(* IEC 61131-3 sources: STAR-PLC-Agent/results/raw/batch_fresh_20261114/PUB009/functional/attempt_0001, 1 file *)

(* ---- test_program.st ---- *)
PROGRAM PLC_PRG
VAR
 BenchStep : UDINT := 0;
 BenchCalls : UDINT := 0;
 BenchDone : BOOL := FALSE;
 BenchUut0 : FB_Task;
 BenchUut1 : FB_Task;
 BenchUut2 : FB_Task;
 BenchUut3 : FB_Task;
 BenchUut4 : FB_Task;
 BenchUut5 : FB_Task;
 BenchUut6 : FB_Task;
 TraceIn_cyclicExecution : ARRAY[0..454] OF BOOL;
 TraceIn_trigger : ARRAY[0..454] OF BOOL;
 TraceIn_value : ARRAY[0..454] OF LREAL;
 TraceIn_windowSize : ARRAY[0..454] OF INT;
 TraceIn_reset : ARRAY[0..454] OF BOOL;
 TraceOut_average : ARRAY[0..454] OF LREAL;
 TraceOut_windowSizeReached : ARRAY[0..454] OF BOOL;
 TraceOut_error : ARRAY[0..454] OF BOOL;
 TraceOut_status : ARRAY[0..454] OF WORD;
END_VAR

IF NOT BenchDone THEN
 CASE BenchStep OF
 0:
   BenchUut0.cyclicExecution := TRUE;
   BenchUut0.trigger := FALSE;
   BenchUut0.value := LREAL#3.0;
   BenchUut0.windowSize := INT#3;
   BenchUut0.reset := FALSE;
   TraceIn_cyclicExecution[0] := BenchUut0.cyclicExecution;
   TraceIn_trigger[0] := BenchUut0.trigger;
   TraceIn_value[0] := BenchUut0.value;
   TraceIn_windowSize[0] := BenchUut0.windowSize;
   TraceIn_reset[0] := BenchUut0.reset;
   BenchUut0();
   TraceOut_average[0] := BenchUut0.average;
   TraceOut_windowSizeReached[0] := BenchUut0.windowSizeReached;
   TraceOut_error[0] := BenchUut0.error;
   TraceOut_status[0] := BenchUut0.status;
   BenchCalls := BenchCalls + 1;
 1:
   BenchUut0.cyclicExecution := TRUE;
   BenchUut0.trigger := FALSE;
   BenchUut0.value := LREAL#6.0;
   BenchUut0.windowSize := INT#3;
   BenchUut0.reset := FALSE;
   TraceIn_cyclicExecution[1] := BenchUut0.cyclicExecution;
   TraceIn_trigger[1] := BenchUut0.trigger;
   TraceIn_value[1] := BenchUut0.value;
   TraceIn_windowSize[1] := BenchUut0.windowSize;
   TraceIn_reset[1] := BenchUut0.reset;
   BenchUut0();
   TraceOut_average[1] := BenchUut0.average;
   TraceOut_windowSizeReached[1] := BenchUut0.windowSizeReached;
   TraceOut_error[1] := BenchUut0.error;
   TraceOut_status[1] := BenchUut0.status;
   BenchCalls := BenchCalls + 1;
 2:
   BenchUut0.cyclicExecution := TRUE;
   BenchUut0.trigger := FALSE;
   BenchUut0.value := LREAL#9.0;
   BenchUut0.windowSize := INT#3;
   BenchUut0.reset := FALSE;
   TraceIn_cyclicExecution[2] := BenchUut0.cyclicExecution;
   TraceIn_trigger[2] := BenchUut0.trigger;
   TraceIn_value[2] := BenchUut0.value;
   TraceIn_windowSize[2] := BenchUut0.windowSize;
   TraceIn_reset[2] := BenchUut0.reset;
   BenchUut0();
   TraceOut_average[2] := BenchUut0.average;
   TraceOut_windowSizeReached[2] := BenchUut0.windowSizeReached;
   TraceOut_error[2] := BenchUut0.error;
   TraceOut_status[2] := BenchUut0.status;
   BenchCalls := BenchCalls + 1;
 3:
   BenchUut0.cyclicExecution := TRUE;
   BenchUut0.trigger := TRUE;
   BenchUut0.value := LREAL#12.0;
   BenchUut0.windowSize := INT#3;
   BenchUut0.reset := FALSE;
   TraceIn_cyclicExecution[3] := BenchUut0.cyclicExecution;
   TraceIn_trigger[3] := BenchUut0.trigger;
   TraceIn_value[3] := BenchUut0.value;
   TraceIn_windowSize[3] := BenchUut0.windowSize;
   TraceIn_reset[3] := BenchUut0.reset;
   BenchUut0();
   TraceOut_average[3] := BenchUut0.average;
   TraceOut_windowSizeReached[3] := BenchUut0.windowSizeReached;
   TraceOut_error[3] := BenchUut0.error;
   TraceOut_status[3] := BenchUut0.status;
   BenchCalls := BenchCalls + 1;
 4:
   BenchUut0.cyclicExecution := TRUE;
   BenchUut0.trigger := FALSE;
   BenchUut0.value := LREAL#99.0;
   BenchUut0.windowSize := INT#3;
   BenchUut0.reset := TRUE;
   TraceIn_cyclicExecution[4] := BenchUut0.cyclicExecution;
   TraceIn_trigger[4] := BenchUut0.trigger;
   TraceIn_value[4] := BenchUut0.value;
   TraceIn_windowSize[4] := BenchUut0.windowSize;
   TraceIn_reset[4] := BenchUut0.reset;
   BenchUut0();
   TraceOut_average[4] := BenchUut0.average;
   TraceOut_windowSizeReached[4] := BenchUut0.windowSizeReached;
   TraceOut_error[4] := BenchUut0.error;
   TraceOut_status[4] := BenchUut0.status;
   BenchCalls := BenchCalls + 1;
 5:
   BenchUut0.cyclicExecution := TRUE;
   BenchUut0.trigger := FALSE;
   BenchUut0.value := LREAL#-6.0;
   BenchUut0.windowSize := INT#3;
   BenchUut0.reset := FALSE;
   TraceIn_cyclicExecution[5] := BenchUut0.cyclicExecution;
   TraceIn_trigger[5] := BenchUut0.trigger;
   TraceIn_value[5] := BenchUut0.value;
   TraceIn_windowSize[5] := BenchUut0.windowSize;
   TraceIn_reset[5] := BenchUut0.reset;
   BenchUut0();
   TraceOut_average[5] := BenchUut0.average;
   TraceOut_windowSizeReached[5] := BenchUut0.windowSizeReached;
   TraceOut_error[5] := BenchUut0.error;
   TraceOut_status[5] := BenchUut0.status;
   BenchCalls := BenchCalls + 1;
 6:
   BenchUut1.cyclicExecution := FALSE;
   BenchUut1.trigger := TRUE;
   BenchUut1.value := LREAL#2.0;
   BenchUut1.windowSize := INT#3;
   BenchUut1.reset := FALSE;
   TraceIn_cyclicExecution[6] := BenchUut1.cyclicExecution;
   TraceIn_trigger[6] := BenchUut1.trigger;
   TraceIn_value[6] := BenchUut1.value;
   TraceIn_windowSize[6] := BenchUut1.windowSize;
   TraceIn_reset[6] := BenchUut1.reset;
   BenchUut1();
   TraceOut_average[6] := BenchUut1.average;
   TraceOut_windowSizeReached[6] := BenchUut1.windowSizeReached;
   TraceOut_error[6] := BenchUut1.error;
   TraceOut_status[6] := BenchUut1.status;
   BenchCalls := BenchCalls + 1;
 7:
   BenchUut1.cyclicExecution := FALSE;
   BenchUut1.trigger := TRUE;
   BenchUut1.value := LREAL#100.0;
   BenchUut1.windowSize := INT#3;
   BenchUut1.reset := FALSE;
   TraceIn_cyclicExecution[7] := BenchUut1.cyclicExecution;
   TraceIn_trigger[7] := BenchUut1.trigger;
   TraceIn_value[7] := BenchUut1.value;
   TraceIn_windowSize[7] := BenchUut1.windowSize;
   TraceIn_reset[7] := BenchUut1.reset;
   BenchUut1();
   TraceOut_average[7] := BenchUut1.average;
   TraceOut_windowSizeReached[7] := BenchUut1.windowSizeReached;
   TraceOut_error[7] := BenchUut1.error;
   TraceOut_status[7] := BenchUut1.status;
   BenchCalls := BenchCalls + 1;
 8:
   BenchUut1.cyclicExecution := FALSE;
   BenchUut1.trigger := FALSE;
   BenchUut1.value := LREAL#100.0;
   BenchUut1.windowSize := INT#3;
   BenchUut1.reset := FALSE;
   TraceIn_cyclicExecution[8] := BenchUut1.cyclicExecution;
   TraceIn_trigger[8] := BenchUut1.trigger;
   TraceIn_value[8] := BenchUut1.value;
   TraceIn_windowSize[8] := BenchUut1.windowSize;
   TraceIn_reset[8] := BenchUut1.reset;
   BenchUut1();
   TraceOut_average[8] := BenchUut1.average;
   TraceOut_windowSizeReached[8] := BenchUut1.windowSizeReached;
   TraceOut_error[8] := BenchUut1.error;
   TraceOut_status[8] := BenchUut1.status;
   BenchCalls := BenchCalls + 1;
 9:
   BenchUut1.cyclicExecution := FALSE;
   BenchUut1.trigger := TRUE;
   BenchUut1.value := LREAL#4.0;
   BenchUut1.windowSize := INT#3;
   BenchUut1.reset := FALSE;
   TraceIn_cyclicExecution[9] := BenchUut1.cyclicExecution;
   TraceIn_trigger[9] := BenchUut1.trigger;
   TraceIn_value[9] := BenchUut1.value;
   TraceIn_windowSize[9] := BenchUut1.windowSize;
   TraceIn_reset[9] := BenchUut1.reset;
   BenchUut1();
   TraceOut_average[9] := BenchUut1.average;
   TraceOut_windowSizeReached[9] := BenchUut1.windowSizeReached;
   TraceOut_error[9] := BenchUut1.error;
   TraceOut_status[9] := BenchUut1.status;
   BenchCalls := BenchCalls + 1;
 10:
   BenchUut1.cyclicExecution := TRUE;
   BenchUut1.trigger := FALSE;
   BenchUut1.value := LREAL#8.0;
   BenchUut1.windowSize := INT#1;
   BenchUut1.reset := FALSE;
   TraceIn_cyclicExecution[10] := BenchUut1.cyclicExecution;
   TraceIn_trigger[10] := BenchUut1.trigger;
   TraceIn_value[10] := BenchUut1.value;
   TraceIn_windowSize[10] := BenchUut1.windowSize;
   TraceIn_reset[10] := BenchUut1.reset;
   BenchUut1();
   TraceOut_average[10] := BenchUut1.average;
   TraceOut_windowSizeReached[10] := BenchUut1.windowSizeReached;
   TraceOut_error[10] := BenchUut1.error;
   TraceOut_status[10] := BenchUut1.status;
   BenchCalls := BenchCalls + 1;
 11:
   BenchUut1.cyclicExecution := FALSE;
   BenchUut1.trigger := FALSE;
   BenchUut1.value := LREAL#0.0;
   BenchUut1.windowSize := INT#0;
   BenchUut1.reset := FALSE;
   TraceIn_cyclicExecution[11] := BenchUut1.cyclicExecution;
   TraceIn_trigger[11] := BenchUut1.trigger;
   TraceIn_value[11] := BenchUut1.value;
   TraceIn_windowSize[11] := BenchUut1.windowSize;
   TraceIn_reset[11] := BenchUut1.reset;
   BenchUut1();
   TraceOut_average[11] := BenchUut1.average;
   TraceOut_windowSizeReached[11] := BenchUut1.windowSizeReached;
   TraceOut_error[11] := BenchUut1.error;
   TraceOut_status[11] := BenchUut1.status;
   BenchCalls := BenchCalls + 1;
 12:
   BenchUut1.cyclicExecution := FALSE;
   BenchUut1.trigger := FALSE;
   BenchUut1.value := LREAL#0.0;
   BenchUut1.windowSize := INT#101;
   BenchUut1.reset := FALSE;
   TraceIn_cyclicExecution[12] := BenchUut1.cyclicExecution;
   TraceIn_trigger[12] := BenchUut1.trigger;
   TraceIn_value[12] := BenchUut1.value;
   TraceIn_windowSize[12] := BenchUut1.windowSize;
   TraceIn_reset[12] := BenchUut1.reset;
   BenchUut1();
   TraceOut_average[12] := BenchUut1.average;
   TraceOut_windowSizeReached[12] := BenchUut1.windowSizeReached;
   TraceOut_error[12] := BenchUut1.error;
   TraceOut_status[12] := BenchUut1.status;
   BenchCalls := BenchCalls + 1;
 13:
   BenchUut1.cyclicExecution := FALSE;
   BenchUut1.trigger := FALSE;
   BenchUut1.value := LREAL#0.0;
   BenchUut1.windowSize := INT#1;
   BenchUut1.reset := TRUE;
   TraceIn_cyclicExecution[13] := BenchUut1.cyclicExecution;
   TraceIn_trigger[13] := BenchUut1.trigger;
   TraceIn_value[13] := BenchUut1.value;
   TraceIn_windowSize[13] := BenchUut1.windowSize;
   TraceIn_reset[13] := BenchUut1.reset;
   BenchUut1();
   TraceOut_average[13] := BenchUut1.average;
   TraceOut_windowSizeReached[13] := BenchUut1.windowSizeReached;
   TraceOut_error[13] := BenchUut1.error;
   TraceOut_status[13] := BenchUut1.status;
   BenchCalls := BenchCalls + 1;
 14:
   BenchUut1.cyclicExecution := FALSE;
   BenchUut1.trigger := TRUE;
   BenchUut1.value := LREAL#5.0;
   BenchUut1.windowSize := INT#1;
   BenchUut1.reset := FALSE;
   TraceIn_cyclicExecution[14] := BenchUut1.cyclicExecution;
   TraceIn_trigger[14] := BenchUut1.trigger;
   TraceIn_value[14] := BenchUut1.value;
   TraceIn_windowSize[14] := BenchUut1.windowSize;
   TraceIn_reset[14] := BenchUut1.reset;
   BenchUut1();
   TraceOut_average[14] := BenchUut1.average;
   TraceOut_windowSizeReached[14] := BenchUut1.windowSizeReached;
   TraceOut_error[14] := BenchUut1.error;
   TraceOut_status[14] := BenchUut1.status;
   BenchCalls := BenchCalls + 1;
 15:
   BenchUut2.cyclicExecution := FALSE;
   BenchUut2.trigger := TRUE;
   BenchUut2.value := LREAL#8.0;
   BenchUut2.windowSize := INT#2;
   BenchUut2.reset := FALSE;
   TraceIn_cyclicExecution[15] := BenchUut2.cyclicExecution;
   TraceIn_trigger[15] := BenchUut2.trigger;
   TraceIn_value[15] := BenchUut2.value;
   TraceIn_windowSize[15] := BenchUut2.windowSize;
   TraceIn_reset[15] := BenchUut2.reset;
   BenchUut2();
   TraceOut_average[15] := BenchUut2.average;
   TraceOut_windowSizeReached[15] := BenchUut2.windowSizeReached;
   TraceOut_error[15] := BenchUut2.error;
   TraceOut_status[15] := BenchUut2.status;
   BenchCalls := BenchCalls + 1;
 16:
   BenchUut2.cyclicExecution := FALSE;
   BenchUut2.trigger := FALSE;
   BenchUut2.value := LREAL#8.0;
   BenchUut2.windowSize := INT#2;
   BenchUut2.reset := FALSE;
   TraceIn_cyclicExecution[16] := BenchUut2.cyclicExecution;
   TraceIn_trigger[16] := BenchUut2.trigger;
   TraceIn_value[16] := BenchUut2.value;
   TraceIn_windowSize[16] := BenchUut2.windowSize;
   TraceIn_reset[16] := BenchUut2.reset;
   BenchUut2();
   TraceOut_average[16] := BenchUut2.average;
   TraceOut_windowSizeReached[16] := BenchUut2.windowSizeReached;
   TraceOut_error[16] := BenchUut2.error;
   TraceOut_status[16] := BenchUut2.status;
   BenchCalls := BenchCalls + 1;
 17:
   BenchUut2.cyclicExecution := FALSE;
   BenchUut2.trigger := TRUE;
   BenchUut2.value := LREAL#99.0;
   BenchUut2.windowSize := INT#0;
   BenchUut2.reset := FALSE;
   TraceIn_cyclicExecution[17] := BenchUut2.cyclicExecution;
   TraceIn_trigger[17] := BenchUut2.trigger;
   TraceIn_value[17] := BenchUut2.value;
   TraceIn_windowSize[17] := BenchUut2.windowSize;
   TraceIn_reset[17] := BenchUut2.reset;
   BenchUut2();
   TraceOut_average[17] := BenchUut2.average;
   TraceOut_windowSizeReached[17] := BenchUut2.windowSizeReached;
   TraceOut_error[17] := BenchUut2.error;
   TraceOut_status[17] := BenchUut2.status;
   BenchCalls := BenchCalls + 1;
 18:
   BenchUut2.cyclicExecution := FALSE;
   BenchUut2.trigger := TRUE;
   BenchUut2.value := LREAL#100.0;
   BenchUut2.windowSize := INT#2;
   BenchUut2.reset := FALSE;
   TraceIn_cyclicExecution[18] := BenchUut2.cyclicExecution;
   TraceIn_trigger[18] := BenchUut2.trigger;
   TraceIn_value[18] := BenchUut2.value;
   TraceIn_windowSize[18] := BenchUut2.windowSize;
   TraceIn_reset[18] := BenchUut2.reset;
   BenchUut2();
   TraceOut_average[18] := BenchUut2.average;
   TraceOut_windowSizeReached[18] := BenchUut2.windowSizeReached;
   TraceOut_error[18] := BenchUut2.error;
   TraceOut_status[18] := BenchUut2.status;
   BenchCalls := BenchCalls + 1;
 19:
   BenchUut2.cyclicExecution := FALSE;
   BenchUut2.trigger := FALSE;
   BenchUut2.value := LREAL#8.0;
   BenchUut2.windowSize := INT#2;
   BenchUut2.reset := FALSE;
   TraceIn_cyclicExecution[19] := BenchUut2.cyclicExecution;
   TraceIn_trigger[19] := BenchUut2.trigger;
   TraceIn_value[19] := BenchUut2.value;
   TraceIn_windowSize[19] := BenchUut2.windowSize;
   TraceIn_reset[19] := BenchUut2.reset;
   BenchUut2();
   TraceOut_average[19] := BenchUut2.average;
   TraceOut_windowSizeReached[19] := BenchUut2.windowSizeReached;
   TraceOut_error[19] := BenchUut2.error;
   TraceOut_status[19] := BenchUut2.status;
   BenchCalls := BenchCalls + 1;
 20:
   BenchUut2.cyclicExecution := FALSE;
   BenchUut2.trigger := TRUE;
   BenchUut2.value := LREAL#4.0;
   BenchUut2.windowSize := INT#2;
   BenchUut2.reset := FALSE;
   TraceIn_cyclicExecution[20] := BenchUut2.cyclicExecution;
   TraceIn_trigger[20] := BenchUut2.trigger;
   TraceIn_value[20] := BenchUut2.value;
   TraceIn_windowSize[20] := BenchUut2.windowSize;
   TraceIn_reset[20] := BenchUut2.reset;
   BenchUut2();
   TraceOut_average[20] := BenchUut2.average;
   TraceOut_windowSizeReached[20] := BenchUut2.windowSizeReached;
   TraceOut_error[20] := BenchUut2.error;
   TraceOut_status[20] := BenchUut2.status;
   BenchCalls := BenchCalls + 1;
 21:
   BenchUut2.cyclicExecution := FALSE;
   BenchUut2.trigger := FALSE;
   BenchUut2.value := LREAL#8.0;
   BenchUut2.windowSize := INT#3;
   BenchUut2.reset := FALSE;
   TraceIn_cyclicExecution[21] := BenchUut2.cyclicExecution;
   TraceIn_trigger[21] := BenchUut2.trigger;
   TraceIn_value[21] := BenchUut2.value;
   TraceIn_windowSize[21] := BenchUut2.windowSize;
   TraceIn_reset[21] := BenchUut2.reset;
   BenchUut2();
   TraceOut_average[21] := BenchUut2.average;
   TraceOut_windowSizeReached[21] := BenchUut2.windowSizeReached;
   TraceOut_error[21] := BenchUut2.error;
   TraceOut_status[21] := BenchUut2.status;
   BenchCalls := BenchCalls + 1;
 22:
   BenchUut3.cyclicExecution := TRUE;
   BenchUut3.trigger := FALSE;
   BenchUut3.value := LREAL#10.0;
   BenchUut3.windowSize := INT#2;
   BenchUut3.reset := FALSE;
   TraceIn_cyclicExecution[22] := BenchUut3.cyclicExecution;
   TraceIn_trigger[22] := BenchUut3.trigger;
   TraceIn_value[22] := BenchUut3.value;
   TraceIn_windowSize[22] := BenchUut3.windowSize;
   TraceIn_reset[22] := BenchUut3.reset;
   BenchUut3();
   TraceOut_average[22] := BenchUut3.average;
   TraceOut_windowSizeReached[22] := BenchUut3.windowSizeReached;
   TraceOut_error[22] := BenchUut3.error;
   TraceOut_status[22] := BenchUut3.status;
   BenchCalls := BenchCalls + 1;
 23:
   BenchUut3.cyclicExecution := TRUE;
   BenchUut3.trigger := FALSE;
   BenchUut3.value := LREAL#20.0;
   BenchUut3.windowSize := INT#2;
   BenchUut3.reset := FALSE;
   TraceIn_cyclicExecution[23] := BenchUut3.cyclicExecution;
   TraceIn_trigger[23] := BenchUut3.trigger;
   TraceIn_value[23] := BenchUut3.value;
   TraceIn_windowSize[23] := BenchUut3.windowSize;
   TraceIn_reset[23] := BenchUut3.reset;
   BenchUut3();
   TraceOut_average[23] := BenchUut3.average;
   TraceOut_windowSizeReached[23] := BenchUut3.windowSizeReached;
   TraceOut_error[23] := BenchUut3.error;
   TraceOut_status[23] := BenchUut3.status;
   BenchCalls := BenchCalls + 1;
 24:
   BenchUut3.cyclicExecution := TRUE;
   BenchUut3.trigger := FALSE;
   BenchUut3.value := LREAL#99.0;
   BenchUut3.windowSize := INT#0;
   BenchUut3.reset := TRUE;
   TraceIn_cyclicExecution[24] := BenchUut3.cyclicExecution;
   TraceIn_trigger[24] := BenchUut3.trigger;
   TraceIn_value[24] := BenchUut3.value;
   TraceIn_windowSize[24] := BenchUut3.windowSize;
   TraceIn_reset[24] := BenchUut3.reset;
   BenchUut3();
   TraceOut_average[24] := BenchUut3.average;
   TraceOut_windowSizeReached[24] := BenchUut3.windowSizeReached;
   TraceOut_error[24] := BenchUut3.error;
   TraceOut_status[24] := BenchUut3.status;
   BenchCalls := BenchCalls + 1;
 25:
   BenchUut3.cyclicExecution := TRUE;
   BenchUut3.trigger := FALSE;
   BenchUut3.value := LREAL#99.0;
   BenchUut3.windowSize := INT#-3;
   BenchUut3.reset := FALSE;
   TraceIn_cyclicExecution[25] := BenchUut3.cyclicExecution;
   TraceIn_trigger[25] := BenchUut3.trigger;
   TraceIn_value[25] := BenchUut3.value;
   TraceIn_windowSize[25] := BenchUut3.windowSize;
   TraceIn_reset[25] := BenchUut3.reset;
   BenchUut3();
   TraceOut_average[25] := BenchUut3.average;
   TraceOut_windowSizeReached[25] := BenchUut3.windowSizeReached;
   TraceOut_error[25] := BenchUut3.error;
   TraceOut_status[25] := BenchUut3.status;
   BenchCalls := BenchCalls + 1;
 26:
   BenchUut3.cyclicExecution := TRUE;
   BenchUut3.trigger := FALSE;
   BenchUut3.value := LREAL#30.0;
   BenchUut3.windowSize := INT#3;
   BenchUut3.reset := FALSE;
   TraceIn_cyclicExecution[26] := BenchUut3.cyclicExecution;
   TraceIn_trigger[26] := BenchUut3.trigger;
   TraceIn_value[26] := BenchUut3.value;
   TraceIn_windowSize[26] := BenchUut3.windowSize;
   TraceIn_reset[26] := BenchUut3.reset;
   BenchUut3();
   TraceOut_average[26] := BenchUut3.average;
   TraceOut_windowSizeReached[26] := BenchUut3.windowSizeReached;
   TraceOut_error[26] := BenchUut3.error;
   TraceOut_status[26] := BenchUut3.status;
   BenchCalls := BenchCalls + 1;
 27:
   BenchUut3.cyclicExecution := FALSE;
   BenchUut3.trigger := TRUE;
   BenchUut3.value := LREAL#60.0;
   BenchUut3.windowSize := INT#3;
   BenchUut3.reset := FALSE;
   TraceIn_cyclicExecution[27] := BenchUut3.cyclicExecution;
   TraceIn_trigger[27] := BenchUut3.trigger;
   TraceIn_value[27] := BenchUut3.value;
   TraceIn_windowSize[27] := BenchUut3.windowSize;
   TraceIn_reset[27] := BenchUut3.reset;
   BenchUut3();
   TraceOut_average[27] := BenchUut3.average;
   TraceOut_windowSizeReached[27] := BenchUut3.windowSizeReached;
   TraceOut_error[27] := BenchUut3.error;
   TraceOut_status[27] := BenchUut3.status;
   BenchCalls := BenchCalls + 1;
 28:
   BenchUut3.cyclicExecution := FALSE;
   BenchUut3.trigger := TRUE;
   BenchUut3.value := LREAL#90.0;
   BenchUut3.windowSize := INT#3;
   BenchUut3.reset := FALSE;
   TraceIn_cyclicExecution[28] := BenchUut3.cyclicExecution;
   TraceIn_trigger[28] := BenchUut3.trigger;
   TraceIn_value[28] := BenchUut3.value;
   TraceIn_windowSize[28] := BenchUut3.windowSize;
   TraceIn_reset[28] := BenchUut3.reset;
   BenchUut3();
   TraceOut_average[28] := BenchUut3.average;
   TraceOut_windowSizeReached[28] := BenchUut3.windowSizeReached;
   TraceOut_error[28] := BenchUut3.error;
   TraceOut_status[28] := BenchUut3.status;
   BenchCalls := BenchCalls + 1;
 29:
   BenchUut3.cyclicExecution := TRUE;
   BenchUut3.trigger := FALSE;
   BenchUut3.value := LREAL#90.0;
   BenchUut3.windowSize := INT#3;
   BenchUut3.reset := FALSE;
   TraceIn_cyclicExecution[29] := BenchUut3.cyclicExecution;
   TraceIn_trigger[29] := BenchUut3.trigger;
   TraceIn_value[29] := BenchUut3.value;
   TraceIn_windowSize[29] := BenchUut3.windowSize;
   TraceIn_reset[29] := BenchUut3.reset;
   BenchUut3();
   TraceOut_average[29] := BenchUut3.average;
   TraceOut_windowSizeReached[29] := BenchUut3.windowSizeReached;
   TraceOut_error[29] := BenchUut3.error;
   TraceOut_status[29] := BenchUut3.status;
   BenchCalls := BenchCalls + 1;
 30:
   BenchUut3.cyclicExecution := TRUE;
   BenchUut3.trigger := FALSE;
   BenchUut3.value := LREAL#1.0;
   BenchUut3.windowSize := INT#100;
   BenchUut3.reset := FALSE;
   TraceIn_cyclicExecution[30] := BenchUut3.cyclicExecution;
   TraceIn_trigger[30] := BenchUut3.trigger;
   TraceIn_value[30] := BenchUut3.value;
   TraceIn_windowSize[30] := BenchUut3.windowSize;
   TraceIn_reset[30] := BenchUut3.reset;
   BenchUut3();
   TraceOut_average[30] := BenchUut3.average;
   TraceOut_windowSizeReached[30] := BenchUut3.windowSizeReached;
   TraceOut_error[30] := BenchUut3.error;
   TraceOut_status[30] := BenchUut3.status;
   BenchCalls := BenchCalls + 1;
 31:
   BenchUut3.cyclicExecution := TRUE;
   BenchUut3.trigger := FALSE;
   BenchUut3.value := LREAL#2.0;
   BenchUut3.windowSize := INT#100;
   BenchUut3.reset := FALSE;
   TraceIn_cyclicExecution[31] := BenchUut3.cyclicExecution;
   TraceIn_trigger[31] := BenchUut3.trigger;
   TraceIn_value[31] := BenchUut3.value;
   TraceIn_windowSize[31] := BenchUut3.windowSize;
   TraceIn_reset[31] := BenchUut3.reset;
   BenchUut3();
   TraceOut_average[31] := BenchUut3.average;
   TraceOut_windowSizeReached[31] := BenchUut3.windowSizeReached;
   TraceOut_error[31] := BenchUut3.error;
   TraceOut_status[31] := BenchUut3.status;
   BenchCalls := BenchCalls + 1;
 32:
   BenchUut3.cyclicExecution := TRUE;
   BenchUut3.trigger := FALSE;
   BenchUut3.value := LREAL#3.0;
   BenchUut3.windowSize := INT#100;
   BenchUut3.reset := FALSE;
   TraceIn_cyclicExecution[32] := BenchUut3.cyclicExecution;
   TraceIn_trigger[32] := BenchUut3.trigger;
   TraceIn_value[32] := BenchUut3.value;
   TraceIn_windowSize[32] := BenchUut3.windowSize;
   TraceIn_reset[32] := BenchUut3.reset;
   BenchUut3();
   TraceOut_average[32] := BenchUut3.average;
   TraceOut_windowSizeReached[32] := BenchUut3.windowSizeReached;
   TraceOut_error[32] := BenchUut3.error;
   TraceOut_status[32] := BenchUut3.status;
   BenchCalls := BenchCalls + 1;
 33:
   BenchUut3.cyclicExecution := TRUE;
   BenchUut3.trigger := FALSE;
   BenchUut3.value := LREAL#4.0;
   BenchUut3.windowSize := INT#100;
   BenchUut3.reset := FALSE;
   TraceIn_cyclicExecution[33] := BenchUut3.cyclicExecution;
   TraceIn_trigger[33] := BenchUut3.trigger;
   TraceIn_value[33] := BenchUut3.value;
   TraceIn_windowSize[33] := BenchUut3.windowSize;
   TraceIn_reset[33] := BenchUut3.reset;
   BenchUut3();
   TraceOut_average[33] := BenchUut3.average;
   TraceOut_windowSizeReached[33] := BenchUut3.windowSizeReached;
   TraceOut_error[33] := BenchUut3.error;
   TraceOut_status[33] := BenchUut3.status;
   BenchCalls := BenchCalls + 1;
 34:
   BenchUut3.cyclicExecution := TRUE;
   BenchUut3.trigger := FALSE;
   BenchUut3.value := LREAL#5.0;
   BenchUut3.windowSize := INT#100;
   BenchUut3.reset := FALSE;
   TraceIn_cyclicExecution[34] := BenchUut3.cyclicExecution;
   TraceIn_trigger[34] := BenchUut3.trigger;
   TraceIn_value[34] := BenchUut3.value;
   TraceIn_windowSize[34] := BenchUut3.windowSize;
   TraceIn_reset[34] := BenchUut3.reset;
   BenchUut3();
   TraceOut_average[34] := BenchUut3.average;
   TraceOut_windowSizeReached[34] := BenchUut3.windowSizeReached;
   TraceOut_error[34] := BenchUut3.error;
   TraceOut_status[34] := BenchUut3.status;
   BenchCalls := BenchCalls + 1;
 35:
   BenchUut3.cyclicExecution := TRUE;
   BenchUut3.trigger := FALSE;
   BenchUut3.value := LREAL#6.0;
   BenchUut3.windowSize := INT#100;
   BenchUut3.reset := FALSE;
   TraceIn_cyclicExecution[35] := BenchUut3.cyclicExecution;
   TraceIn_trigger[35] := BenchUut3.trigger;
   TraceIn_value[35] := BenchUut3.value;
   TraceIn_windowSize[35] := BenchUut3.windowSize;
   TraceIn_reset[35] := BenchUut3.reset;
   BenchUut3();
   TraceOut_average[35] := BenchUut3.average;
   TraceOut_windowSizeReached[35] := BenchUut3.windowSizeReached;
   TraceOut_error[35] := BenchUut3.error;
   TraceOut_status[35] := BenchUut3.status;
   BenchCalls := BenchCalls + 1;
 36:
   BenchUut3.cyclicExecution := TRUE;
   BenchUut3.trigger := FALSE;
   BenchUut3.value := LREAL#7.0;
   BenchUut3.windowSize := INT#100;
   BenchUut3.reset := FALSE;
   TraceIn_cyclicExecution[36] := BenchUut3.cyclicExecution;
   TraceIn_trigger[36] := BenchUut3.trigger;
   TraceIn_value[36] := BenchUut3.value;
   TraceIn_windowSize[36] := BenchUut3.windowSize;
   TraceIn_reset[36] := BenchUut3.reset;
   BenchUut3();
   TraceOut_average[36] := BenchUut3.average;
   TraceOut_windowSizeReached[36] := BenchUut3.windowSizeReached;
   TraceOut_error[36] := BenchUut3.error;
   TraceOut_status[36] := BenchUut3.status;
   BenchCalls := BenchCalls + 1;
 37:
   BenchUut3.cyclicExecution := TRUE;
   BenchUut3.trigger := FALSE;
   BenchUut3.value := LREAL#8.0;
   BenchUut3.windowSize := INT#100;
   BenchUut3.reset := FALSE;
   TraceIn_cyclicExecution[37] := BenchUut3.cyclicExecution;
   TraceIn_trigger[37] := BenchUut3.trigger;
   TraceIn_value[37] := BenchUut3.value;
   TraceIn_windowSize[37] := BenchUut3.windowSize;
   TraceIn_reset[37] := BenchUut3.reset;
   BenchUut3();
   TraceOut_average[37] := BenchUut3.average;
   TraceOut_windowSizeReached[37] := BenchUut3.windowSizeReached;
   TraceOut_error[37] := BenchUut3.error;
   TraceOut_status[37] := BenchUut3.status;
   BenchCalls := BenchCalls + 1;
 38:
   BenchUut3.cyclicExecution := TRUE;
   BenchUut3.trigger := FALSE;
   BenchUut3.value := LREAL#9.0;
   BenchUut3.windowSize := INT#100;
   BenchUut3.reset := FALSE;
   TraceIn_cyclicExecution[38] := BenchUut3.cyclicExecution;
   TraceIn_trigger[38] := BenchUut3.trigger;
   TraceIn_value[38] := BenchUut3.value;
   TraceIn_windowSize[38] := BenchUut3.windowSize;
   TraceIn_reset[38] := BenchUut3.reset;
   BenchUut3();
   TraceOut_average[38] := BenchUut3.average;
   TraceOut_windowSizeReached[38] := BenchUut3.windowSizeReached;
   TraceOut_error[38] := BenchUut3.error;
   TraceOut_status[38] := BenchUut3.status;
   BenchCalls := BenchCalls + 1;
 39:
   BenchUut3.cyclicExecution := TRUE;
   BenchUut3.trigger := FALSE;
   BenchUut3.value := LREAL#10.0;
   BenchUut3.windowSize := INT#100;
   BenchUut3.reset := FALSE;
   TraceIn_cyclicExecution[39] := BenchUut3.cyclicExecution;
   TraceIn_trigger[39] := BenchUut3.trigger;
   TraceIn_value[39] := BenchUut3.value;
   TraceIn_windowSize[39] := BenchUut3.windowSize;
   TraceIn_reset[39] := BenchUut3.reset;
   BenchUut3();
   TraceOut_average[39] := BenchUut3.average;
   TraceOut_windowSizeReached[39] := BenchUut3.windowSizeReached;
   TraceOut_error[39] := BenchUut3.error;
   TraceOut_status[39] := BenchUut3.status;
   BenchCalls := BenchCalls + 1;
 40:
   BenchUut3.cyclicExecution := TRUE;
   BenchUut3.trigger := FALSE;
   BenchUut3.value := LREAL#11.0;
   BenchUut3.windowSize := INT#100;
   BenchUut3.reset := FALSE;
   TraceIn_cyclicExecution[40] := BenchUut3.cyclicExecution;
   TraceIn_trigger[40] := BenchUut3.trigger;
   TraceIn_value[40] := BenchUut3.value;
   TraceIn_windowSize[40] := BenchUut3.windowSize;
   TraceIn_reset[40] := BenchUut3.reset;
   BenchUut3();
   TraceOut_average[40] := BenchUut3.average;
   TraceOut_windowSizeReached[40] := BenchUut3.windowSizeReached;
   TraceOut_error[40] := BenchUut3.error;
   TraceOut_status[40] := BenchUut3.status;
   BenchCalls := BenchCalls + 1;
 41:
   BenchUut3.cyclicExecution := TRUE;
   BenchUut3.trigger := FALSE;
   BenchUut3.value := LREAL#12.0;
   BenchUut3.windowSize := INT#100;
   BenchUut3.reset := FALSE;
   TraceIn_cyclicExecution[41] := BenchUut3.cyclicExecution;
   TraceIn_trigger[41] := BenchUut3.trigger;
   TraceIn_value[41] := BenchUut3.value;
   TraceIn_windowSize[41] := BenchUut3.windowSize;
   TraceIn_reset[41] := BenchUut3.reset;
   BenchUut3();
   TraceOut_average[41] := BenchUut3.average;
   TraceOut_windowSizeReached[41] := BenchUut3.windowSizeReached;
   TraceOut_error[41] := BenchUut3.error;
   TraceOut_status[41] := BenchUut3.status;
   BenchCalls := BenchCalls + 1;
 42:
   BenchUut3.cyclicExecution := TRUE;
   BenchUut3.trigger := FALSE;
   BenchUut3.value := LREAL#13.0;
   BenchUut3.windowSize := INT#100;
   BenchUut3.reset := FALSE;
   TraceIn_cyclicExecution[42] := BenchUut3.cyclicExecution;
   TraceIn_trigger[42] := BenchUut3.trigger;
   TraceIn_value[42] := BenchUut3.value;
   TraceIn_windowSize[42] := BenchUut3.windowSize;
   TraceIn_reset[42] := BenchUut3.reset;
   BenchUut3();
   TraceOut_average[42] := BenchUut3.average;
   TraceOut_windowSizeReached[42] := BenchUut3.windowSizeReached;
   TraceOut_error[42] := BenchUut3.error;
   TraceOut_status[42] := BenchUut3.status;
   BenchCalls := BenchCalls + 1;
 43:
   BenchUut3.cyclicExecution := TRUE;
   BenchUut3.trigger := FALSE;
   BenchUut3.value := LREAL#14.0;
   BenchUut3.windowSize := INT#100;
   BenchUut3.reset := FALSE;
   TraceIn_cyclicExecution[43] := BenchUut3.cyclicExecution;
   TraceIn_trigger[43] := BenchUut3.trigger;
   TraceIn_value[43] := BenchUut3.value;
   TraceIn_windowSize[43] := BenchUut3.windowSize;
   TraceIn_reset[43] := BenchUut3.reset;
   BenchUut3();
   TraceOut_average[43] := BenchUut3.average;
   TraceOut_windowSizeReached[43] := BenchUut3.windowSizeReached;
   TraceOut_error[43] := BenchUut3.error;
   TraceOut_status[43] := BenchUut3.status;
   BenchCalls := BenchCalls + 1;
 44:
   BenchUut3.cyclicExecution := TRUE;
   BenchUut3.trigger := FALSE;
   BenchUut3.value := LREAL#15.0;
   BenchUut3.windowSize := INT#100;
   BenchUut3.reset := FALSE;
   TraceIn_cyclicExecution[44] := BenchUut3.cyclicExecution;
   TraceIn_trigger[44] := BenchUut3.trigger;
   TraceIn_value[44] := BenchUut3.value;
   TraceIn_windowSize[44] := BenchUut3.windowSize;
   TraceIn_reset[44] := BenchUut3.reset;
   BenchUut3();
   TraceOut_average[44] := BenchUut3.average;
   TraceOut_windowSizeReached[44] := BenchUut3.windowSizeReached;
   TraceOut_error[44] := BenchUut3.error;
   TraceOut_status[44] := BenchUut3.status;
   BenchCalls := BenchCalls + 1;
 45:
   BenchUut3.cyclicExecution := TRUE;
   BenchUut3.trigger := FALSE;
   BenchUut3.value := LREAL#16.0;
   BenchUut3.windowSize := INT#100;
   BenchUut3.reset := FALSE;
   TraceIn_cyclicExecution[45] := BenchUut3.cyclicExecution;
   TraceIn_trigger[45] := BenchUut3.trigger;
   TraceIn_value[45] := BenchUut3.value;
   TraceIn_windowSize[45] := BenchUut3.windowSize;
   TraceIn_reset[45] := BenchUut3.reset;
   BenchUut3();
   TraceOut_average[45] := BenchUut3.average;
   TraceOut_windowSizeReached[45] := BenchUut3.windowSizeReached;
   TraceOut_error[45] := BenchUut3.error;
   TraceOut_status[45] := BenchUut3.status;
   BenchCalls := BenchCalls + 1;
 46:
   BenchUut3.cyclicExecution := TRUE;
   BenchUut3.trigger := FALSE;
   BenchUut3.value := LREAL#17.0;
   BenchUut3.windowSize := INT#100;
   BenchUut3.reset := FALSE;
   TraceIn_cyclicExecution[46] := BenchUut3.cyclicExecution;
   TraceIn_trigger[46] := BenchUut3.trigger;
   TraceIn_value[46] := BenchUut3.value;
   TraceIn_windowSize[46] := BenchUut3.windowSize;
   TraceIn_reset[46] := BenchUut3.reset;
   BenchUut3();
   TraceOut_average[46] := BenchUut3.average;
   TraceOut_windowSizeReached[46] := BenchUut3.windowSizeReached;
   TraceOut_error[46] := BenchUut3.error;
   TraceOut_status[46] := BenchUut3.status;
   BenchCalls := BenchCalls + 1;
 47:
   BenchUut3.cyclicExecution := TRUE;
   BenchUut3.trigger := FALSE;
   BenchUut3.value := LREAL#18.0;
   BenchUut3.windowSize := INT#100;
   BenchUut3.reset := FALSE;
   TraceIn_cyclicExecution[47] := BenchUut3.cyclicExecution;
   TraceIn_trigger[47] := BenchUut3.trigger;
   TraceIn_value[47] := BenchUut3.value;
   TraceIn_windowSize[47] := BenchUut3.windowSize;
   TraceIn_reset[47] := BenchUut3.reset;
   BenchUut3();
   TraceOut_average[47] := BenchUut3.average;
   TraceOut_windowSizeReached[47] := BenchUut3.windowSizeReached;
   TraceOut_error[47] := BenchUut3.error;
   TraceOut_status[47] := BenchUut3.status;
   BenchCalls := BenchCalls + 1;
 48:
   BenchUut3.cyclicExecution := TRUE;
   BenchUut3.trigger := FALSE;
   BenchUut3.value := LREAL#19.0;
   BenchUut3.windowSize := INT#100;
   BenchUut3.reset := FALSE;
   TraceIn_cyclicExecution[48] := BenchUut3.cyclicExecution;
   TraceIn_trigger[48] := BenchUut3.trigger;
   TraceIn_value[48] := BenchUut3.value;
   TraceIn_windowSize[48] := BenchUut3.windowSize;
   TraceIn_reset[48] := BenchUut3.reset;
   BenchUut3();
   TraceOut_average[48] := BenchUut3.average;
   TraceOut_windowSizeReached[48] := BenchUut3.windowSizeReached;
   TraceOut_error[48] := BenchUut3.error;
   TraceOut_status[48] := BenchUut3.status;
   BenchCalls := BenchCalls + 1;
 49:
   BenchUut3.cyclicExecution := TRUE;
   BenchUut3.trigger := FALSE;
   BenchUut3.value := LREAL#20.0;
   BenchUut3.windowSize := INT#100;
   BenchUut3.reset := FALSE;
   TraceIn_cyclicExecution[49] := BenchUut3.cyclicExecution;
   TraceIn_trigger[49] := BenchUut3.trigger;
   TraceIn_value[49] := BenchUut3.value;
   TraceIn_windowSize[49] := BenchUut3.windowSize;
   TraceIn_reset[49] := BenchUut3.reset;
   BenchUut3();
   TraceOut_average[49] := BenchUut3.average;
   TraceOut_windowSizeReached[49] := BenchUut3.windowSizeReached;
   TraceOut_error[49] := BenchUut3.error;
   TraceOut_status[49] := BenchUut3.status;
   BenchCalls := BenchCalls + 1;
 50:
   BenchUut3.cyclicExecution := TRUE;
   BenchUut3.trigger := FALSE;
   BenchUut3.value := LREAL#21.0;
   BenchUut3.windowSize := INT#100;
   BenchUut3.reset := FALSE;
   TraceIn_cyclicExecution[50] := BenchUut3.cyclicExecution;
   TraceIn_trigger[50] := BenchUut3.trigger;
   TraceIn_value[50] := BenchUut3.value;
   TraceIn_windowSize[50] := BenchUut3.windowSize;
   TraceIn_reset[50] := BenchUut3.reset;
   BenchUut3();
   TraceOut_average[50] := BenchUut3.average;
   TraceOut_windowSizeReached[50] := BenchUut3.windowSizeReached;
   TraceOut_error[50] := BenchUut3.error;
   TraceOut_status[50] := BenchUut3.status;
   BenchCalls := BenchCalls + 1;
 51:
   BenchUut3.cyclicExecution := TRUE;
   BenchUut3.trigger := FALSE;
   BenchUut3.value := LREAL#22.0;
   BenchUut3.windowSize := INT#100;
   BenchUut3.reset := FALSE;
   TraceIn_cyclicExecution[51] := BenchUut3.cyclicExecution;
   TraceIn_trigger[51] := BenchUut3.trigger;
   TraceIn_value[51] := BenchUut3.value;
   TraceIn_windowSize[51] := BenchUut3.windowSize;
   TraceIn_reset[51] := BenchUut3.reset;
   BenchUut3();
   TraceOut_average[51] := BenchUut3.average;
   TraceOut_windowSizeReached[51] := BenchUut3.windowSizeReached;
   TraceOut_error[51] := BenchUut3.error;
   TraceOut_status[51] := BenchUut3.status;
   BenchCalls := BenchCalls + 1;
 52:
   BenchUut3.cyclicExecution := TRUE;
   BenchUut3.trigger := FALSE;
   BenchUut3.value := LREAL#23.0;
   BenchUut3.windowSize := INT#100;
   BenchUut3.reset := FALSE;
   TraceIn_cyclicExecution[52] := BenchUut3.cyclicExecution;
   TraceIn_trigger[52] := BenchUut3.trigger;
   TraceIn_value[52] := BenchUut3.value;
   TraceIn_windowSize[52] := BenchUut3.windowSize;
   TraceIn_reset[52] := BenchUut3.reset;
   BenchUut3();
   TraceOut_average[52] := BenchUut3.average;
   TraceOut_windowSizeReached[52] := BenchUut3.windowSizeReached;
   TraceOut_error[52] := BenchUut3.error;
   TraceOut_status[52] := BenchUut3.status;
   BenchCalls := BenchCalls + 1;
 53:
   BenchUut3.cyclicExecution := TRUE;
   BenchUut3.trigger := FALSE;
   BenchUut3.value := LREAL#24.0;
   BenchUut3.windowSize := INT#100;
   BenchUut3.reset := FALSE;
   TraceIn_cyclicExecution[53] := BenchUut3.cyclicExecution;
   TraceIn_trigger[53] := BenchUut3.trigger;
   TraceIn_value[53] := BenchUut3.value;
   TraceIn_windowSize[53] := BenchUut3.windowSize;
   TraceIn_reset[53] := BenchUut3.reset;
   BenchUut3();
   TraceOut_average[53] := BenchUut3.average;
   TraceOut_windowSizeReached[53] := BenchUut3.windowSizeReached;
   TraceOut_error[53] := BenchUut3.error;
   TraceOut_status[53] := BenchUut3.status;
   BenchCalls := BenchCalls + 1;
 54:
   BenchUut3.cyclicExecution := TRUE;
   BenchUut3.trigger := FALSE;
   BenchUut3.value := LREAL#25.0;
   BenchUut3.windowSize := INT#100;
   BenchUut3.reset := FALSE;
   TraceIn_cyclicExecution[54] := BenchUut3.cyclicExecution;
   TraceIn_trigger[54] := BenchUut3.trigger;
   TraceIn_value[54] := BenchUut3.value;
   TraceIn_windowSize[54] := BenchUut3.windowSize;
   TraceIn_reset[54] := BenchUut3.reset;
   BenchUut3();
   TraceOut_average[54] := BenchUut3.average;
   TraceOut_windowSizeReached[54] := BenchUut3.windowSizeReached;
   TraceOut_error[54] := BenchUut3.error;
   TraceOut_status[54] := BenchUut3.status;
   BenchCalls := BenchCalls + 1;
 55:
   BenchUut3.cyclicExecution := TRUE;
   BenchUut3.trigger := FALSE;
   BenchUut3.value := LREAL#26.0;
   BenchUut3.windowSize := INT#100;
   BenchUut3.reset := FALSE;
   TraceIn_cyclicExecution[55] := BenchUut3.cyclicExecution;
   TraceIn_trigger[55] := BenchUut3.trigger;
   TraceIn_value[55] := BenchUut3.value;
   TraceIn_windowSize[55] := BenchUut3.windowSize;
   TraceIn_reset[55] := BenchUut3.reset;
   BenchUut3();
   TraceOut_average[55] := BenchUut3.average;
   TraceOut_windowSizeReached[55] := BenchUut3.windowSizeReached;
   TraceOut_error[55] := BenchUut3.error;
   TraceOut_status[55] := BenchUut3.status;
   BenchCalls := BenchCalls + 1;
 56:
   BenchUut3.cyclicExecution := TRUE;
   BenchUut3.trigger := FALSE;
   BenchUut3.value := LREAL#27.0;
   BenchUut3.windowSize := INT#100;
   BenchUut3.reset := FALSE;
   TraceIn_cyclicExecution[56] := BenchUut3.cyclicExecution;
   TraceIn_trigger[56] := BenchUut3.trigger;
   TraceIn_value[56] := BenchUut3.value;
   TraceIn_windowSize[56] := BenchUut3.windowSize;
   TraceIn_reset[56] := BenchUut3.reset;
   BenchUut3();
   TraceOut_average[56] := BenchUut3.average;
   TraceOut_windowSizeReached[56] := BenchUut3.windowSizeReached;
   TraceOut_error[56] := BenchUut3.error;
   TraceOut_status[56] := BenchUut3.status;
   BenchCalls := BenchCalls + 1;
 57:
   BenchUut3.cyclicExecution := TRUE;
   BenchUut3.trigger := FALSE;
   BenchUut3.value := LREAL#28.0;
   BenchUut3.windowSize := INT#100;
   BenchUut3.reset := FALSE;
   TraceIn_cyclicExecution[57] := BenchUut3.cyclicExecution;
   TraceIn_trigger[57] := BenchUut3.trigger;
   TraceIn_value[57] := BenchUut3.value;
   TraceIn_windowSize[57] := BenchUut3.windowSize;
   TraceIn_reset[57] := BenchUut3.reset;
   BenchUut3();
   TraceOut_average[57] := BenchUut3.average;
   TraceOut_windowSizeReached[57] := BenchUut3.windowSizeReached;
   TraceOut_error[57] := BenchUut3.error;
   TraceOut_status[57] := BenchUut3.status;
   BenchCalls := BenchCalls + 1;
 58:
   BenchUut3.cyclicExecution := TRUE;
   BenchUut3.trigger := FALSE;
   BenchUut3.value := LREAL#29.0;
   BenchUut3.windowSize := INT#100;
   BenchUut3.reset := FALSE;
   TraceIn_cyclicExecution[58] := BenchUut3.cyclicExecution;
   TraceIn_trigger[58] := BenchUut3.trigger;
   TraceIn_value[58] := BenchUut3.value;
   TraceIn_windowSize[58] := BenchUut3.windowSize;
   TraceIn_reset[58] := BenchUut3.reset;
   BenchUut3();
   TraceOut_average[58] := BenchUut3.average;
   TraceOut_windowSizeReached[58] := BenchUut3.windowSizeReached;
   TraceOut_error[58] := BenchUut3.error;
   TraceOut_status[58] := BenchUut3.status;
   BenchCalls := BenchCalls + 1;
 59:
   BenchUut3.cyclicExecution := TRUE;
   BenchUut3.trigger := FALSE;
   BenchUut3.value := LREAL#30.0;
   BenchUut3.windowSize := INT#100;
   BenchUut3.reset := FALSE;
   TraceIn_cyclicExecution[59] := BenchUut3.cyclicExecution;
   TraceIn_trigger[59] := BenchUut3.trigger;
   TraceIn_value[59] := BenchUut3.value;
   TraceIn_windowSize[59] := BenchUut3.windowSize;
   TraceIn_reset[59] := BenchUut3.reset;
   BenchUut3();
   TraceOut_average[59] := BenchUut3.average;
   TraceOut_windowSizeReached[59] := BenchUut3.windowSizeReached;
   TraceOut_error[59] := BenchUut3.error;
   TraceOut_status[59] := BenchUut3.status;
   BenchCalls := BenchCalls + 1;
 60:
   BenchUut3.cyclicExecution := TRUE;
   BenchUut3.trigger := FALSE;
   BenchUut3.value := LREAL#31.0;
   BenchUut3.windowSize := INT#100;
   BenchUut3.reset := FALSE;
   TraceIn_cyclicExecution[60] := BenchUut3.cyclicExecution;
   TraceIn_trigger[60] := BenchUut3.trigger;
   TraceIn_value[60] := BenchUut3.value;
   TraceIn_windowSize[60] := BenchUut3.windowSize;
   TraceIn_reset[60] := BenchUut3.reset;
   BenchUut3();
   TraceOut_average[60] := BenchUut3.average;
   TraceOut_windowSizeReached[60] := BenchUut3.windowSizeReached;
   TraceOut_error[60] := BenchUut3.error;
   TraceOut_status[60] := BenchUut3.status;
   BenchCalls := BenchCalls + 1;
 61:
   BenchUut3.cyclicExecution := TRUE;
   BenchUut3.trigger := FALSE;
   BenchUut3.value := LREAL#32.0;
   BenchUut3.windowSize := INT#100;
   BenchUut3.reset := FALSE;
   TraceIn_cyclicExecution[61] := BenchUut3.cyclicExecution;
   TraceIn_trigger[61] := BenchUut3.trigger;
   TraceIn_value[61] := BenchUut3.value;
   TraceIn_windowSize[61] := BenchUut3.windowSize;
   TraceIn_reset[61] := BenchUut3.reset;
   BenchUut3();
   TraceOut_average[61] := BenchUut3.average;
   TraceOut_windowSizeReached[61] := BenchUut3.windowSizeReached;
   TraceOut_error[61] := BenchUut3.error;
   TraceOut_status[61] := BenchUut3.status;
   BenchCalls := BenchCalls + 1;
 62:
   BenchUut3.cyclicExecution := TRUE;
   BenchUut3.trigger := FALSE;
   BenchUut3.value := LREAL#33.0;
   BenchUut3.windowSize := INT#100;
   BenchUut3.reset := FALSE;
   TraceIn_cyclicExecution[62] := BenchUut3.cyclicExecution;
   TraceIn_trigger[62] := BenchUut3.trigger;
   TraceIn_value[62] := BenchUut3.value;
   TraceIn_windowSize[62] := BenchUut3.windowSize;
   TraceIn_reset[62] := BenchUut3.reset;
   BenchUut3();
   TraceOut_average[62] := BenchUut3.average;
   TraceOut_windowSizeReached[62] := BenchUut3.windowSizeReached;
   TraceOut_error[62] := BenchUut3.error;
   TraceOut_status[62] := BenchUut3.status;
   BenchCalls := BenchCalls + 1;
 63:
   BenchUut3.cyclicExecution := TRUE;
   BenchUut3.trigger := FALSE;
   BenchUut3.value := LREAL#34.0;
   BenchUut3.windowSize := INT#100;
   BenchUut3.reset := FALSE;
   TraceIn_cyclicExecution[63] := BenchUut3.cyclicExecution;
   TraceIn_trigger[63] := BenchUut3.trigger;
   TraceIn_value[63] := BenchUut3.value;
   TraceIn_windowSize[63] := BenchUut3.windowSize;
   TraceIn_reset[63] := BenchUut3.reset;
   BenchUut3();
   TraceOut_average[63] := BenchUut3.average;
   TraceOut_windowSizeReached[63] := BenchUut3.windowSizeReached;
   TraceOut_error[63] := BenchUut3.error;
   TraceOut_status[63] := BenchUut3.status;
   BenchCalls := BenchCalls + 1;
 64:
   BenchUut3.cyclicExecution := TRUE;
   BenchUut3.trigger := FALSE;
   BenchUut3.value := LREAL#35.0;
   BenchUut3.windowSize := INT#100;
   BenchUut3.reset := FALSE;
   TraceIn_cyclicExecution[64] := BenchUut3.cyclicExecution;
   TraceIn_trigger[64] := BenchUut3.trigger;
   TraceIn_value[64] := BenchUut3.value;
   TraceIn_windowSize[64] := BenchUut3.windowSize;
   TraceIn_reset[64] := BenchUut3.reset;
   BenchUut3();
   TraceOut_average[64] := BenchUut3.average;
   TraceOut_windowSizeReached[64] := BenchUut3.windowSizeReached;
   TraceOut_error[64] := BenchUut3.error;
   TraceOut_status[64] := BenchUut3.status;
   BenchCalls := BenchCalls + 1;
 65:
   BenchUut3.cyclicExecution := TRUE;
   BenchUut3.trigger := FALSE;
   BenchUut3.value := LREAL#36.0;
   BenchUut3.windowSize := INT#100;
   BenchUut3.reset := FALSE;
   TraceIn_cyclicExecution[65] := BenchUut3.cyclicExecution;
   TraceIn_trigger[65] := BenchUut3.trigger;
   TraceIn_value[65] := BenchUut3.value;
   TraceIn_windowSize[65] := BenchUut3.windowSize;
   TraceIn_reset[65] := BenchUut3.reset;
   BenchUut3();
   TraceOut_average[65] := BenchUut3.average;
   TraceOut_windowSizeReached[65] := BenchUut3.windowSizeReached;
   TraceOut_error[65] := BenchUut3.error;
   TraceOut_status[65] := BenchUut3.status;
   BenchCalls := BenchCalls + 1;
 66:
   BenchUut3.cyclicExecution := TRUE;
   BenchUut3.trigger := FALSE;
   BenchUut3.value := LREAL#37.0;
   BenchUut3.windowSize := INT#100;
   BenchUut3.reset := FALSE;
   TraceIn_cyclicExecution[66] := BenchUut3.cyclicExecution;
   TraceIn_trigger[66] := BenchUut3.trigger;
   TraceIn_value[66] := BenchUut3.value;
   TraceIn_windowSize[66] := BenchUut3.windowSize;
   TraceIn_reset[66] := BenchUut3.reset;
   BenchUut3();
   TraceOut_average[66] := BenchUut3.average;
   TraceOut_windowSizeReached[66] := BenchUut3.windowSizeReached;
   TraceOut_error[66] := BenchUut3.error;
   TraceOut_status[66] := BenchUut3.status;
   BenchCalls := BenchCalls + 1;
 67:
   BenchUut3.cyclicExecution := TRUE;
   BenchUut3.trigger := FALSE;
   BenchUut3.value := LREAL#38.0;
   BenchUut3.windowSize := INT#100;
   BenchUut3.reset := FALSE;
   TraceIn_cyclicExecution[67] := BenchUut3.cyclicExecution;
   TraceIn_trigger[67] := BenchUut3.trigger;
   TraceIn_value[67] := BenchUut3.value;
   TraceIn_windowSize[67] := BenchUut3.windowSize;
   TraceIn_reset[67] := BenchUut3.reset;
   BenchUut3();
   TraceOut_average[67] := BenchUut3.average;
   TraceOut_windowSizeReached[67] := BenchUut3.windowSizeReached;
   TraceOut_error[67] := BenchUut3.error;
   TraceOut_status[67] := BenchUut3.status;
   BenchCalls := BenchCalls + 1;
 68:
   BenchUut3.cyclicExecution := TRUE;
   BenchUut3.trigger := FALSE;
   BenchUut3.value := LREAL#39.0;
   BenchUut3.windowSize := INT#100;
   BenchUut3.reset := FALSE;
   TraceIn_cyclicExecution[68] := BenchUut3.cyclicExecution;
   TraceIn_trigger[68] := BenchUut3.trigger;
   TraceIn_value[68] := BenchUut3.value;
   TraceIn_windowSize[68] := BenchUut3.windowSize;
   TraceIn_reset[68] := BenchUut3.reset;
   BenchUut3();
   TraceOut_average[68] := BenchUut3.average;
   TraceOut_windowSizeReached[68] := BenchUut3.windowSizeReached;
   TraceOut_error[68] := BenchUut3.error;
   TraceOut_status[68] := BenchUut3.status;
   BenchCalls := BenchCalls + 1;
 69:
   BenchUut3.cyclicExecution := TRUE;
   BenchUut3.trigger := FALSE;
   BenchUut3.value := LREAL#40.0;
   BenchUut3.windowSize := INT#100;
   BenchUut3.reset := FALSE;
   TraceIn_cyclicExecution[69] := BenchUut3.cyclicExecution;
   TraceIn_trigger[69] := BenchUut3.trigger;
   TraceIn_value[69] := BenchUut3.value;
   TraceIn_windowSize[69] := BenchUut3.windowSize;
   TraceIn_reset[69] := BenchUut3.reset;
   BenchUut3();
   TraceOut_average[69] := BenchUut3.average;
   TraceOut_windowSizeReached[69] := BenchUut3.windowSizeReached;
   TraceOut_error[69] := BenchUut3.error;
   TraceOut_status[69] := BenchUut3.status;
   BenchCalls := BenchCalls + 1;
 70:
   BenchUut3.cyclicExecution := TRUE;
   BenchUut3.trigger := FALSE;
   BenchUut3.value := LREAL#41.0;
   BenchUut3.windowSize := INT#100;
   BenchUut3.reset := FALSE;
   TraceIn_cyclicExecution[70] := BenchUut3.cyclicExecution;
   TraceIn_trigger[70] := BenchUut3.trigger;
   TraceIn_value[70] := BenchUut3.value;
   TraceIn_windowSize[70] := BenchUut3.windowSize;
   TraceIn_reset[70] := BenchUut3.reset;
   BenchUut3();
   TraceOut_average[70] := BenchUut3.average;
   TraceOut_windowSizeReached[70] := BenchUut3.windowSizeReached;
   TraceOut_error[70] := BenchUut3.error;
   TraceOut_status[70] := BenchUut3.status;
   BenchCalls := BenchCalls + 1;
 71:
   BenchUut3.cyclicExecution := TRUE;
   BenchUut3.trigger := FALSE;
   BenchUut3.value := LREAL#42.0;
   BenchUut3.windowSize := INT#100;
   BenchUut3.reset := FALSE;
   TraceIn_cyclicExecution[71] := BenchUut3.cyclicExecution;
   TraceIn_trigger[71] := BenchUut3.trigger;
   TraceIn_value[71] := BenchUut3.value;
   TraceIn_windowSize[71] := BenchUut3.windowSize;
   TraceIn_reset[71] := BenchUut3.reset;
   BenchUut3();
   TraceOut_average[71] := BenchUut3.average;
   TraceOut_windowSizeReached[71] := BenchUut3.windowSizeReached;
   TraceOut_error[71] := BenchUut3.error;
   TraceOut_status[71] := BenchUut3.status;
   BenchCalls := BenchCalls + 1;
 72:
   BenchUut3.cyclicExecution := TRUE;
   BenchUut3.trigger := FALSE;
   BenchUut3.value := LREAL#43.0;
   BenchUut3.windowSize := INT#100;
   BenchUut3.reset := FALSE;
   TraceIn_cyclicExecution[72] := BenchUut3.cyclicExecution;
   TraceIn_trigger[72] := BenchUut3.trigger;
   TraceIn_value[72] := BenchUut3.value;
   TraceIn_windowSize[72] := BenchUut3.windowSize;
   TraceIn_reset[72] := BenchUut3.reset;
   BenchUut3();
   TraceOut_average[72] := BenchUut3.average;
   TraceOut_windowSizeReached[72] := BenchUut3.windowSizeReached;
   TraceOut_error[72] := BenchUut3.error;
   TraceOut_status[72] := BenchUut3.status;
   BenchCalls := BenchCalls + 1;
 73:
   BenchUut3.cyclicExecution := TRUE;
   BenchUut3.trigger := FALSE;
   BenchUut3.value := LREAL#44.0;
   BenchUut3.windowSize := INT#100;
   BenchUut3.reset := FALSE;
   TraceIn_cyclicExecution[73] := BenchUut3.cyclicExecution;
   TraceIn_trigger[73] := BenchUut3.trigger;
   TraceIn_value[73] := BenchUut3.value;
   TraceIn_windowSize[73] := BenchUut3.windowSize;
   TraceIn_reset[73] := BenchUut3.reset;
   BenchUut3();
   TraceOut_average[73] := BenchUut3.average;
   TraceOut_windowSizeReached[73] := BenchUut3.windowSizeReached;
   TraceOut_error[73] := BenchUut3.error;
   TraceOut_status[73] := BenchUut3.status;
   BenchCalls := BenchCalls + 1;
 74:
   BenchUut3.cyclicExecution := TRUE;
   BenchUut3.trigger := FALSE;
   BenchUut3.value := LREAL#45.0;
   BenchUut3.windowSize := INT#100;
   BenchUut3.reset := FALSE;
   TraceIn_cyclicExecution[74] := BenchUut3.cyclicExecution;
   TraceIn_trigger[74] := BenchUut3.trigger;
   TraceIn_value[74] := BenchUut3.value;
   TraceIn_windowSize[74] := BenchUut3.windowSize;
   TraceIn_reset[74] := BenchUut3.reset;
   BenchUut3();
   TraceOut_average[74] := BenchUut3.average;
   TraceOut_windowSizeReached[74] := BenchUut3.windowSizeReached;
   TraceOut_error[74] := BenchUut3.error;
   TraceOut_status[74] := BenchUut3.status;
   BenchCalls := BenchCalls + 1;
 75:
   BenchUut3.cyclicExecution := TRUE;
   BenchUut3.trigger := FALSE;
   BenchUut3.value := LREAL#46.0;
   BenchUut3.windowSize := INT#100;
   BenchUut3.reset := FALSE;
   TraceIn_cyclicExecution[75] := BenchUut3.cyclicExecution;
   TraceIn_trigger[75] := BenchUut3.trigger;
   TraceIn_value[75] := BenchUut3.value;
   TraceIn_windowSize[75] := BenchUut3.windowSize;
   TraceIn_reset[75] := BenchUut3.reset;
   BenchUut3();
   TraceOut_average[75] := BenchUut3.average;
   TraceOut_windowSizeReached[75] := BenchUut3.windowSizeReached;
   TraceOut_error[75] := BenchUut3.error;
   TraceOut_status[75] := BenchUut3.status;
   BenchCalls := BenchCalls + 1;
 76:
   BenchUut3.cyclicExecution := TRUE;
   BenchUut3.trigger := FALSE;
   BenchUut3.value := LREAL#47.0;
   BenchUut3.windowSize := INT#100;
   BenchUut3.reset := FALSE;
   TraceIn_cyclicExecution[76] := BenchUut3.cyclicExecution;
   TraceIn_trigger[76] := BenchUut3.trigger;
   TraceIn_value[76] := BenchUut3.value;
   TraceIn_windowSize[76] := BenchUut3.windowSize;
   TraceIn_reset[76] := BenchUut3.reset;
   BenchUut3();
   TraceOut_average[76] := BenchUut3.average;
   TraceOut_windowSizeReached[76] := BenchUut3.windowSizeReached;
   TraceOut_error[76] := BenchUut3.error;
   TraceOut_status[76] := BenchUut3.status;
   BenchCalls := BenchCalls + 1;
 77:
   BenchUut3.cyclicExecution := TRUE;
   BenchUut3.trigger := FALSE;
   BenchUut3.value := LREAL#48.0;
   BenchUut3.windowSize := INT#100;
   BenchUut3.reset := FALSE;
   TraceIn_cyclicExecution[77] := BenchUut3.cyclicExecution;
   TraceIn_trigger[77] := BenchUut3.trigger;
   TraceIn_value[77] := BenchUut3.value;
   TraceIn_windowSize[77] := BenchUut3.windowSize;
   TraceIn_reset[77] := BenchUut3.reset;
   BenchUut3();
   TraceOut_average[77] := BenchUut3.average;
   TraceOut_windowSizeReached[77] := BenchUut3.windowSizeReached;
   TraceOut_error[77] := BenchUut3.error;
   TraceOut_status[77] := BenchUut3.status;
   BenchCalls := BenchCalls + 1;
 78:
   BenchUut3.cyclicExecution := TRUE;
   BenchUut3.trigger := FALSE;
   BenchUut3.value := LREAL#49.0;
   BenchUut3.windowSize := INT#100;
   BenchUut3.reset := FALSE;
   TraceIn_cyclicExecution[78] := BenchUut3.cyclicExecution;
   TraceIn_trigger[78] := BenchUut3.trigger;
   TraceIn_value[78] := BenchUut3.value;
   TraceIn_windowSize[78] := BenchUut3.windowSize;
   TraceIn_reset[78] := BenchUut3.reset;
   BenchUut3();
   TraceOut_average[78] := BenchUut3.average;
   TraceOut_windowSizeReached[78] := BenchUut3.windowSizeReached;
   TraceOut_error[78] := BenchUut3.error;
   TraceOut_status[78] := BenchUut3.status;
   BenchCalls := BenchCalls + 1;
 79:
   BenchUut3.cyclicExecution := TRUE;
   BenchUut3.trigger := FALSE;
   BenchUut3.value := LREAL#50.0;
   BenchUut3.windowSize := INT#100;
   BenchUut3.reset := FALSE;
   TraceIn_cyclicExecution[79] := BenchUut3.cyclicExecution;
   TraceIn_trigger[79] := BenchUut3.trigger;
   TraceIn_value[79] := BenchUut3.value;
   TraceIn_windowSize[79] := BenchUut3.windowSize;
   TraceIn_reset[79] := BenchUut3.reset;
   BenchUut3();
   TraceOut_average[79] := BenchUut3.average;
   TraceOut_windowSizeReached[79] := BenchUut3.windowSizeReached;
   TraceOut_error[79] := BenchUut3.error;
   TraceOut_status[79] := BenchUut3.status;
   BenchCalls := BenchCalls + 1;
 80:
   BenchUut3.cyclicExecution := TRUE;
   BenchUut3.trigger := FALSE;
   BenchUut3.value := LREAL#51.0;
   BenchUut3.windowSize := INT#100;
   BenchUut3.reset := FALSE;
   TraceIn_cyclicExecution[80] := BenchUut3.cyclicExecution;
   TraceIn_trigger[80] := BenchUut3.trigger;
   TraceIn_value[80] := BenchUut3.value;
   TraceIn_windowSize[80] := BenchUut3.windowSize;
   TraceIn_reset[80] := BenchUut3.reset;
   BenchUut3();
   TraceOut_average[80] := BenchUut3.average;
   TraceOut_windowSizeReached[80] := BenchUut3.windowSizeReached;
   TraceOut_error[80] := BenchUut3.error;
   TraceOut_status[80] := BenchUut3.status;
   BenchCalls := BenchCalls + 1;
 81:
   BenchUut3.cyclicExecution := TRUE;
   BenchUut3.trigger := FALSE;
   BenchUut3.value := LREAL#52.0;
   BenchUut3.windowSize := INT#100;
   BenchUut3.reset := FALSE;
   TraceIn_cyclicExecution[81] := BenchUut3.cyclicExecution;
   TraceIn_trigger[81] := BenchUut3.trigger;
   TraceIn_value[81] := BenchUut3.value;
   TraceIn_windowSize[81] := BenchUut3.windowSize;
   TraceIn_reset[81] := BenchUut3.reset;
   BenchUut3();
   TraceOut_average[81] := BenchUut3.average;
   TraceOut_windowSizeReached[81] := BenchUut3.windowSizeReached;
   TraceOut_error[81] := BenchUut3.error;
   TraceOut_status[81] := BenchUut3.status;
   BenchCalls := BenchCalls + 1;
 82:
   BenchUut3.cyclicExecution := TRUE;
   BenchUut3.trigger := FALSE;
   BenchUut3.value := LREAL#53.0;
   BenchUut3.windowSize := INT#100;
   BenchUut3.reset := FALSE;
   TraceIn_cyclicExecution[82] := BenchUut3.cyclicExecution;
   TraceIn_trigger[82] := BenchUut3.trigger;
   TraceIn_value[82] := BenchUut3.value;
   TraceIn_windowSize[82] := BenchUut3.windowSize;
   TraceIn_reset[82] := BenchUut3.reset;
   BenchUut3();
   TraceOut_average[82] := BenchUut3.average;
   TraceOut_windowSizeReached[82] := BenchUut3.windowSizeReached;
   TraceOut_error[82] := BenchUut3.error;
   TraceOut_status[82] := BenchUut3.status;
   BenchCalls := BenchCalls + 1;
 83:
   BenchUut3.cyclicExecution := TRUE;
   BenchUut3.trigger := FALSE;
   BenchUut3.value := LREAL#54.0;
   BenchUut3.windowSize := INT#100;
   BenchUut3.reset := FALSE;
   TraceIn_cyclicExecution[83] := BenchUut3.cyclicExecution;
   TraceIn_trigger[83] := BenchUut3.trigger;
   TraceIn_value[83] := BenchUut3.value;
   TraceIn_windowSize[83] := BenchUut3.windowSize;
   TraceIn_reset[83] := BenchUut3.reset;
   BenchUut3();
   TraceOut_average[83] := BenchUut3.average;
   TraceOut_windowSizeReached[83] := BenchUut3.windowSizeReached;
   TraceOut_error[83] := BenchUut3.error;
   TraceOut_status[83] := BenchUut3.status;
   BenchCalls := BenchCalls + 1;
 84:
   BenchUut3.cyclicExecution := TRUE;
   BenchUut3.trigger := FALSE;
   BenchUut3.value := LREAL#55.0;
   BenchUut3.windowSize := INT#100;
   BenchUut3.reset := FALSE;
   TraceIn_cyclicExecution[84] := BenchUut3.cyclicExecution;
   TraceIn_trigger[84] := BenchUut3.trigger;
   TraceIn_value[84] := BenchUut3.value;
   TraceIn_windowSize[84] := BenchUut3.windowSize;
   TraceIn_reset[84] := BenchUut3.reset;
   BenchUut3();
   TraceOut_average[84] := BenchUut3.average;
   TraceOut_windowSizeReached[84] := BenchUut3.windowSizeReached;
   TraceOut_error[84] := BenchUut3.error;
   TraceOut_status[84] := BenchUut3.status;
   BenchCalls := BenchCalls + 1;
 85:
   BenchUut3.cyclicExecution := TRUE;
   BenchUut3.trigger := FALSE;
   BenchUut3.value := LREAL#56.0;
   BenchUut3.windowSize := INT#100;
   BenchUut3.reset := FALSE;
   TraceIn_cyclicExecution[85] := BenchUut3.cyclicExecution;
   TraceIn_trigger[85] := BenchUut3.trigger;
   TraceIn_value[85] := BenchUut3.value;
   TraceIn_windowSize[85] := BenchUut3.windowSize;
   TraceIn_reset[85] := BenchUut3.reset;
   BenchUut3();
   TraceOut_average[85] := BenchUut3.average;
   TraceOut_windowSizeReached[85] := BenchUut3.windowSizeReached;
   TraceOut_error[85] := BenchUut3.error;
   TraceOut_status[85] := BenchUut3.status;
   BenchCalls := BenchCalls + 1;
 86:
   BenchUut3.cyclicExecution := TRUE;
   BenchUut3.trigger := FALSE;
   BenchUut3.value := LREAL#57.0;
   BenchUut3.windowSize := INT#100;
   BenchUut3.reset := FALSE;
   TraceIn_cyclicExecution[86] := BenchUut3.cyclicExecution;
   TraceIn_trigger[86] := BenchUut3.trigger;
   TraceIn_value[86] := BenchUut3.value;
   TraceIn_windowSize[86] := BenchUut3.windowSize;
   TraceIn_reset[86] := BenchUut3.reset;
   BenchUut3();
   TraceOut_average[86] := BenchUut3.average;
   TraceOut_windowSizeReached[86] := BenchUut3.windowSizeReached;
   TraceOut_error[86] := BenchUut3.error;
   TraceOut_status[86] := BenchUut3.status;
   BenchCalls := BenchCalls + 1;
 87:
   BenchUut3.cyclicExecution := TRUE;
   BenchUut3.trigger := FALSE;
   BenchUut3.value := LREAL#58.0;
   BenchUut3.windowSize := INT#100;
   BenchUut3.reset := FALSE;
   TraceIn_cyclicExecution[87] := BenchUut3.cyclicExecution;
   TraceIn_trigger[87] := BenchUut3.trigger;
   TraceIn_value[87] := BenchUut3.value;
   TraceIn_windowSize[87] := BenchUut3.windowSize;
   TraceIn_reset[87] := BenchUut3.reset;
   BenchUut3();
   TraceOut_average[87] := BenchUut3.average;
   TraceOut_windowSizeReached[87] := BenchUut3.windowSizeReached;
   TraceOut_error[87] := BenchUut3.error;
   TraceOut_status[87] := BenchUut3.status;
   BenchCalls := BenchCalls + 1;
 88:
   BenchUut3.cyclicExecution := TRUE;
   BenchUut3.trigger := FALSE;
   BenchUut3.value := LREAL#59.0;
   BenchUut3.windowSize := INT#100;
   BenchUut3.reset := FALSE;
   TraceIn_cyclicExecution[88] := BenchUut3.cyclicExecution;
   TraceIn_trigger[88] := BenchUut3.trigger;
   TraceIn_value[88] := BenchUut3.value;
   TraceIn_windowSize[88] := BenchUut3.windowSize;
   TraceIn_reset[88] := BenchUut3.reset;
   BenchUut3();
   TraceOut_average[88] := BenchUut3.average;
   TraceOut_windowSizeReached[88] := BenchUut3.windowSizeReached;
   TraceOut_error[88] := BenchUut3.error;
   TraceOut_status[88] := BenchUut3.status;
   BenchCalls := BenchCalls + 1;
 89:
   BenchUut3.cyclicExecution := TRUE;
   BenchUut3.trigger := FALSE;
   BenchUut3.value := LREAL#60.0;
   BenchUut3.windowSize := INT#100;
   BenchUut3.reset := FALSE;
   TraceIn_cyclicExecution[89] := BenchUut3.cyclicExecution;
   TraceIn_trigger[89] := BenchUut3.trigger;
   TraceIn_value[89] := BenchUut3.value;
   TraceIn_windowSize[89] := BenchUut3.windowSize;
   TraceIn_reset[89] := BenchUut3.reset;
   BenchUut3();
   TraceOut_average[89] := BenchUut3.average;
   TraceOut_windowSizeReached[89] := BenchUut3.windowSizeReached;
   TraceOut_error[89] := BenchUut3.error;
   TraceOut_status[89] := BenchUut3.status;
   BenchCalls := BenchCalls + 1;
 90:
   BenchUut3.cyclicExecution := TRUE;
   BenchUut3.trigger := FALSE;
   BenchUut3.value := LREAL#61.0;
   BenchUut3.windowSize := INT#100;
   BenchUut3.reset := FALSE;
   TraceIn_cyclicExecution[90] := BenchUut3.cyclicExecution;
   TraceIn_trigger[90] := BenchUut3.trigger;
   TraceIn_value[90] := BenchUut3.value;
   TraceIn_windowSize[90] := BenchUut3.windowSize;
   TraceIn_reset[90] := BenchUut3.reset;
   BenchUut3();
   TraceOut_average[90] := BenchUut3.average;
   TraceOut_windowSizeReached[90] := BenchUut3.windowSizeReached;
   TraceOut_error[90] := BenchUut3.error;
   TraceOut_status[90] := BenchUut3.status;
   BenchCalls := BenchCalls + 1;
 91:
   BenchUut3.cyclicExecution := TRUE;
   BenchUut3.trigger := FALSE;
   BenchUut3.value := LREAL#62.0;
   BenchUut3.windowSize := INT#100;
   BenchUut3.reset := FALSE;
   TraceIn_cyclicExecution[91] := BenchUut3.cyclicExecution;
   TraceIn_trigger[91] := BenchUut3.trigger;
   TraceIn_value[91] := BenchUut3.value;
   TraceIn_windowSize[91] := BenchUut3.windowSize;
   TraceIn_reset[91] := BenchUut3.reset;
   BenchUut3();
   TraceOut_average[91] := BenchUut3.average;
   TraceOut_windowSizeReached[91] := BenchUut3.windowSizeReached;
   TraceOut_error[91] := BenchUut3.error;
   TraceOut_status[91] := BenchUut3.status;
   BenchCalls := BenchCalls + 1;
 92:
   BenchUut3.cyclicExecution := TRUE;
   BenchUut3.trigger := FALSE;
   BenchUut3.value := LREAL#63.0;
   BenchUut3.windowSize := INT#100;
   BenchUut3.reset := FALSE;
   TraceIn_cyclicExecution[92] := BenchUut3.cyclicExecution;
   TraceIn_trigger[92] := BenchUut3.trigger;
   TraceIn_value[92] := BenchUut3.value;
   TraceIn_windowSize[92] := BenchUut3.windowSize;
   TraceIn_reset[92] := BenchUut3.reset;
   BenchUut3();
   TraceOut_average[92] := BenchUut3.average;
   TraceOut_windowSizeReached[92] := BenchUut3.windowSizeReached;
   TraceOut_error[92] := BenchUut3.error;
   TraceOut_status[92] := BenchUut3.status;
   BenchCalls := BenchCalls + 1;
 93:
   BenchUut3.cyclicExecution := TRUE;
   BenchUut3.trigger := FALSE;
   BenchUut3.value := LREAL#64.0;
   BenchUut3.windowSize := INT#100;
   BenchUut3.reset := FALSE;
   TraceIn_cyclicExecution[93] := BenchUut3.cyclicExecution;
   TraceIn_trigger[93] := BenchUut3.trigger;
   TraceIn_value[93] := BenchUut3.value;
   TraceIn_windowSize[93] := BenchUut3.windowSize;
   TraceIn_reset[93] := BenchUut3.reset;
   BenchUut3();
   TraceOut_average[93] := BenchUut3.average;
   TraceOut_windowSizeReached[93] := BenchUut3.windowSizeReached;
   TraceOut_error[93] := BenchUut3.error;
   TraceOut_status[93] := BenchUut3.status;
   BenchCalls := BenchCalls + 1;
 94:
   BenchUut3.cyclicExecution := TRUE;
   BenchUut3.trigger := FALSE;
   BenchUut3.value := LREAL#65.0;
   BenchUut3.windowSize := INT#100;
   BenchUut3.reset := FALSE;
   TraceIn_cyclicExecution[94] := BenchUut3.cyclicExecution;
   TraceIn_trigger[94] := BenchUut3.trigger;
   TraceIn_value[94] := BenchUut3.value;
   TraceIn_windowSize[94] := BenchUut3.windowSize;
   TraceIn_reset[94] := BenchUut3.reset;
   BenchUut3();
   TraceOut_average[94] := BenchUut3.average;
   TraceOut_windowSizeReached[94] := BenchUut3.windowSizeReached;
   TraceOut_error[94] := BenchUut3.error;
   TraceOut_status[94] := BenchUut3.status;
   BenchCalls := BenchCalls + 1;
 95:
   BenchUut3.cyclicExecution := TRUE;
   BenchUut3.trigger := FALSE;
   BenchUut3.value := LREAL#66.0;
   BenchUut3.windowSize := INT#100;
   BenchUut3.reset := FALSE;
   TraceIn_cyclicExecution[95] := BenchUut3.cyclicExecution;
   TraceIn_trigger[95] := BenchUut3.trigger;
   TraceIn_value[95] := BenchUut3.value;
   TraceIn_windowSize[95] := BenchUut3.windowSize;
   TraceIn_reset[95] := BenchUut3.reset;
   BenchUut3();
   TraceOut_average[95] := BenchUut3.average;
   TraceOut_windowSizeReached[95] := BenchUut3.windowSizeReached;
   TraceOut_error[95] := BenchUut3.error;
   TraceOut_status[95] := BenchUut3.status;
   BenchCalls := BenchCalls + 1;
 96:
   BenchUut3.cyclicExecution := TRUE;
   BenchUut3.trigger := FALSE;
   BenchUut3.value := LREAL#67.0;
   BenchUut3.windowSize := INT#100;
   BenchUut3.reset := FALSE;
   TraceIn_cyclicExecution[96] := BenchUut3.cyclicExecution;
   TraceIn_trigger[96] := BenchUut3.trigger;
   TraceIn_value[96] := BenchUut3.value;
   TraceIn_windowSize[96] := BenchUut3.windowSize;
   TraceIn_reset[96] := BenchUut3.reset;
   BenchUut3();
   TraceOut_average[96] := BenchUut3.average;
   TraceOut_windowSizeReached[96] := BenchUut3.windowSizeReached;
   TraceOut_error[96] := BenchUut3.error;
   TraceOut_status[96] := BenchUut3.status;
   BenchCalls := BenchCalls + 1;
 97:
   BenchUut3.cyclicExecution := TRUE;
   BenchUut3.trigger := FALSE;
   BenchUut3.value := LREAL#68.0;
   BenchUut3.windowSize := INT#100;
   BenchUut3.reset := FALSE;
   TraceIn_cyclicExecution[97] := BenchUut3.cyclicExecution;
   TraceIn_trigger[97] := BenchUut3.trigger;
   TraceIn_value[97] := BenchUut3.value;
   TraceIn_windowSize[97] := BenchUut3.windowSize;
   TraceIn_reset[97] := BenchUut3.reset;
   BenchUut3();
   TraceOut_average[97] := BenchUut3.average;
   TraceOut_windowSizeReached[97] := BenchUut3.windowSizeReached;
   TraceOut_error[97] := BenchUut3.error;
   TraceOut_status[97] := BenchUut3.status;
   BenchCalls := BenchCalls + 1;
 98:
   BenchUut3.cyclicExecution := TRUE;
   BenchUut3.trigger := FALSE;
   BenchUut3.value := LREAL#69.0;
   BenchUut3.windowSize := INT#100;
   BenchUut3.reset := FALSE;
   TraceIn_cyclicExecution[98] := BenchUut3.cyclicExecution;
   TraceIn_trigger[98] := BenchUut3.trigger;
   TraceIn_value[98] := BenchUut3.value;
   TraceIn_windowSize[98] := BenchUut3.windowSize;
   TraceIn_reset[98] := BenchUut3.reset;
   BenchUut3();
   TraceOut_average[98] := BenchUut3.average;
   TraceOut_windowSizeReached[98] := BenchUut3.windowSizeReached;
   TraceOut_error[98] := BenchUut3.error;
   TraceOut_status[98] := BenchUut3.status;
   BenchCalls := BenchCalls + 1;
 99:
   BenchUut3.cyclicExecution := TRUE;
   BenchUut3.trigger := FALSE;
   BenchUut3.value := LREAL#70.0;
   BenchUut3.windowSize := INT#100;
   BenchUut3.reset := FALSE;
   TraceIn_cyclicExecution[99] := BenchUut3.cyclicExecution;
   TraceIn_trigger[99] := BenchUut3.trigger;
   TraceIn_value[99] := BenchUut3.value;
   TraceIn_windowSize[99] := BenchUut3.windowSize;
   TraceIn_reset[99] := BenchUut3.reset;
   BenchUut3();
   TraceOut_average[99] := BenchUut3.average;
   TraceOut_windowSizeReached[99] := BenchUut3.windowSizeReached;
   TraceOut_error[99] := BenchUut3.error;
   TraceOut_status[99] := BenchUut3.status;
   BenchCalls := BenchCalls + 1;
 100:
   BenchUut3.cyclicExecution := TRUE;
   BenchUut3.trigger := FALSE;
   BenchUut3.value := LREAL#71.0;
   BenchUut3.windowSize := INT#100;
   BenchUut3.reset := FALSE;
   TraceIn_cyclicExecution[100] := BenchUut3.cyclicExecution;
   TraceIn_trigger[100] := BenchUut3.trigger;
   TraceIn_value[100] := BenchUut3.value;
   TraceIn_windowSize[100] := BenchUut3.windowSize;
   TraceIn_reset[100] := BenchUut3.reset;
   BenchUut3();
   TraceOut_average[100] := BenchUut3.average;
   TraceOut_windowSizeReached[100] := BenchUut3.windowSizeReached;
   TraceOut_error[100] := BenchUut3.error;
   TraceOut_status[100] := BenchUut3.status;
   BenchCalls := BenchCalls + 1;
 101:
   BenchUut3.cyclicExecution := TRUE;
   BenchUut3.trigger := FALSE;
   BenchUut3.value := LREAL#72.0;
   BenchUut3.windowSize := INT#100;
   BenchUut3.reset := FALSE;
   TraceIn_cyclicExecution[101] := BenchUut3.cyclicExecution;
   TraceIn_trigger[101] := BenchUut3.trigger;
   TraceIn_value[101] := BenchUut3.value;
   TraceIn_windowSize[101] := BenchUut3.windowSize;
   TraceIn_reset[101] := BenchUut3.reset;
   BenchUut3();
   TraceOut_average[101] := BenchUut3.average;
   TraceOut_windowSizeReached[101] := BenchUut3.windowSizeReached;
   TraceOut_error[101] := BenchUut3.error;
   TraceOut_status[101] := BenchUut3.status;
   BenchCalls := BenchCalls + 1;
 102:
   BenchUut3.cyclicExecution := TRUE;
   BenchUut3.trigger := FALSE;
   BenchUut3.value := LREAL#73.0;
   BenchUut3.windowSize := INT#100;
   BenchUut3.reset := FALSE;
   TraceIn_cyclicExecution[102] := BenchUut3.cyclicExecution;
   TraceIn_trigger[102] := BenchUut3.trigger;
   TraceIn_value[102] := BenchUut3.value;
   TraceIn_windowSize[102] := BenchUut3.windowSize;
   TraceIn_reset[102] := BenchUut3.reset;
   BenchUut3();
   TraceOut_average[102] := BenchUut3.average;
   TraceOut_windowSizeReached[102] := BenchUut3.windowSizeReached;
   TraceOut_error[102] := BenchUut3.error;
   TraceOut_status[102] := BenchUut3.status;
   BenchCalls := BenchCalls + 1;
 103:
   BenchUut3.cyclicExecution := TRUE;
   BenchUut3.trigger := FALSE;
   BenchUut3.value := LREAL#74.0;
   BenchUut3.windowSize := INT#100;
   BenchUut3.reset := FALSE;
   TraceIn_cyclicExecution[103] := BenchUut3.cyclicExecution;
   TraceIn_trigger[103] := BenchUut3.trigger;
   TraceIn_value[103] := BenchUut3.value;
   TraceIn_windowSize[103] := BenchUut3.windowSize;
   TraceIn_reset[103] := BenchUut3.reset;
   BenchUut3();
   TraceOut_average[103] := BenchUut3.average;
   TraceOut_windowSizeReached[103] := BenchUut3.windowSizeReached;
   TraceOut_error[103] := BenchUut3.error;
   TraceOut_status[103] := BenchUut3.status;
   BenchCalls := BenchCalls + 1;
 104:
   BenchUut3.cyclicExecution := TRUE;
   BenchUut3.trigger := FALSE;
   BenchUut3.value := LREAL#75.0;
   BenchUut3.windowSize := INT#100;
   BenchUut3.reset := FALSE;
   TraceIn_cyclicExecution[104] := BenchUut3.cyclicExecution;
   TraceIn_trigger[104] := BenchUut3.trigger;
   TraceIn_value[104] := BenchUut3.value;
   TraceIn_windowSize[104] := BenchUut3.windowSize;
   TraceIn_reset[104] := BenchUut3.reset;
   BenchUut3();
   TraceOut_average[104] := BenchUut3.average;
   TraceOut_windowSizeReached[104] := BenchUut3.windowSizeReached;
   TraceOut_error[104] := BenchUut3.error;
   TraceOut_status[104] := BenchUut3.status;
   BenchCalls := BenchCalls + 1;
 105:
   BenchUut3.cyclicExecution := TRUE;
   BenchUut3.trigger := FALSE;
   BenchUut3.value := LREAL#76.0;
   BenchUut3.windowSize := INT#100;
   BenchUut3.reset := FALSE;
   TraceIn_cyclicExecution[105] := BenchUut3.cyclicExecution;
   TraceIn_trigger[105] := BenchUut3.trigger;
   TraceIn_value[105] := BenchUut3.value;
   TraceIn_windowSize[105] := BenchUut3.windowSize;
   TraceIn_reset[105] := BenchUut3.reset;
   BenchUut3();
   TraceOut_average[105] := BenchUut3.average;
   TraceOut_windowSizeReached[105] := BenchUut3.windowSizeReached;
   TraceOut_error[105] := BenchUut3.error;
   TraceOut_status[105] := BenchUut3.status;
   BenchCalls := BenchCalls + 1;
 106:
   BenchUut3.cyclicExecution := TRUE;
   BenchUut3.trigger := FALSE;
   BenchUut3.value := LREAL#77.0;
   BenchUut3.windowSize := INT#100;
   BenchUut3.reset := FALSE;
   TraceIn_cyclicExecution[106] := BenchUut3.cyclicExecution;
   TraceIn_trigger[106] := BenchUut3.trigger;
   TraceIn_value[106] := BenchUut3.value;
   TraceIn_windowSize[106] := BenchUut3.windowSize;
   TraceIn_reset[106] := BenchUut3.reset;
   BenchUut3();
   TraceOut_average[106] := BenchUut3.average;
   TraceOut_windowSizeReached[106] := BenchUut3.windowSizeReached;
   TraceOut_error[106] := BenchUut3.error;
   TraceOut_status[106] := BenchUut3.status;
   BenchCalls := BenchCalls + 1;
 107:
   BenchUut3.cyclicExecution := TRUE;
   BenchUut3.trigger := FALSE;
   BenchUut3.value := LREAL#78.0;
   BenchUut3.windowSize := INT#100;
   BenchUut3.reset := FALSE;
   TraceIn_cyclicExecution[107] := BenchUut3.cyclicExecution;
   TraceIn_trigger[107] := BenchUut3.trigger;
   TraceIn_value[107] := BenchUut3.value;
   TraceIn_windowSize[107] := BenchUut3.windowSize;
   TraceIn_reset[107] := BenchUut3.reset;
   BenchUut3();
   TraceOut_average[107] := BenchUut3.average;
   TraceOut_windowSizeReached[107] := BenchUut3.windowSizeReached;
   TraceOut_error[107] := BenchUut3.error;
   TraceOut_status[107] := BenchUut3.status;
   BenchCalls := BenchCalls + 1;
 108:
   BenchUut3.cyclicExecution := TRUE;
   BenchUut3.trigger := FALSE;
   BenchUut3.value := LREAL#79.0;
   BenchUut3.windowSize := INT#100;
   BenchUut3.reset := FALSE;
   TraceIn_cyclicExecution[108] := BenchUut3.cyclicExecution;
   TraceIn_trigger[108] := BenchUut3.trigger;
   TraceIn_value[108] := BenchUut3.value;
   TraceIn_windowSize[108] := BenchUut3.windowSize;
   TraceIn_reset[108] := BenchUut3.reset;
   BenchUut3();
   TraceOut_average[108] := BenchUut3.average;
   TraceOut_windowSizeReached[108] := BenchUut3.windowSizeReached;
   TraceOut_error[108] := BenchUut3.error;
   TraceOut_status[108] := BenchUut3.status;
   BenchCalls := BenchCalls + 1;
 109:
   BenchUut3.cyclicExecution := TRUE;
   BenchUut3.trigger := FALSE;
   BenchUut3.value := LREAL#80.0;
   BenchUut3.windowSize := INT#100;
   BenchUut3.reset := FALSE;
   TraceIn_cyclicExecution[109] := BenchUut3.cyclicExecution;
   TraceIn_trigger[109] := BenchUut3.trigger;
   TraceIn_value[109] := BenchUut3.value;
   TraceIn_windowSize[109] := BenchUut3.windowSize;
   TraceIn_reset[109] := BenchUut3.reset;
   BenchUut3();
   TraceOut_average[109] := BenchUut3.average;
   TraceOut_windowSizeReached[109] := BenchUut3.windowSizeReached;
   TraceOut_error[109] := BenchUut3.error;
   TraceOut_status[109] := BenchUut3.status;
   BenchCalls := BenchCalls + 1;
 110:
   BenchUut3.cyclicExecution := TRUE;
   BenchUut3.trigger := FALSE;
   BenchUut3.value := LREAL#81.0;
   BenchUut3.windowSize := INT#100;
   BenchUut3.reset := FALSE;
   TraceIn_cyclicExecution[110] := BenchUut3.cyclicExecution;
   TraceIn_trigger[110] := BenchUut3.trigger;
   TraceIn_value[110] := BenchUut3.value;
   TraceIn_windowSize[110] := BenchUut3.windowSize;
   TraceIn_reset[110] := BenchUut3.reset;
   BenchUut3();
   TraceOut_average[110] := BenchUut3.average;
   TraceOut_windowSizeReached[110] := BenchUut3.windowSizeReached;
   TraceOut_error[110] := BenchUut3.error;
   TraceOut_status[110] := BenchUut3.status;
   BenchCalls := BenchCalls + 1;
 111:
   BenchUut3.cyclicExecution := TRUE;
   BenchUut3.trigger := FALSE;
   BenchUut3.value := LREAL#82.0;
   BenchUut3.windowSize := INT#100;
   BenchUut3.reset := FALSE;
   TraceIn_cyclicExecution[111] := BenchUut3.cyclicExecution;
   TraceIn_trigger[111] := BenchUut3.trigger;
   TraceIn_value[111] := BenchUut3.value;
   TraceIn_windowSize[111] := BenchUut3.windowSize;
   TraceIn_reset[111] := BenchUut3.reset;
   BenchUut3();
   TraceOut_average[111] := BenchUut3.average;
   TraceOut_windowSizeReached[111] := BenchUut3.windowSizeReached;
   TraceOut_error[111] := BenchUut3.error;
   TraceOut_status[111] := BenchUut3.status;
   BenchCalls := BenchCalls + 1;
 112:
   BenchUut3.cyclicExecution := TRUE;
   BenchUut3.trigger := FALSE;
   BenchUut3.value := LREAL#83.0;
   BenchUut3.windowSize := INT#100;
   BenchUut3.reset := FALSE;
   TraceIn_cyclicExecution[112] := BenchUut3.cyclicExecution;
   TraceIn_trigger[112] := BenchUut3.trigger;
   TraceIn_value[112] := BenchUut3.value;
   TraceIn_windowSize[112] := BenchUut3.windowSize;
   TraceIn_reset[112] := BenchUut3.reset;
   BenchUut3();
   TraceOut_average[112] := BenchUut3.average;
   TraceOut_windowSizeReached[112] := BenchUut3.windowSizeReached;
   TraceOut_error[112] := BenchUut3.error;
   TraceOut_status[112] := BenchUut3.status;
   BenchCalls := BenchCalls + 1;
 113:
   BenchUut3.cyclicExecution := TRUE;
   BenchUut3.trigger := FALSE;
   BenchUut3.value := LREAL#84.0;
   BenchUut3.windowSize := INT#100;
   BenchUut3.reset := FALSE;
   TraceIn_cyclicExecution[113] := BenchUut3.cyclicExecution;
   TraceIn_trigger[113] := BenchUut3.trigger;
   TraceIn_value[113] := BenchUut3.value;
   TraceIn_windowSize[113] := BenchUut3.windowSize;
   TraceIn_reset[113] := BenchUut3.reset;
   BenchUut3();
   TraceOut_average[113] := BenchUut3.average;
   TraceOut_windowSizeReached[113] := BenchUut3.windowSizeReached;
   TraceOut_error[113] := BenchUut3.error;
   TraceOut_status[113] := BenchUut3.status;
   BenchCalls := BenchCalls + 1;
 114:
   BenchUut3.cyclicExecution := TRUE;
   BenchUut3.trigger := FALSE;
   BenchUut3.value := LREAL#85.0;
   BenchUut3.windowSize := INT#100;
   BenchUut3.reset := FALSE;
   TraceIn_cyclicExecution[114] := BenchUut3.cyclicExecution;
   TraceIn_trigger[114] := BenchUut3.trigger;
   TraceIn_value[114] := BenchUut3.value;
   TraceIn_windowSize[114] := BenchUut3.windowSize;
   TraceIn_reset[114] := BenchUut3.reset;
   BenchUut3();
   TraceOut_average[114] := BenchUut3.average;
   TraceOut_windowSizeReached[114] := BenchUut3.windowSizeReached;
   TraceOut_error[114] := BenchUut3.error;
   TraceOut_status[114] := BenchUut3.status;
   BenchCalls := BenchCalls + 1;
 115:
   BenchUut3.cyclicExecution := TRUE;
   BenchUut3.trigger := FALSE;
   BenchUut3.value := LREAL#86.0;
   BenchUut3.windowSize := INT#100;
   BenchUut3.reset := FALSE;
   TraceIn_cyclicExecution[115] := BenchUut3.cyclicExecution;
   TraceIn_trigger[115] := BenchUut3.trigger;
   TraceIn_value[115] := BenchUut3.value;
   TraceIn_windowSize[115] := BenchUut3.windowSize;
   TraceIn_reset[115] := BenchUut3.reset;
   BenchUut3();
   TraceOut_average[115] := BenchUut3.average;
   TraceOut_windowSizeReached[115] := BenchUut3.windowSizeReached;
   TraceOut_error[115] := BenchUut3.error;
   TraceOut_status[115] := BenchUut3.status;
   BenchCalls := BenchCalls + 1;
 116:
   BenchUut3.cyclicExecution := TRUE;
   BenchUut3.trigger := FALSE;
   BenchUut3.value := LREAL#87.0;
   BenchUut3.windowSize := INT#100;
   BenchUut3.reset := FALSE;
   TraceIn_cyclicExecution[116] := BenchUut3.cyclicExecution;
   TraceIn_trigger[116] := BenchUut3.trigger;
   TraceIn_value[116] := BenchUut3.value;
   TraceIn_windowSize[116] := BenchUut3.windowSize;
   TraceIn_reset[116] := BenchUut3.reset;
   BenchUut3();
   TraceOut_average[116] := BenchUut3.average;
   TraceOut_windowSizeReached[116] := BenchUut3.windowSizeReached;
   TraceOut_error[116] := BenchUut3.error;
   TraceOut_status[116] := BenchUut3.status;
   BenchCalls := BenchCalls + 1;
 117:
   BenchUut3.cyclicExecution := TRUE;
   BenchUut3.trigger := FALSE;
   BenchUut3.value := LREAL#88.0;
   BenchUut3.windowSize := INT#100;
   BenchUut3.reset := FALSE;
   TraceIn_cyclicExecution[117] := BenchUut3.cyclicExecution;
   TraceIn_trigger[117] := BenchUut3.trigger;
   TraceIn_value[117] := BenchUut3.value;
   TraceIn_windowSize[117] := BenchUut3.windowSize;
   TraceIn_reset[117] := BenchUut3.reset;
   BenchUut3();
   TraceOut_average[117] := BenchUut3.average;
   TraceOut_windowSizeReached[117] := BenchUut3.windowSizeReached;
   TraceOut_error[117] := BenchUut3.error;
   TraceOut_status[117] := BenchUut3.status;
   BenchCalls := BenchCalls + 1;
 118:
   BenchUut3.cyclicExecution := TRUE;
   BenchUut3.trigger := FALSE;
   BenchUut3.value := LREAL#89.0;
   BenchUut3.windowSize := INT#100;
   BenchUut3.reset := FALSE;
   TraceIn_cyclicExecution[118] := BenchUut3.cyclicExecution;
   TraceIn_trigger[118] := BenchUut3.trigger;
   TraceIn_value[118] := BenchUut3.value;
   TraceIn_windowSize[118] := BenchUut3.windowSize;
   TraceIn_reset[118] := BenchUut3.reset;
   BenchUut3();
   TraceOut_average[118] := BenchUut3.average;
   TraceOut_windowSizeReached[118] := BenchUut3.windowSizeReached;
   TraceOut_error[118] := BenchUut3.error;
   TraceOut_status[118] := BenchUut3.status;
   BenchCalls := BenchCalls + 1;
 119:
   BenchUut3.cyclicExecution := TRUE;
   BenchUut3.trigger := FALSE;
   BenchUut3.value := LREAL#90.0;
   BenchUut3.windowSize := INT#100;
   BenchUut3.reset := FALSE;
   TraceIn_cyclicExecution[119] := BenchUut3.cyclicExecution;
   TraceIn_trigger[119] := BenchUut3.trigger;
   TraceIn_value[119] := BenchUut3.value;
   TraceIn_windowSize[119] := BenchUut3.windowSize;
   TraceIn_reset[119] := BenchUut3.reset;
   BenchUut3();
   TraceOut_average[119] := BenchUut3.average;
   TraceOut_windowSizeReached[119] := BenchUut3.windowSizeReached;
   TraceOut_error[119] := BenchUut3.error;
   TraceOut_status[119] := BenchUut3.status;
   BenchCalls := BenchCalls + 1;
 120:
   BenchUut3.cyclicExecution := TRUE;
   BenchUut3.trigger := FALSE;
   BenchUut3.value := LREAL#91.0;
   BenchUut3.windowSize := INT#100;
   BenchUut3.reset := FALSE;
   TraceIn_cyclicExecution[120] := BenchUut3.cyclicExecution;
   TraceIn_trigger[120] := BenchUut3.trigger;
   TraceIn_value[120] := BenchUut3.value;
   TraceIn_windowSize[120] := BenchUut3.windowSize;
   TraceIn_reset[120] := BenchUut3.reset;
   BenchUut3();
   TraceOut_average[120] := BenchUut3.average;
   TraceOut_windowSizeReached[120] := BenchUut3.windowSizeReached;
   TraceOut_error[120] := BenchUut3.error;
   TraceOut_status[120] := BenchUut3.status;
   BenchCalls := BenchCalls + 1;
 121:
   BenchUut3.cyclicExecution := TRUE;
   BenchUut3.trigger := FALSE;
   BenchUut3.value := LREAL#92.0;
   BenchUut3.windowSize := INT#100;
   BenchUut3.reset := FALSE;
   TraceIn_cyclicExecution[121] := BenchUut3.cyclicExecution;
   TraceIn_trigger[121] := BenchUut3.trigger;
   TraceIn_value[121] := BenchUut3.value;
   TraceIn_windowSize[121] := BenchUut3.windowSize;
   TraceIn_reset[121] := BenchUut3.reset;
   BenchUut3();
   TraceOut_average[121] := BenchUut3.average;
   TraceOut_windowSizeReached[121] := BenchUut3.windowSizeReached;
   TraceOut_error[121] := BenchUut3.error;
   TraceOut_status[121] := BenchUut3.status;
   BenchCalls := BenchCalls + 1;
 122:
   BenchUut3.cyclicExecution := TRUE;
   BenchUut3.trigger := FALSE;
   BenchUut3.value := LREAL#93.0;
   BenchUut3.windowSize := INT#100;
   BenchUut3.reset := FALSE;
   TraceIn_cyclicExecution[122] := BenchUut3.cyclicExecution;
   TraceIn_trigger[122] := BenchUut3.trigger;
   TraceIn_value[122] := BenchUut3.value;
   TraceIn_windowSize[122] := BenchUut3.windowSize;
   TraceIn_reset[122] := BenchUut3.reset;
   BenchUut3();
   TraceOut_average[122] := BenchUut3.average;
   TraceOut_windowSizeReached[122] := BenchUut3.windowSizeReached;
   TraceOut_error[122] := BenchUut3.error;
   TraceOut_status[122] := BenchUut3.status;
   BenchCalls := BenchCalls + 1;
 123:
   BenchUut3.cyclicExecution := TRUE;
   BenchUut3.trigger := FALSE;
   BenchUut3.value := LREAL#94.0;
   BenchUut3.windowSize := INT#100;
   BenchUut3.reset := FALSE;
   TraceIn_cyclicExecution[123] := BenchUut3.cyclicExecution;
   TraceIn_trigger[123] := BenchUut3.trigger;
   TraceIn_value[123] := BenchUut3.value;
   TraceIn_windowSize[123] := BenchUut3.windowSize;
   TraceIn_reset[123] := BenchUut3.reset;
   BenchUut3();
   TraceOut_average[123] := BenchUut3.average;
   TraceOut_windowSizeReached[123] := BenchUut3.windowSizeReached;
   TraceOut_error[123] := BenchUut3.error;
   TraceOut_status[123] := BenchUut3.status;
   BenchCalls := BenchCalls + 1;
 124:
   BenchUut3.cyclicExecution := TRUE;
   BenchUut3.trigger := FALSE;
   BenchUut3.value := LREAL#95.0;
   BenchUut3.windowSize := INT#100;
   BenchUut3.reset := FALSE;
   TraceIn_cyclicExecution[124] := BenchUut3.cyclicExecution;
   TraceIn_trigger[124] := BenchUut3.trigger;
   TraceIn_value[124] := BenchUut3.value;
   TraceIn_windowSize[124] := BenchUut3.windowSize;
   TraceIn_reset[124] := BenchUut3.reset;
   BenchUut3();
   TraceOut_average[124] := BenchUut3.average;
   TraceOut_windowSizeReached[124] := BenchUut3.windowSizeReached;
   TraceOut_error[124] := BenchUut3.error;
   TraceOut_status[124] := BenchUut3.status;
   BenchCalls := BenchCalls + 1;
 125:
   BenchUut3.cyclicExecution := TRUE;
   BenchUut3.trigger := FALSE;
   BenchUut3.value := LREAL#96.0;
   BenchUut3.windowSize := INT#100;
   BenchUut3.reset := FALSE;
   TraceIn_cyclicExecution[125] := BenchUut3.cyclicExecution;
   TraceIn_trigger[125] := BenchUut3.trigger;
   TraceIn_value[125] := BenchUut3.value;
   TraceIn_windowSize[125] := BenchUut3.windowSize;
   TraceIn_reset[125] := BenchUut3.reset;
   BenchUut3();
   TraceOut_average[125] := BenchUut3.average;
   TraceOut_windowSizeReached[125] := BenchUut3.windowSizeReached;
   TraceOut_error[125] := BenchUut3.error;
   TraceOut_status[125] := BenchUut3.status;
   BenchCalls := BenchCalls + 1;
 126:
   BenchUut3.cyclicExecution := TRUE;
   BenchUut3.trigger := FALSE;
   BenchUut3.value := LREAL#97.0;
   BenchUut3.windowSize := INT#100;
   BenchUut3.reset := FALSE;
   TraceIn_cyclicExecution[126] := BenchUut3.cyclicExecution;
   TraceIn_trigger[126] := BenchUut3.trigger;
   TraceIn_value[126] := BenchUut3.value;
   TraceIn_windowSize[126] := BenchUut3.windowSize;
   TraceIn_reset[126] := BenchUut3.reset;
   BenchUut3();
   TraceOut_average[126] := BenchUut3.average;
   TraceOut_windowSizeReached[126] := BenchUut3.windowSizeReached;
   TraceOut_error[126] := BenchUut3.error;
   TraceOut_status[126] := BenchUut3.status;
   BenchCalls := BenchCalls + 1;
 127:
   BenchUut3.cyclicExecution := TRUE;
   BenchUut3.trigger := FALSE;
   BenchUut3.value := LREAL#98.0;
   BenchUut3.windowSize := INT#100;
   BenchUut3.reset := FALSE;
   TraceIn_cyclicExecution[127] := BenchUut3.cyclicExecution;
   TraceIn_trigger[127] := BenchUut3.trigger;
   TraceIn_value[127] := BenchUut3.value;
   TraceIn_windowSize[127] := BenchUut3.windowSize;
   TraceIn_reset[127] := BenchUut3.reset;
   BenchUut3();
   TraceOut_average[127] := BenchUut3.average;
   TraceOut_windowSizeReached[127] := BenchUut3.windowSizeReached;
   TraceOut_error[127] := BenchUut3.error;
   TraceOut_status[127] := BenchUut3.status;
   BenchCalls := BenchCalls + 1;
 128:
   BenchUut3.cyclicExecution := TRUE;
   BenchUut3.trigger := FALSE;
   BenchUut3.value := LREAL#99.0;
   BenchUut3.windowSize := INT#100;
   BenchUut3.reset := FALSE;
   TraceIn_cyclicExecution[128] := BenchUut3.cyclicExecution;
   TraceIn_trigger[128] := BenchUut3.trigger;
   TraceIn_value[128] := BenchUut3.value;
   TraceIn_windowSize[128] := BenchUut3.windowSize;
   TraceIn_reset[128] := BenchUut3.reset;
   BenchUut3();
   TraceOut_average[128] := BenchUut3.average;
   TraceOut_windowSizeReached[128] := BenchUut3.windowSizeReached;
   TraceOut_error[128] := BenchUut3.error;
   TraceOut_status[128] := BenchUut3.status;
   BenchCalls := BenchCalls + 1;
 129:
   BenchUut3.cyclicExecution := TRUE;
   BenchUut3.trigger := FALSE;
   BenchUut3.value := LREAL#100.0;
   BenchUut3.windowSize := INT#100;
   BenchUut3.reset := FALSE;
   TraceIn_cyclicExecution[129] := BenchUut3.cyclicExecution;
   TraceIn_trigger[129] := BenchUut3.trigger;
   TraceIn_value[129] := BenchUut3.value;
   TraceIn_windowSize[129] := BenchUut3.windowSize;
   TraceIn_reset[129] := BenchUut3.reset;
   BenchUut3();
   TraceOut_average[129] := BenchUut3.average;
   TraceOut_windowSizeReached[129] := BenchUut3.windowSizeReached;
   TraceOut_error[129] := BenchUut3.error;
   TraceOut_status[129] := BenchUut3.status;
   BenchCalls := BenchCalls + 1;
 130:
   BenchUut3.cyclicExecution := TRUE;
   BenchUut3.trigger := FALSE;
   BenchUut3.value := LREAL#101.0;
   BenchUut3.windowSize := INT#100;
   BenchUut3.reset := FALSE;
   TraceIn_cyclicExecution[130] := BenchUut3.cyclicExecution;
   TraceIn_trigger[130] := BenchUut3.trigger;
   TraceIn_value[130] := BenchUut3.value;
   TraceIn_windowSize[130] := BenchUut3.windowSize;
   TraceIn_reset[130] := BenchUut3.reset;
   BenchUut3();
   TraceOut_average[130] := BenchUut3.average;
   TraceOut_windowSizeReached[130] := BenchUut3.windowSizeReached;
   TraceOut_error[130] := BenchUut3.error;
   TraceOut_status[130] := BenchUut3.status;
   BenchCalls := BenchCalls + 1;
 131:
   BenchUut4.cyclicExecution := TRUE;
   BenchUut4.trigger := FALSE;
   BenchUut4.value := LREAL#3.0;
   BenchUut4.windowSize := INT#100;
   BenchUut4.reset := FALSE;
   TraceIn_cyclicExecution[131] := BenchUut4.cyclicExecution;
   TraceIn_trigger[131] := BenchUut4.trigger;
   TraceIn_value[131] := BenchUut4.value;
   TraceIn_windowSize[131] := BenchUut4.windowSize;
   TraceIn_reset[131] := BenchUut4.reset;
   BenchUut4();
   TraceOut_average[131] := BenchUut4.average;
   TraceOut_windowSizeReached[131] := BenchUut4.windowSizeReached;
   TraceOut_error[131] := BenchUut4.error;
   TraceOut_status[131] := BenchUut4.status;
   BenchCalls := BenchCalls + 1;
 132:
   BenchUut5.cyclicExecution := TRUE;
   BenchUut5.trigger := TRUE;
   BenchUut5.value := LREAL#0.0;
   BenchUut5.windowSize := INT#100;
   BenchUut5.reset := FALSE;
   TraceIn_cyclicExecution[132] := BenchUut5.cyclicExecution;
   TraceIn_trigger[132] := BenchUut5.trigger;
   TraceIn_value[132] := BenchUut5.value;
   TraceIn_windowSize[132] := BenchUut5.windowSize;
   TraceIn_reset[132] := BenchUut5.reset;
   BenchUut5();
   TraceOut_average[132] := BenchUut5.average;
   TraceOut_windowSizeReached[132] := BenchUut5.windowSizeReached;
   TraceOut_error[132] := BenchUut5.error;
   TraceOut_status[132] := BenchUut5.status;
   BenchCalls := BenchCalls + 1;
 133:
   BenchUut5.cyclicExecution := TRUE;
   BenchUut5.trigger := TRUE;
   BenchUut5.value := LREAL#1.0;
   BenchUut5.windowSize := INT#100;
   BenchUut5.reset := FALSE;
   TraceIn_cyclicExecution[133] := BenchUut5.cyclicExecution;
   TraceIn_trigger[133] := BenchUut5.trigger;
   TraceIn_value[133] := BenchUut5.value;
   TraceIn_windowSize[133] := BenchUut5.windowSize;
   TraceIn_reset[133] := BenchUut5.reset;
   BenchUut5();
   TraceOut_average[133] := BenchUut5.average;
   TraceOut_windowSizeReached[133] := BenchUut5.windowSizeReached;
   TraceOut_error[133] := BenchUut5.error;
   TraceOut_status[133] := BenchUut5.status;
   BenchCalls := BenchCalls + 1;
 134:
   BenchUut5.cyclicExecution := TRUE;
   BenchUut5.trigger := TRUE;
   BenchUut5.value := LREAL#2.0;
   BenchUut5.windowSize := INT#100;
   BenchUut5.reset := FALSE;
   TraceIn_cyclicExecution[134] := BenchUut5.cyclicExecution;
   TraceIn_trigger[134] := BenchUut5.trigger;
   TraceIn_value[134] := BenchUut5.value;
   TraceIn_windowSize[134] := BenchUut5.windowSize;
   TraceIn_reset[134] := BenchUut5.reset;
   BenchUut5();
   TraceOut_average[134] := BenchUut5.average;
   TraceOut_windowSizeReached[134] := BenchUut5.windowSizeReached;
   TraceOut_error[134] := BenchUut5.error;
   TraceOut_status[134] := BenchUut5.status;
   BenchCalls := BenchCalls + 1;
 135:
   BenchUut5.cyclicExecution := TRUE;
   BenchUut5.trigger := TRUE;
   BenchUut5.value := LREAL#3.0;
   BenchUut5.windowSize := INT#100;
   BenchUut5.reset := FALSE;
   TraceIn_cyclicExecution[135] := BenchUut5.cyclicExecution;
   TraceIn_trigger[135] := BenchUut5.trigger;
   TraceIn_value[135] := BenchUut5.value;
   TraceIn_windowSize[135] := BenchUut5.windowSize;
   TraceIn_reset[135] := BenchUut5.reset;
   BenchUut5();
   TraceOut_average[135] := BenchUut5.average;
   TraceOut_windowSizeReached[135] := BenchUut5.windowSizeReached;
   TraceOut_error[135] := BenchUut5.error;
   TraceOut_status[135] := BenchUut5.status;
   BenchCalls := BenchCalls + 1;
 136:
   BenchUut5.cyclicExecution := TRUE;
   BenchUut5.trigger := TRUE;
   BenchUut5.value := LREAL#4.0;
   BenchUut5.windowSize := INT#100;
   BenchUut5.reset := FALSE;
   TraceIn_cyclicExecution[136] := BenchUut5.cyclicExecution;
   TraceIn_trigger[136] := BenchUut5.trigger;
   TraceIn_value[136] := BenchUut5.value;
   TraceIn_windowSize[136] := BenchUut5.windowSize;
   TraceIn_reset[136] := BenchUut5.reset;
   BenchUut5();
   TraceOut_average[136] := BenchUut5.average;
   TraceOut_windowSizeReached[136] := BenchUut5.windowSizeReached;
   TraceOut_error[136] := BenchUut5.error;
   TraceOut_status[136] := BenchUut5.status;
   BenchCalls := BenchCalls + 1;
 137:
   BenchUut5.cyclicExecution := TRUE;
   BenchUut5.trigger := TRUE;
   BenchUut5.value := LREAL#5.0;
   BenchUut5.windowSize := INT#100;
   BenchUut5.reset := FALSE;
   TraceIn_cyclicExecution[137] := BenchUut5.cyclicExecution;
   TraceIn_trigger[137] := BenchUut5.trigger;
   TraceIn_value[137] := BenchUut5.value;
   TraceIn_windowSize[137] := BenchUut5.windowSize;
   TraceIn_reset[137] := BenchUut5.reset;
   BenchUut5();
   TraceOut_average[137] := BenchUut5.average;
   TraceOut_windowSizeReached[137] := BenchUut5.windowSizeReached;
   TraceOut_error[137] := BenchUut5.error;
   TraceOut_status[137] := BenchUut5.status;
   BenchCalls := BenchCalls + 1;
 138:
   BenchUut5.cyclicExecution := TRUE;
   BenchUut5.trigger := TRUE;
   BenchUut5.value := LREAL#6.0;
   BenchUut5.windowSize := INT#100;
   BenchUut5.reset := FALSE;
   TraceIn_cyclicExecution[138] := BenchUut5.cyclicExecution;
   TraceIn_trigger[138] := BenchUut5.trigger;
   TraceIn_value[138] := BenchUut5.value;
   TraceIn_windowSize[138] := BenchUut5.windowSize;
   TraceIn_reset[138] := BenchUut5.reset;
   BenchUut5();
   TraceOut_average[138] := BenchUut5.average;
   TraceOut_windowSizeReached[138] := BenchUut5.windowSizeReached;
   TraceOut_error[138] := BenchUut5.error;
   TraceOut_status[138] := BenchUut5.status;
   BenchCalls := BenchCalls + 1;
 139:
   BenchUut5.cyclicExecution := TRUE;
   BenchUut5.trigger := TRUE;
   BenchUut5.value := LREAL#7.0;
   BenchUut5.windowSize := INT#100;
   BenchUut5.reset := FALSE;
   TraceIn_cyclicExecution[139] := BenchUut5.cyclicExecution;
   TraceIn_trigger[139] := BenchUut5.trigger;
   TraceIn_value[139] := BenchUut5.value;
   TraceIn_windowSize[139] := BenchUut5.windowSize;
   TraceIn_reset[139] := BenchUut5.reset;
   BenchUut5();
   TraceOut_average[139] := BenchUut5.average;
   TraceOut_windowSizeReached[139] := BenchUut5.windowSizeReached;
   TraceOut_error[139] := BenchUut5.error;
   TraceOut_status[139] := BenchUut5.status;
   BenchCalls := BenchCalls + 1;
 140:
   BenchUut5.cyclicExecution := TRUE;
   BenchUut5.trigger := TRUE;
   BenchUut5.value := LREAL#8.0;
   BenchUut5.windowSize := INT#100;
   BenchUut5.reset := FALSE;
   TraceIn_cyclicExecution[140] := BenchUut5.cyclicExecution;
   TraceIn_trigger[140] := BenchUut5.trigger;
   TraceIn_value[140] := BenchUut5.value;
   TraceIn_windowSize[140] := BenchUut5.windowSize;
   TraceIn_reset[140] := BenchUut5.reset;
   BenchUut5();
   TraceOut_average[140] := BenchUut5.average;
   TraceOut_windowSizeReached[140] := BenchUut5.windowSizeReached;
   TraceOut_error[140] := BenchUut5.error;
   TraceOut_status[140] := BenchUut5.status;
   BenchCalls := BenchCalls + 1;
 141:
   BenchUut5.cyclicExecution := TRUE;
   BenchUut5.trigger := TRUE;
   BenchUut5.value := LREAL#9.0;
   BenchUut5.windowSize := INT#100;
   BenchUut5.reset := FALSE;
   TraceIn_cyclicExecution[141] := BenchUut5.cyclicExecution;
   TraceIn_trigger[141] := BenchUut5.trigger;
   TraceIn_value[141] := BenchUut5.value;
   TraceIn_windowSize[141] := BenchUut5.windowSize;
   TraceIn_reset[141] := BenchUut5.reset;
   BenchUut5();
   TraceOut_average[141] := BenchUut5.average;
   TraceOut_windowSizeReached[141] := BenchUut5.windowSizeReached;
   TraceOut_error[141] := BenchUut5.error;
   TraceOut_status[141] := BenchUut5.status;
   BenchCalls := BenchCalls + 1;
 142:
   BenchUut5.cyclicExecution := TRUE;
   BenchUut5.trigger := TRUE;
   BenchUut5.value := LREAL#10.0;
   BenchUut5.windowSize := INT#100;
   BenchUut5.reset := FALSE;
   TraceIn_cyclicExecution[142] := BenchUut5.cyclicExecution;
   TraceIn_trigger[142] := BenchUut5.trigger;
   TraceIn_value[142] := BenchUut5.value;
   TraceIn_windowSize[142] := BenchUut5.windowSize;
   TraceIn_reset[142] := BenchUut5.reset;
   BenchUut5();
   TraceOut_average[142] := BenchUut5.average;
   TraceOut_windowSizeReached[142] := BenchUut5.windowSizeReached;
   TraceOut_error[142] := BenchUut5.error;
   TraceOut_status[142] := BenchUut5.status;
   BenchCalls := BenchCalls + 1;
 143:
   BenchUut5.cyclicExecution := TRUE;
   BenchUut5.trigger := TRUE;
   BenchUut5.value := LREAL#11.0;
   BenchUut5.windowSize := INT#100;
   BenchUut5.reset := FALSE;
   TraceIn_cyclicExecution[143] := BenchUut5.cyclicExecution;
   TraceIn_trigger[143] := BenchUut5.trigger;
   TraceIn_value[143] := BenchUut5.value;
   TraceIn_windowSize[143] := BenchUut5.windowSize;
   TraceIn_reset[143] := BenchUut5.reset;
   BenchUut5();
   TraceOut_average[143] := BenchUut5.average;
   TraceOut_windowSizeReached[143] := BenchUut5.windowSizeReached;
   TraceOut_error[143] := BenchUut5.error;
   TraceOut_status[143] := BenchUut5.status;
   BenchCalls := BenchCalls + 1;
 144:
   BenchUut5.cyclicExecution := TRUE;
   BenchUut5.trigger := TRUE;
   BenchUut5.value := LREAL#12.0;
   BenchUut5.windowSize := INT#100;
   BenchUut5.reset := FALSE;
   TraceIn_cyclicExecution[144] := BenchUut5.cyclicExecution;
   TraceIn_trigger[144] := BenchUut5.trigger;
   TraceIn_value[144] := BenchUut5.value;
   TraceIn_windowSize[144] := BenchUut5.windowSize;
   TraceIn_reset[144] := BenchUut5.reset;
   BenchUut5();
   TraceOut_average[144] := BenchUut5.average;
   TraceOut_windowSizeReached[144] := BenchUut5.windowSizeReached;
   TraceOut_error[144] := BenchUut5.error;
   TraceOut_status[144] := BenchUut5.status;
   BenchCalls := BenchCalls + 1;
 145:
   BenchUut5.cyclicExecution := TRUE;
   BenchUut5.trigger := TRUE;
   BenchUut5.value := LREAL#13.0;
   BenchUut5.windowSize := INT#100;
   BenchUut5.reset := FALSE;
   TraceIn_cyclicExecution[145] := BenchUut5.cyclicExecution;
   TraceIn_trigger[145] := BenchUut5.trigger;
   TraceIn_value[145] := BenchUut5.value;
   TraceIn_windowSize[145] := BenchUut5.windowSize;
   TraceIn_reset[145] := BenchUut5.reset;
   BenchUut5();
   TraceOut_average[145] := BenchUut5.average;
   TraceOut_windowSizeReached[145] := BenchUut5.windowSizeReached;
   TraceOut_error[145] := BenchUut5.error;
   TraceOut_status[145] := BenchUut5.status;
   BenchCalls := BenchCalls + 1;
 146:
   BenchUut5.cyclicExecution := TRUE;
   BenchUut5.trigger := TRUE;
   BenchUut5.value := LREAL#14.0;
   BenchUut5.windowSize := INT#100;
   BenchUut5.reset := FALSE;
   TraceIn_cyclicExecution[146] := BenchUut5.cyclicExecution;
   TraceIn_trigger[146] := BenchUut5.trigger;
   TraceIn_value[146] := BenchUut5.value;
   TraceIn_windowSize[146] := BenchUut5.windowSize;
   TraceIn_reset[146] := BenchUut5.reset;
   BenchUut5();
   TraceOut_average[146] := BenchUut5.average;
   TraceOut_windowSizeReached[146] := BenchUut5.windowSizeReached;
   TraceOut_error[146] := BenchUut5.error;
   TraceOut_status[146] := BenchUut5.status;
   BenchCalls := BenchCalls + 1;
 147:
   BenchUut5.cyclicExecution := TRUE;
   BenchUut5.trigger := TRUE;
   BenchUut5.value := LREAL#15.0;
   BenchUut5.windowSize := INT#100;
   BenchUut5.reset := FALSE;
   TraceIn_cyclicExecution[147] := BenchUut5.cyclicExecution;
   TraceIn_trigger[147] := BenchUut5.trigger;
   TraceIn_value[147] := BenchUut5.value;
   TraceIn_windowSize[147] := BenchUut5.windowSize;
   TraceIn_reset[147] := BenchUut5.reset;
   BenchUut5();
   TraceOut_average[147] := BenchUut5.average;
   TraceOut_windowSizeReached[147] := BenchUut5.windowSizeReached;
   TraceOut_error[147] := BenchUut5.error;
   TraceOut_status[147] := BenchUut5.status;
   BenchCalls := BenchCalls + 1;
 148:
   BenchUut5.cyclicExecution := TRUE;
   BenchUut5.trigger := TRUE;
   BenchUut5.value := LREAL#16.0;
   BenchUut5.windowSize := INT#100;
   BenchUut5.reset := FALSE;
   TraceIn_cyclicExecution[148] := BenchUut5.cyclicExecution;
   TraceIn_trigger[148] := BenchUut5.trigger;
   TraceIn_value[148] := BenchUut5.value;
   TraceIn_windowSize[148] := BenchUut5.windowSize;
   TraceIn_reset[148] := BenchUut5.reset;
   BenchUut5();
   TraceOut_average[148] := BenchUut5.average;
   TraceOut_windowSizeReached[148] := BenchUut5.windowSizeReached;
   TraceOut_error[148] := BenchUut5.error;
   TraceOut_status[148] := BenchUut5.status;
   BenchCalls := BenchCalls + 1;
 149:
   BenchUut5.cyclicExecution := TRUE;
   BenchUut5.trigger := TRUE;
   BenchUut5.value := LREAL#17.0;
   BenchUut5.windowSize := INT#100;
   BenchUut5.reset := FALSE;
   TraceIn_cyclicExecution[149] := BenchUut5.cyclicExecution;
   TraceIn_trigger[149] := BenchUut5.trigger;
   TraceIn_value[149] := BenchUut5.value;
   TraceIn_windowSize[149] := BenchUut5.windowSize;
   TraceIn_reset[149] := BenchUut5.reset;
   BenchUut5();
   TraceOut_average[149] := BenchUut5.average;
   TraceOut_windowSizeReached[149] := BenchUut5.windowSizeReached;
   TraceOut_error[149] := BenchUut5.error;
   TraceOut_status[149] := BenchUut5.status;
   BenchCalls := BenchCalls + 1;
 150:
   BenchUut5.cyclicExecution := TRUE;
   BenchUut5.trigger := TRUE;
   BenchUut5.value := LREAL#18.0;
   BenchUut5.windowSize := INT#100;
   BenchUut5.reset := FALSE;
   TraceIn_cyclicExecution[150] := BenchUut5.cyclicExecution;
   TraceIn_trigger[150] := BenchUut5.trigger;
   TraceIn_value[150] := BenchUut5.value;
   TraceIn_windowSize[150] := BenchUut5.windowSize;
   TraceIn_reset[150] := BenchUut5.reset;
   BenchUut5();
   TraceOut_average[150] := BenchUut5.average;
   TraceOut_windowSizeReached[150] := BenchUut5.windowSizeReached;
   TraceOut_error[150] := BenchUut5.error;
   TraceOut_status[150] := BenchUut5.status;
   BenchCalls := BenchCalls + 1;
 151:
   BenchUut5.cyclicExecution := TRUE;
   BenchUut5.trigger := TRUE;
   BenchUut5.value := LREAL#19.0;
   BenchUut5.windowSize := INT#100;
   BenchUut5.reset := FALSE;
   TraceIn_cyclicExecution[151] := BenchUut5.cyclicExecution;
   TraceIn_trigger[151] := BenchUut5.trigger;
   TraceIn_value[151] := BenchUut5.value;
   TraceIn_windowSize[151] := BenchUut5.windowSize;
   TraceIn_reset[151] := BenchUut5.reset;
   BenchUut5();
   TraceOut_average[151] := BenchUut5.average;
   TraceOut_windowSizeReached[151] := BenchUut5.windowSizeReached;
   TraceOut_error[151] := BenchUut5.error;
   TraceOut_status[151] := BenchUut5.status;
   BenchCalls := BenchCalls + 1;
 152:
   BenchUut5.cyclicExecution := TRUE;
   BenchUut5.trigger := TRUE;
   BenchUut5.value := LREAL#20.0;
   BenchUut5.windowSize := INT#100;
   BenchUut5.reset := FALSE;
   TraceIn_cyclicExecution[152] := BenchUut5.cyclicExecution;
   TraceIn_trigger[152] := BenchUut5.trigger;
   TraceIn_value[152] := BenchUut5.value;
   TraceIn_windowSize[152] := BenchUut5.windowSize;
   TraceIn_reset[152] := BenchUut5.reset;
   BenchUut5();
   TraceOut_average[152] := BenchUut5.average;
   TraceOut_windowSizeReached[152] := BenchUut5.windowSizeReached;
   TraceOut_error[152] := BenchUut5.error;
   TraceOut_status[152] := BenchUut5.status;
   BenchCalls := BenchCalls + 1;
 153:
   BenchUut5.cyclicExecution := TRUE;
   BenchUut5.trigger := TRUE;
   BenchUut5.value := LREAL#21.0;
   BenchUut5.windowSize := INT#100;
   BenchUut5.reset := FALSE;
   TraceIn_cyclicExecution[153] := BenchUut5.cyclicExecution;
   TraceIn_trigger[153] := BenchUut5.trigger;
   TraceIn_value[153] := BenchUut5.value;
   TraceIn_windowSize[153] := BenchUut5.windowSize;
   TraceIn_reset[153] := BenchUut5.reset;
   BenchUut5();
   TraceOut_average[153] := BenchUut5.average;
   TraceOut_windowSizeReached[153] := BenchUut5.windowSizeReached;
   TraceOut_error[153] := BenchUut5.error;
   TraceOut_status[153] := BenchUut5.status;
   BenchCalls := BenchCalls + 1;
 154:
   BenchUut5.cyclicExecution := TRUE;
   BenchUut5.trigger := TRUE;
   BenchUut5.value := LREAL#22.0;
   BenchUut5.windowSize := INT#100;
   BenchUut5.reset := FALSE;
   TraceIn_cyclicExecution[154] := BenchUut5.cyclicExecution;
   TraceIn_trigger[154] := BenchUut5.trigger;
   TraceIn_value[154] := BenchUut5.value;
   TraceIn_windowSize[154] := BenchUut5.windowSize;
   TraceIn_reset[154] := BenchUut5.reset;
   BenchUut5();
   TraceOut_average[154] := BenchUut5.average;
   TraceOut_windowSizeReached[154] := BenchUut5.windowSizeReached;
   TraceOut_error[154] := BenchUut5.error;
   TraceOut_status[154] := BenchUut5.status;
   BenchCalls := BenchCalls + 1;
 155:
   BenchUut5.cyclicExecution := TRUE;
   BenchUut5.trigger := TRUE;
   BenchUut5.value := LREAL#23.0;
   BenchUut5.windowSize := INT#100;
   BenchUut5.reset := FALSE;
   TraceIn_cyclicExecution[155] := BenchUut5.cyclicExecution;
   TraceIn_trigger[155] := BenchUut5.trigger;
   TraceIn_value[155] := BenchUut5.value;
   TraceIn_windowSize[155] := BenchUut5.windowSize;
   TraceIn_reset[155] := BenchUut5.reset;
   BenchUut5();
   TraceOut_average[155] := BenchUut5.average;
   TraceOut_windowSizeReached[155] := BenchUut5.windowSizeReached;
   TraceOut_error[155] := BenchUut5.error;
   TraceOut_status[155] := BenchUut5.status;
   BenchCalls := BenchCalls + 1;
 156:
   BenchUut5.cyclicExecution := TRUE;
   BenchUut5.trigger := TRUE;
   BenchUut5.value := LREAL#24.0;
   BenchUut5.windowSize := INT#100;
   BenchUut5.reset := FALSE;
   TraceIn_cyclicExecution[156] := BenchUut5.cyclicExecution;
   TraceIn_trigger[156] := BenchUut5.trigger;
   TraceIn_value[156] := BenchUut5.value;
   TraceIn_windowSize[156] := BenchUut5.windowSize;
   TraceIn_reset[156] := BenchUut5.reset;
   BenchUut5();
   TraceOut_average[156] := BenchUut5.average;
   TraceOut_windowSizeReached[156] := BenchUut5.windowSizeReached;
   TraceOut_error[156] := BenchUut5.error;
   TraceOut_status[156] := BenchUut5.status;
   BenchCalls := BenchCalls + 1;
 157:
   BenchUut5.cyclicExecution := TRUE;
   BenchUut5.trigger := TRUE;
   BenchUut5.value := LREAL#25.0;
   BenchUut5.windowSize := INT#100;
   BenchUut5.reset := FALSE;
   TraceIn_cyclicExecution[157] := BenchUut5.cyclicExecution;
   TraceIn_trigger[157] := BenchUut5.trigger;
   TraceIn_value[157] := BenchUut5.value;
   TraceIn_windowSize[157] := BenchUut5.windowSize;
   TraceIn_reset[157] := BenchUut5.reset;
   BenchUut5();
   TraceOut_average[157] := BenchUut5.average;
   TraceOut_windowSizeReached[157] := BenchUut5.windowSizeReached;
   TraceOut_error[157] := BenchUut5.error;
   TraceOut_status[157] := BenchUut5.status;
   BenchCalls := BenchCalls + 1;
 158:
   BenchUut5.cyclicExecution := TRUE;
   BenchUut5.trigger := TRUE;
   BenchUut5.value := LREAL#26.0;
   BenchUut5.windowSize := INT#100;
   BenchUut5.reset := FALSE;
   TraceIn_cyclicExecution[158] := BenchUut5.cyclicExecution;
   TraceIn_trigger[158] := BenchUut5.trigger;
   TraceIn_value[158] := BenchUut5.value;
   TraceIn_windowSize[158] := BenchUut5.windowSize;
   TraceIn_reset[158] := BenchUut5.reset;
   BenchUut5();
   TraceOut_average[158] := BenchUut5.average;
   TraceOut_windowSizeReached[158] := BenchUut5.windowSizeReached;
   TraceOut_error[158] := BenchUut5.error;
   TraceOut_status[158] := BenchUut5.status;
   BenchCalls := BenchCalls + 1;
 159:
   BenchUut5.cyclicExecution := TRUE;
   BenchUut5.trigger := TRUE;
   BenchUut5.value := LREAL#27.0;
   BenchUut5.windowSize := INT#100;
   BenchUut5.reset := FALSE;
   TraceIn_cyclicExecution[159] := BenchUut5.cyclicExecution;
   TraceIn_trigger[159] := BenchUut5.trigger;
   TraceIn_value[159] := BenchUut5.value;
   TraceIn_windowSize[159] := BenchUut5.windowSize;
   TraceIn_reset[159] := BenchUut5.reset;
   BenchUut5();
   TraceOut_average[159] := BenchUut5.average;
   TraceOut_windowSizeReached[159] := BenchUut5.windowSizeReached;
   TraceOut_error[159] := BenchUut5.error;
   TraceOut_status[159] := BenchUut5.status;
   BenchCalls := BenchCalls + 1;
 160:
   BenchUut5.cyclicExecution := TRUE;
   BenchUut5.trigger := TRUE;
   BenchUut5.value := LREAL#28.0;
   BenchUut5.windowSize := INT#100;
   BenchUut5.reset := FALSE;
   TraceIn_cyclicExecution[160] := BenchUut5.cyclicExecution;
   TraceIn_trigger[160] := BenchUut5.trigger;
   TraceIn_value[160] := BenchUut5.value;
   TraceIn_windowSize[160] := BenchUut5.windowSize;
   TraceIn_reset[160] := BenchUut5.reset;
   BenchUut5();
   TraceOut_average[160] := BenchUut5.average;
   TraceOut_windowSizeReached[160] := BenchUut5.windowSizeReached;
   TraceOut_error[160] := BenchUut5.error;
   TraceOut_status[160] := BenchUut5.status;
   BenchCalls := BenchCalls + 1;
 161:
   BenchUut5.cyclicExecution := TRUE;
   BenchUut5.trigger := TRUE;
   BenchUut5.value := LREAL#29.0;
   BenchUut5.windowSize := INT#100;
   BenchUut5.reset := FALSE;
   TraceIn_cyclicExecution[161] := BenchUut5.cyclicExecution;
   TraceIn_trigger[161] := BenchUut5.trigger;
   TraceIn_value[161] := BenchUut5.value;
   TraceIn_windowSize[161] := BenchUut5.windowSize;
   TraceIn_reset[161] := BenchUut5.reset;
   BenchUut5();
   TraceOut_average[161] := BenchUut5.average;
   TraceOut_windowSizeReached[161] := BenchUut5.windowSizeReached;
   TraceOut_error[161] := BenchUut5.error;
   TraceOut_status[161] := BenchUut5.status;
   BenchCalls := BenchCalls + 1;
 162:
   BenchUut5.cyclicExecution := TRUE;
   BenchUut5.trigger := TRUE;
   BenchUut5.value := LREAL#30.0;
   BenchUut5.windowSize := INT#100;
   BenchUut5.reset := FALSE;
   TraceIn_cyclicExecution[162] := BenchUut5.cyclicExecution;
   TraceIn_trigger[162] := BenchUut5.trigger;
   TraceIn_value[162] := BenchUut5.value;
   TraceIn_windowSize[162] := BenchUut5.windowSize;
   TraceIn_reset[162] := BenchUut5.reset;
   BenchUut5();
   TraceOut_average[162] := BenchUut5.average;
   TraceOut_windowSizeReached[162] := BenchUut5.windowSizeReached;
   TraceOut_error[162] := BenchUut5.error;
   TraceOut_status[162] := BenchUut5.status;
   BenchCalls := BenchCalls + 1;
 163:
   BenchUut5.cyclicExecution := TRUE;
   BenchUut5.trigger := TRUE;
   BenchUut5.value := LREAL#31.0;
   BenchUut5.windowSize := INT#100;
   BenchUut5.reset := FALSE;
   TraceIn_cyclicExecution[163] := BenchUut5.cyclicExecution;
   TraceIn_trigger[163] := BenchUut5.trigger;
   TraceIn_value[163] := BenchUut5.value;
   TraceIn_windowSize[163] := BenchUut5.windowSize;
   TraceIn_reset[163] := BenchUut5.reset;
   BenchUut5();
   TraceOut_average[163] := BenchUut5.average;
   TraceOut_windowSizeReached[163] := BenchUut5.windowSizeReached;
   TraceOut_error[163] := BenchUut5.error;
   TraceOut_status[163] := BenchUut5.status;
   BenchCalls := BenchCalls + 1;
 164:
   BenchUut5.cyclicExecution := TRUE;
   BenchUut5.trigger := TRUE;
   BenchUut5.value := LREAL#32.0;
   BenchUut5.windowSize := INT#100;
   BenchUut5.reset := FALSE;
   TraceIn_cyclicExecution[164] := BenchUut5.cyclicExecution;
   TraceIn_trigger[164] := BenchUut5.trigger;
   TraceIn_value[164] := BenchUut5.value;
   TraceIn_windowSize[164] := BenchUut5.windowSize;
   TraceIn_reset[164] := BenchUut5.reset;
   BenchUut5();
   TraceOut_average[164] := BenchUut5.average;
   TraceOut_windowSizeReached[164] := BenchUut5.windowSizeReached;
   TraceOut_error[164] := BenchUut5.error;
   TraceOut_status[164] := BenchUut5.status;
   BenchCalls := BenchCalls + 1;
 165:
   BenchUut5.cyclicExecution := TRUE;
   BenchUut5.trigger := TRUE;
   BenchUut5.value := LREAL#33.0;
   BenchUut5.windowSize := INT#100;
   BenchUut5.reset := FALSE;
   TraceIn_cyclicExecution[165] := BenchUut5.cyclicExecution;
   TraceIn_trigger[165] := BenchUut5.trigger;
   TraceIn_value[165] := BenchUut5.value;
   TraceIn_windowSize[165] := BenchUut5.windowSize;
   TraceIn_reset[165] := BenchUut5.reset;
   BenchUut5();
   TraceOut_average[165] := BenchUut5.average;
   TraceOut_windowSizeReached[165] := BenchUut5.windowSizeReached;
   TraceOut_error[165] := BenchUut5.error;
   TraceOut_status[165] := BenchUut5.status;
   BenchCalls := BenchCalls + 1;
 166:
   BenchUut5.cyclicExecution := TRUE;
   BenchUut5.trigger := TRUE;
   BenchUut5.value := LREAL#34.0;
   BenchUut5.windowSize := INT#100;
   BenchUut5.reset := FALSE;
   TraceIn_cyclicExecution[166] := BenchUut5.cyclicExecution;
   TraceIn_trigger[166] := BenchUut5.trigger;
   TraceIn_value[166] := BenchUut5.value;
   TraceIn_windowSize[166] := BenchUut5.windowSize;
   TraceIn_reset[166] := BenchUut5.reset;
   BenchUut5();
   TraceOut_average[166] := BenchUut5.average;
   TraceOut_windowSizeReached[166] := BenchUut5.windowSizeReached;
   TraceOut_error[166] := BenchUut5.error;
   TraceOut_status[166] := BenchUut5.status;
   BenchCalls := BenchCalls + 1;
 167:
   BenchUut5.cyclicExecution := TRUE;
   BenchUut5.trigger := TRUE;
   BenchUut5.value := LREAL#35.0;
   BenchUut5.windowSize := INT#100;
   BenchUut5.reset := FALSE;
   TraceIn_cyclicExecution[167] := BenchUut5.cyclicExecution;
   TraceIn_trigger[167] := BenchUut5.trigger;
   TraceIn_value[167] := BenchUut5.value;
   TraceIn_windowSize[167] := BenchUut5.windowSize;
   TraceIn_reset[167] := BenchUut5.reset;
   BenchUut5();
   TraceOut_average[167] := BenchUut5.average;
   TraceOut_windowSizeReached[167] := BenchUut5.windowSizeReached;
   TraceOut_error[167] := BenchUut5.error;
   TraceOut_status[167] := BenchUut5.status;
   BenchCalls := BenchCalls + 1;
 168:
   BenchUut5.cyclicExecution := TRUE;
   BenchUut5.trigger := TRUE;
   BenchUut5.value := LREAL#36.0;
   BenchUut5.windowSize := INT#100;
   BenchUut5.reset := FALSE;
   TraceIn_cyclicExecution[168] := BenchUut5.cyclicExecution;
   TraceIn_trigger[168] := BenchUut5.trigger;
   TraceIn_value[168] := BenchUut5.value;
   TraceIn_windowSize[168] := BenchUut5.windowSize;
   TraceIn_reset[168] := BenchUut5.reset;
   BenchUut5();
   TraceOut_average[168] := BenchUut5.average;
   TraceOut_windowSizeReached[168] := BenchUut5.windowSizeReached;
   TraceOut_error[168] := BenchUut5.error;
   TraceOut_status[168] := BenchUut5.status;
   BenchCalls := BenchCalls + 1;
 169:
   BenchUut5.cyclicExecution := TRUE;
   BenchUut5.trigger := TRUE;
   BenchUut5.value := LREAL#37.0;
   BenchUut5.windowSize := INT#100;
   BenchUut5.reset := FALSE;
   TraceIn_cyclicExecution[169] := BenchUut5.cyclicExecution;
   TraceIn_trigger[169] := BenchUut5.trigger;
   TraceIn_value[169] := BenchUut5.value;
   TraceIn_windowSize[169] := BenchUut5.windowSize;
   TraceIn_reset[169] := BenchUut5.reset;
   BenchUut5();
   TraceOut_average[169] := BenchUut5.average;
   TraceOut_windowSizeReached[169] := BenchUut5.windowSizeReached;
   TraceOut_error[169] := BenchUut5.error;
   TraceOut_status[169] := BenchUut5.status;
   BenchCalls := BenchCalls + 1;
 170:
   BenchUut5.cyclicExecution := TRUE;
   BenchUut5.trigger := TRUE;
   BenchUut5.value := LREAL#38.0;
   BenchUut5.windowSize := INT#100;
   BenchUut5.reset := FALSE;
   TraceIn_cyclicExecution[170] := BenchUut5.cyclicExecution;
   TraceIn_trigger[170] := BenchUut5.trigger;
   TraceIn_value[170] := BenchUut5.value;
   TraceIn_windowSize[170] := BenchUut5.windowSize;
   TraceIn_reset[170] := BenchUut5.reset;
   BenchUut5();
   TraceOut_average[170] := BenchUut5.average;
   TraceOut_windowSizeReached[170] := BenchUut5.windowSizeReached;
   TraceOut_error[170] := BenchUut5.error;
   TraceOut_status[170] := BenchUut5.status;
   BenchCalls := BenchCalls + 1;
 171:
   BenchUut5.cyclicExecution := TRUE;
   BenchUut5.trigger := TRUE;
   BenchUut5.value := LREAL#39.0;
   BenchUut5.windowSize := INT#100;
   BenchUut5.reset := FALSE;
   TraceIn_cyclicExecution[171] := BenchUut5.cyclicExecution;
   TraceIn_trigger[171] := BenchUut5.trigger;
   TraceIn_value[171] := BenchUut5.value;
   TraceIn_windowSize[171] := BenchUut5.windowSize;
   TraceIn_reset[171] := BenchUut5.reset;
   BenchUut5();
   TraceOut_average[171] := BenchUut5.average;
   TraceOut_windowSizeReached[171] := BenchUut5.windowSizeReached;
   TraceOut_error[171] := BenchUut5.error;
   TraceOut_status[171] := BenchUut5.status;
   BenchCalls := BenchCalls + 1;
 172:
   BenchUut5.cyclicExecution := TRUE;
   BenchUut5.trigger := TRUE;
   BenchUut5.value := LREAL#40.0;
   BenchUut5.windowSize := INT#100;
   BenchUut5.reset := FALSE;
   TraceIn_cyclicExecution[172] := BenchUut5.cyclicExecution;
   TraceIn_trigger[172] := BenchUut5.trigger;
   TraceIn_value[172] := BenchUut5.value;
   TraceIn_windowSize[172] := BenchUut5.windowSize;
   TraceIn_reset[172] := BenchUut5.reset;
   BenchUut5();
   TraceOut_average[172] := BenchUut5.average;
   TraceOut_windowSizeReached[172] := BenchUut5.windowSizeReached;
   TraceOut_error[172] := BenchUut5.error;
   TraceOut_status[172] := BenchUut5.status;
   BenchCalls := BenchCalls + 1;
 173:
   BenchUut5.cyclicExecution := TRUE;
   BenchUut5.trigger := TRUE;
   BenchUut5.value := LREAL#41.0;
   BenchUut5.windowSize := INT#100;
   BenchUut5.reset := FALSE;
   TraceIn_cyclicExecution[173] := BenchUut5.cyclicExecution;
   TraceIn_trigger[173] := BenchUut5.trigger;
   TraceIn_value[173] := BenchUut5.value;
   TraceIn_windowSize[173] := BenchUut5.windowSize;
   TraceIn_reset[173] := BenchUut5.reset;
   BenchUut5();
   TraceOut_average[173] := BenchUut5.average;
   TraceOut_windowSizeReached[173] := BenchUut5.windowSizeReached;
   TraceOut_error[173] := BenchUut5.error;
   TraceOut_status[173] := BenchUut5.status;
   BenchCalls := BenchCalls + 1;
 174:
   BenchUut5.cyclicExecution := TRUE;
   BenchUut5.trigger := TRUE;
   BenchUut5.value := LREAL#42.0;
   BenchUut5.windowSize := INT#100;
   BenchUut5.reset := FALSE;
   TraceIn_cyclicExecution[174] := BenchUut5.cyclicExecution;
   TraceIn_trigger[174] := BenchUut5.trigger;
   TraceIn_value[174] := BenchUut5.value;
   TraceIn_windowSize[174] := BenchUut5.windowSize;
   TraceIn_reset[174] := BenchUut5.reset;
   BenchUut5();
   TraceOut_average[174] := BenchUut5.average;
   TraceOut_windowSizeReached[174] := BenchUut5.windowSizeReached;
   TraceOut_error[174] := BenchUut5.error;
   TraceOut_status[174] := BenchUut5.status;
   BenchCalls := BenchCalls + 1;
 175:
   BenchUut5.cyclicExecution := TRUE;
   BenchUut5.trigger := TRUE;
   BenchUut5.value := LREAL#43.0;
   BenchUut5.windowSize := INT#100;
   BenchUut5.reset := FALSE;
   TraceIn_cyclicExecution[175] := BenchUut5.cyclicExecution;
   TraceIn_trigger[175] := BenchUut5.trigger;
   TraceIn_value[175] := BenchUut5.value;
   TraceIn_windowSize[175] := BenchUut5.windowSize;
   TraceIn_reset[175] := BenchUut5.reset;
   BenchUut5();
   TraceOut_average[175] := BenchUut5.average;
   TraceOut_windowSizeReached[175] := BenchUut5.windowSizeReached;
   TraceOut_error[175] := BenchUut5.error;
   TraceOut_status[175] := BenchUut5.status;
   BenchCalls := BenchCalls + 1;
 176:
   BenchUut5.cyclicExecution := TRUE;
   BenchUut5.trigger := TRUE;
   BenchUut5.value := LREAL#44.0;
   BenchUut5.windowSize := INT#100;
   BenchUut5.reset := FALSE;
   TraceIn_cyclicExecution[176] := BenchUut5.cyclicExecution;
   TraceIn_trigger[176] := BenchUut5.trigger;
   TraceIn_value[176] := BenchUut5.value;
   TraceIn_windowSize[176] := BenchUut5.windowSize;
   TraceIn_reset[176] := BenchUut5.reset;
   BenchUut5();
   TraceOut_average[176] := BenchUut5.average;
   TraceOut_windowSizeReached[176] := BenchUut5.windowSizeReached;
   TraceOut_error[176] := BenchUut5.error;
   TraceOut_status[176] := BenchUut5.status;
   BenchCalls := BenchCalls + 1;
 177:
   BenchUut5.cyclicExecution := TRUE;
   BenchUut5.trigger := TRUE;
   BenchUut5.value := LREAL#45.0;
   BenchUut5.windowSize := INT#100;
   BenchUut5.reset := FALSE;
   TraceIn_cyclicExecution[177] := BenchUut5.cyclicExecution;
   TraceIn_trigger[177] := BenchUut5.trigger;
   TraceIn_value[177] := BenchUut5.value;
   TraceIn_windowSize[177] := BenchUut5.windowSize;
   TraceIn_reset[177] := BenchUut5.reset;
   BenchUut5();
   TraceOut_average[177] := BenchUut5.average;
   TraceOut_windowSizeReached[177] := BenchUut5.windowSizeReached;
   TraceOut_error[177] := BenchUut5.error;
   TraceOut_status[177] := BenchUut5.status;
   BenchCalls := BenchCalls + 1;
 178:
   BenchUut5.cyclicExecution := TRUE;
   BenchUut5.trigger := TRUE;
   BenchUut5.value := LREAL#46.0;
   BenchUut5.windowSize := INT#100;
   BenchUut5.reset := FALSE;
   TraceIn_cyclicExecution[178] := BenchUut5.cyclicExecution;
   TraceIn_trigger[178] := BenchUut5.trigger;
   TraceIn_value[178] := BenchUut5.value;
   TraceIn_windowSize[178] := BenchUut5.windowSize;
   TraceIn_reset[178] := BenchUut5.reset;
   BenchUut5();
   TraceOut_average[178] := BenchUut5.average;
   TraceOut_windowSizeReached[178] := BenchUut5.windowSizeReached;
   TraceOut_error[178] := BenchUut5.error;
   TraceOut_status[178] := BenchUut5.status;
   BenchCalls := BenchCalls + 1;
 179:
   BenchUut5.cyclicExecution := TRUE;
   BenchUut5.trigger := TRUE;
   BenchUut5.value := LREAL#47.0;
   BenchUut5.windowSize := INT#100;
   BenchUut5.reset := FALSE;
   TraceIn_cyclicExecution[179] := BenchUut5.cyclicExecution;
   TraceIn_trigger[179] := BenchUut5.trigger;
   TraceIn_value[179] := BenchUut5.value;
   TraceIn_windowSize[179] := BenchUut5.windowSize;
   TraceIn_reset[179] := BenchUut5.reset;
   BenchUut5();
   TraceOut_average[179] := BenchUut5.average;
   TraceOut_windowSizeReached[179] := BenchUut5.windowSizeReached;
   TraceOut_error[179] := BenchUut5.error;
   TraceOut_status[179] := BenchUut5.status;
   BenchCalls := BenchCalls + 1;
 180:
   BenchUut5.cyclicExecution := TRUE;
   BenchUut5.trigger := TRUE;
   BenchUut5.value := LREAL#48.0;
   BenchUut5.windowSize := INT#100;
   BenchUut5.reset := FALSE;
   TraceIn_cyclicExecution[180] := BenchUut5.cyclicExecution;
   TraceIn_trigger[180] := BenchUut5.trigger;
   TraceIn_value[180] := BenchUut5.value;
   TraceIn_windowSize[180] := BenchUut5.windowSize;
   TraceIn_reset[180] := BenchUut5.reset;
   BenchUut5();
   TraceOut_average[180] := BenchUut5.average;
   TraceOut_windowSizeReached[180] := BenchUut5.windowSizeReached;
   TraceOut_error[180] := BenchUut5.error;
   TraceOut_status[180] := BenchUut5.status;
   BenchCalls := BenchCalls + 1;
 181:
   BenchUut5.cyclicExecution := TRUE;
   BenchUut5.trigger := TRUE;
   BenchUut5.value := LREAL#49.0;
   BenchUut5.windowSize := INT#100;
   BenchUut5.reset := FALSE;
   TraceIn_cyclicExecution[181] := BenchUut5.cyclicExecution;
   TraceIn_trigger[181] := BenchUut5.trigger;
   TraceIn_value[181] := BenchUut5.value;
   TraceIn_windowSize[181] := BenchUut5.windowSize;
   TraceIn_reset[181] := BenchUut5.reset;
   BenchUut5();
   TraceOut_average[181] := BenchUut5.average;
   TraceOut_windowSizeReached[181] := BenchUut5.windowSizeReached;
   TraceOut_error[181] := BenchUut5.error;
   TraceOut_status[181] := BenchUut5.status;
   BenchCalls := BenchCalls + 1;
 182:
   BenchUut5.cyclicExecution := TRUE;
   BenchUut5.trigger := TRUE;
   BenchUut5.value := LREAL#50.0;
   BenchUut5.windowSize := INT#100;
   BenchUut5.reset := FALSE;
   TraceIn_cyclicExecution[182] := BenchUut5.cyclicExecution;
   TraceIn_trigger[182] := BenchUut5.trigger;
   TraceIn_value[182] := BenchUut5.value;
   TraceIn_windowSize[182] := BenchUut5.windowSize;
   TraceIn_reset[182] := BenchUut5.reset;
   BenchUut5();
   TraceOut_average[182] := BenchUut5.average;
   TraceOut_windowSizeReached[182] := BenchUut5.windowSizeReached;
   TraceOut_error[182] := BenchUut5.error;
   TraceOut_status[182] := BenchUut5.status;
   BenchCalls := BenchCalls + 1;
 183:
   BenchUut5.cyclicExecution := TRUE;
   BenchUut5.trigger := TRUE;
   BenchUut5.value := LREAL#51.0;
   BenchUut5.windowSize := INT#100;
   BenchUut5.reset := FALSE;
   TraceIn_cyclicExecution[183] := BenchUut5.cyclicExecution;
   TraceIn_trigger[183] := BenchUut5.trigger;
   TraceIn_value[183] := BenchUut5.value;
   TraceIn_windowSize[183] := BenchUut5.windowSize;
   TraceIn_reset[183] := BenchUut5.reset;
   BenchUut5();
   TraceOut_average[183] := BenchUut5.average;
   TraceOut_windowSizeReached[183] := BenchUut5.windowSizeReached;
   TraceOut_error[183] := BenchUut5.error;
   TraceOut_status[183] := BenchUut5.status;
   BenchCalls := BenchCalls + 1;
 184:
   BenchUut5.cyclicExecution := TRUE;
   BenchUut5.trigger := TRUE;
   BenchUut5.value := LREAL#52.0;
   BenchUut5.windowSize := INT#100;
   BenchUut5.reset := FALSE;
   TraceIn_cyclicExecution[184] := BenchUut5.cyclicExecution;
   TraceIn_trigger[184] := BenchUut5.trigger;
   TraceIn_value[184] := BenchUut5.value;
   TraceIn_windowSize[184] := BenchUut5.windowSize;
   TraceIn_reset[184] := BenchUut5.reset;
   BenchUut5();
   TraceOut_average[184] := BenchUut5.average;
   TraceOut_windowSizeReached[184] := BenchUut5.windowSizeReached;
   TraceOut_error[184] := BenchUut5.error;
   TraceOut_status[184] := BenchUut5.status;
   BenchCalls := BenchCalls + 1;
 185:
   BenchUut5.cyclicExecution := TRUE;
   BenchUut5.trigger := TRUE;
   BenchUut5.value := LREAL#53.0;
   BenchUut5.windowSize := INT#100;
   BenchUut5.reset := FALSE;
   TraceIn_cyclicExecution[185] := BenchUut5.cyclicExecution;
   TraceIn_trigger[185] := BenchUut5.trigger;
   TraceIn_value[185] := BenchUut5.value;
   TraceIn_windowSize[185] := BenchUut5.windowSize;
   TraceIn_reset[185] := BenchUut5.reset;
   BenchUut5();
   TraceOut_average[185] := BenchUut5.average;
   TraceOut_windowSizeReached[185] := BenchUut5.windowSizeReached;
   TraceOut_error[185] := BenchUut5.error;
   TraceOut_status[185] := BenchUut5.status;
   BenchCalls := BenchCalls + 1;
 186:
   BenchUut5.cyclicExecution := TRUE;
   BenchUut5.trigger := TRUE;
   BenchUut5.value := LREAL#54.0;
   BenchUut5.windowSize := INT#100;
   BenchUut5.reset := FALSE;
   TraceIn_cyclicExecution[186] := BenchUut5.cyclicExecution;
   TraceIn_trigger[186] := BenchUut5.trigger;
   TraceIn_value[186] := BenchUut5.value;
   TraceIn_windowSize[186] := BenchUut5.windowSize;
   TraceIn_reset[186] := BenchUut5.reset;
   BenchUut5();
   TraceOut_average[186] := BenchUut5.average;
   TraceOut_windowSizeReached[186] := BenchUut5.windowSizeReached;
   TraceOut_error[186] := BenchUut5.error;
   TraceOut_status[186] := BenchUut5.status;
   BenchCalls := BenchCalls + 1;
 187:
   BenchUut5.cyclicExecution := TRUE;
   BenchUut5.trigger := TRUE;
   BenchUut5.value := LREAL#55.0;
   BenchUut5.windowSize := INT#100;
   BenchUut5.reset := FALSE;
   TraceIn_cyclicExecution[187] := BenchUut5.cyclicExecution;
   TraceIn_trigger[187] := BenchUut5.trigger;
   TraceIn_value[187] := BenchUut5.value;
   TraceIn_windowSize[187] := BenchUut5.windowSize;
   TraceIn_reset[187] := BenchUut5.reset;
   BenchUut5();
   TraceOut_average[187] := BenchUut5.average;
   TraceOut_windowSizeReached[187] := BenchUut5.windowSizeReached;
   TraceOut_error[187] := BenchUut5.error;
   TraceOut_status[187] := BenchUut5.status;
   BenchCalls := BenchCalls + 1;
 188:
   BenchUut5.cyclicExecution := TRUE;
   BenchUut5.trigger := TRUE;
   BenchUut5.value := LREAL#56.0;
   BenchUut5.windowSize := INT#100;
   BenchUut5.reset := FALSE;
   TraceIn_cyclicExecution[188] := BenchUut5.cyclicExecution;
   TraceIn_trigger[188] := BenchUut5.trigger;
   TraceIn_value[188] := BenchUut5.value;
   TraceIn_windowSize[188] := BenchUut5.windowSize;
   TraceIn_reset[188] := BenchUut5.reset;
   BenchUut5();
   TraceOut_average[188] := BenchUut5.average;
   TraceOut_windowSizeReached[188] := BenchUut5.windowSizeReached;
   TraceOut_error[188] := BenchUut5.error;
   TraceOut_status[188] := BenchUut5.status;
   BenchCalls := BenchCalls + 1;
 189:
   BenchUut5.cyclicExecution := TRUE;
   BenchUut5.trigger := TRUE;
   BenchUut5.value := LREAL#57.0;
   BenchUut5.windowSize := INT#100;
   BenchUut5.reset := FALSE;
   TraceIn_cyclicExecution[189] := BenchUut5.cyclicExecution;
   TraceIn_trigger[189] := BenchUut5.trigger;
   TraceIn_value[189] := BenchUut5.value;
   TraceIn_windowSize[189] := BenchUut5.windowSize;
   TraceIn_reset[189] := BenchUut5.reset;
   BenchUut5();
   TraceOut_average[189] := BenchUut5.average;
   TraceOut_windowSizeReached[189] := BenchUut5.windowSizeReached;
   TraceOut_error[189] := BenchUut5.error;
   TraceOut_status[189] := BenchUut5.status;
   BenchCalls := BenchCalls + 1;
 190:
   BenchUut5.cyclicExecution := TRUE;
   BenchUut5.trigger := TRUE;
   BenchUut5.value := LREAL#58.0;
   BenchUut5.windowSize := INT#100;
   BenchUut5.reset := FALSE;
   TraceIn_cyclicExecution[190] := BenchUut5.cyclicExecution;
   TraceIn_trigger[190] := BenchUut5.trigger;
   TraceIn_value[190] := BenchUut5.value;
   TraceIn_windowSize[190] := BenchUut5.windowSize;
   TraceIn_reset[190] := BenchUut5.reset;
   BenchUut5();
   TraceOut_average[190] := BenchUut5.average;
   TraceOut_windowSizeReached[190] := BenchUut5.windowSizeReached;
   TraceOut_error[190] := BenchUut5.error;
   TraceOut_status[190] := BenchUut5.status;
   BenchCalls := BenchCalls + 1;
 191:
   BenchUut5.cyclicExecution := TRUE;
   BenchUut5.trigger := TRUE;
   BenchUut5.value := LREAL#59.0;
   BenchUut5.windowSize := INT#100;
   BenchUut5.reset := FALSE;
   TraceIn_cyclicExecution[191] := BenchUut5.cyclicExecution;
   TraceIn_trigger[191] := BenchUut5.trigger;
   TraceIn_value[191] := BenchUut5.value;
   TraceIn_windowSize[191] := BenchUut5.windowSize;
   TraceIn_reset[191] := BenchUut5.reset;
   BenchUut5();
   TraceOut_average[191] := BenchUut5.average;
   TraceOut_windowSizeReached[191] := BenchUut5.windowSizeReached;
   TraceOut_error[191] := BenchUut5.error;
   TraceOut_status[191] := BenchUut5.status;
   BenchCalls := BenchCalls + 1;
 192:
   BenchUut5.cyclicExecution := TRUE;
   BenchUut5.trigger := TRUE;
   BenchUut5.value := LREAL#60.0;
   BenchUut5.windowSize := INT#100;
   BenchUut5.reset := FALSE;
   TraceIn_cyclicExecution[192] := BenchUut5.cyclicExecution;
   TraceIn_trigger[192] := BenchUut5.trigger;
   TraceIn_value[192] := BenchUut5.value;
   TraceIn_windowSize[192] := BenchUut5.windowSize;
   TraceIn_reset[192] := BenchUut5.reset;
   BenchUut5();
   TraceOut_average[192] := BenchUut5.average;
   TraceOut_windowSizeReached[192] := BenchUut5.windowSizeReached;
   TraceOut_error[192] := BenchUut5.error;
   TraceOut_status[192] := BenchUut5.status;
   BenchCalls := BenchCalls + 1;
 193:
   BenchUut5.cyclicExecution := TRUE;
   BenchUut5.trigger := TRUE;
   BenchUut5.value := LREAL#61.0;
   BenchUut5.windowSize := INT#100;
   BenchUut5.reset := FALSE;
   TraceIn_cyclicExecution[193] := BenchUut5.cyclicExecution;
   TraceIn_trigger[193] := BenchUut5.trigger;
   TraceIn_value[193] := BenchUut5.value;
   TraceIn_windowSize[193] := BenchUut5.windowSize;
   TraceIn_reset[193] := BenchUut5.reset;
   BenchUut5();
   TraceOut_average[193] := BenchUut5.average;
   TraceOut_windowSizeReached[193] := BenchUut5.windowSizeReached;
   TraceOut_error[193] := BenchUut5.error;
   TraceOut_status[193] := BenchUut5.status;
   BenchCalls := BenchCalls + 1;
 194:
   BenchUut5.cyclicExecution := TRUE;
   BenchUut5.trigger := TRUE;
   BenchUut5.value := LREAL#62.0;
   BenchUut5.windowSize := INT#100;
   BenchUut5.reset := FALSE;
   TraceIn_cyclicExecution[194] := BenchUut5.cyclicExecution;
   TraceIn_trigger[194] := BenchUut5.trigger;
   TraceIn_value[194] := BenchUut5.value;
   TraceIn_windowSize[194] := BenchUut5.windowSize;
   TraceIn_reset[194] := BenchUut5.reset;
   BenchUut5();
   TraceOut_average[194] := BenchUut5.average;
   TraceOut_windowSizeReached[194] := BenchUut5.windowSizeReached;
   TraceOut_error[194] := BenchUut5.error;
   TraceOut_status[194] := BenchUut5.status;
   BenchCalls := BenchCalls + 1;
 195:
   BenchUut5.cyclicExecution := TRUE;
   BenchUut5.trigger := TRUE;
   BenchUut5.value := LREAL#63.0;
   BenchUut5.windowSize := INT#100;
   BenchUut5.reset := FALSE;
   TraceIn_cyclicExecution[195] := BenchUut5.cyclicExecution;
   TraceIn_trigger[195] := BenchUut5.trigger;
   TraceIn_value[195] := BenchUut5.value;
   TraceIn_windowSize[195] := BenchUut5.windowSize;
   TraceIn_reset[195] := BenchUut5.reset;
   BenchUut5();
   TraceOut_average[195] := BenchUut5.average;
   TraceOut_windowSizeReached[195] := BenchUut5.windowSizeReached;
   TraceOut_error[195] := BenchUut5.error;
   TraceOut_status[195] := BenchUut5.status;
   BenchCalls := BenchCalls + 1;
 196:
   BenchUut5.cyclicExecution := TRUE;
   BenchUut5.trigger := TRUE;
   BenchUut5.value := LREAL#64.0;
   BenchUut5.windowSize := INT#100;
   BenchUut5.reset := FALSE;
   TraceIn_cyclicExecution[196] := BenchUut5.cyclicExecution;
   TraceIn_trigger[196] := BenchUut5.trigger;
   TraceIn_value[196] := BenchUut5.value;
   TraceIn_windowSize[196] := BenchUut5.windowSize;
   TraceIn_reset[196] := BenchUut5.reset;
   BenchUut5();
   TraceOut_average[196] := BenchUut5.average;
   TraceOut_windowSizeReached[196] := BenchUut5.windowSizeReached;
   TraceOut_error[196] := BenchUut5.error;
   TraceOut_status[196] := BenchUut5.status;
   BenchCalls := BenchCalls + 1;
 197:
   BenchUut5.cyclicExecution := TRUE;
   BenchUut5.trigger := TRUE;
   BenchUut5.value := LREAL#65.0;
   BenchUut5.windowSize := INT#100;
   BenchUut5.reset := FALSE;
   TraceIn_cyclicExecution[197] := BenchUut5.cyclicExecution;
   TraceIn_trigger[197] := BenchUut5.trigger;
   TraceIn_value[197] := BenchUut5.value;
   TraceIn_windowSize[197] := BenchUut5.windowSize;
   TraceIn_reset[197] := BenchUut5.reset;
   BenchUut5();
   TraceOut_average[197] := BenchUut5.average;
   TraceOut_windowSizeReached[197] := BenchUut5.windowSizeReached;
   TraceOut_error[197] := BenchUut5.error;
   TraceOut_status[197] := BenchUut5.status;
   BenchCalls := BenchCalls + 1;
 198:
   BenchUut5.cyclicExecution := TRUE;
   BenchUut5.trigger := TRUE;
   BenchUut5.value := LREAL#66.0;
   BenchUut5.windowSize := INT#100;
   BenchUut5.reset := FALSE;
   TraceIn_cyclicExecution[198] := BenchUut5.cyclicExecution;
   TraceIn_trigger[198] := BenchUut5.trigger;
   TraceIn_value[198] := BenchUut5.value;
   TraceIn_windowSize[198] := BenchUut5.windowSize;
   TraceIn_reset[198] := BenchUut5.reset;
   BenchUut5();
   TraceOut_average[198] := BenchUut5.average;
   TraceOut_windowSizeReached[198] := BenchUut5.windowSizeReached;
   TraceOut_error[198] := BenchUut5.error;
   TraceOut_status[198] := BenchUut5.status;
   BenchCalls := BenchCalls + 1;
 199:
   BenchUut5.cyclicExecution := TRUE;
   BenchUut5.trigger := TRUE;
   BenchUut5.value := LREAL#67.0;
   BenchUut5.windowSize := INT#100;
   BenchUut5.reset := FALSE;
   TraceIn_cyclicExecution[199] := BenchUut5.cyclicExecution;
   TraceIn_trigger[199] := BenchUut5.trigger;
   TraceIn_value[199] := BenchUut5.value;
   TraceIn_windowSize[199] := BenchUut5.windowSize;
   TraceIn_reset[199] := BenchUut5.reset;
   BenchUut5();
   TraceOut_average[199] := BenchUut5.average;
   TraceOut_windowSizeReached[199] := BenchUut5.windowSizeReached;
   TraceOut_error[199] := BenchUut5.error;
   TraceOut_status[199] := BenchUut5.status;
   BenchCalls := BenchCalls + 1;
 200:
   BenchUut5.cyclicExecution := TRUE;
   BenchUut5.trigger := TRUE;
   BenchUut5.value := LREAL#68.0;
   BenchUut5.windowSize := INT#100;
   BenchUut5.reset := FALSE;
   TraceIn_cyclicExecution[200] := BenchUut5.cyclicExecution;
   TraceIn_trigger[200] := BenchUut5.trigger;
   TraceIn_value[200] := BenchUut5.value;
   TraceIn_windowSize[200] := BenchUut5.windowSize;
   TraceIn_reset[200] := BenchUut5.reset;
   BenchUut5();
   TraceOut_average[200] := BenchUut5.average;
   TraceOut_windowSizeReached[200] := BenchUut5.windowSizeReached;
   TraceOut_error[200] := BenchUut5.error;
   TraceOut_status[200] := BenchUut5.status;
   BenchCalls := BenchCalls + 1;
 201:
   BenchUut5.cyclicExecution := TRUE;
   BenchUut5.trigger := TRUE;
   BenchUut5.value := LREAL#69.0;
   BenchUut5.windowSize := INT#100;
   BenchUut5.reset := FALSE;
   TraceIn_cyclicExecution[201] := BenchUut5.cyclicExecution;
   TraceIn_trigger[201] := BenchUut5.trigger;
   TraceIn_value[201] := BenchUut5.value;
   TraceIn_windowSize[201] := BenchUut5.windowSize;
   TraceIn_reset[201] := BenchUut5.reset;
   BenchUut5();
   TraceOut_average[201] := BenchUut5.average;
   TraceOut_windowSizeReached[201] := BenchUut5.windowSizeReached;
   TraceOut_error[201] := BenchUut5.error;
   TraceOut_status[201] := BenchUut5.status;
   BenchCalls := BenchCalls + 1;
 202:
   BenchUut5.cyclicExecution := TRUE;
   BenchUut5.trigger := TRUE;
   BenchUut5.value := LREAL#70.0;
   BenchUut5.windowSize := INT#100;
   BenchUut5.reset := FALSE;
   TraceIn_cyclicExecution[202] := BenchUut5.cyclicExecution;
   TraceIn_trigger[202] := BenchUut5.trigger;
   TraceIn_value[202] := BenchUut5.value;
   TraceIn_windowSize[202] := BenchUut5.windowSize;
   TraceIn_reset[202] := BenchUut5.reset;
   BenchUut5();
   TraceOut_average[202] := BenchUut5.average;
   TraceOut_windowSizeReached[202] := BenchUut5.windowSizeReached;
   TraceOut_error[202] := BenchUut5.error;
   TraceOut_status[202] := BenchUut5.status;
   BenchCalls := BenchCalls + 1;
 203:
   BenchUut5.cyclicExecution := TRUE;
   BenchUut5.trigger := TRUE;
   BenchUut5.value := LREAL#71.0;
   BenchUut5.windowSize := INT#100;
   BenchUut5.reset := FALSE;
   TraceIn_cyclicExecution[203] := BenchUut5.cyclicExecution;
   TraceIn_trigger[203] := BenchUut5.trigger;
   TraceIn_value[203] := BenchUut5.value;
   TraceIn_windowSize[203] := BenchUut5.windowSize;
   TraceIn_reset[203] := BenchUut5.reset;
   BenchUut5();
   TraceOut_average[203] := BenchUut5.average;
   TraceOut_windowSizeReached[203] := BenchUut5.windowSizeReached;
   TraceOut_error[203] := BenchUut5.error;
   TraceOut_status[203] := BenchUut5.status;
   BenchCalls := BenchCalls + 1;
 204:
   BenchUut5.cyclicExecution := TRUE;
   BenchUut5.trigger := TRUE;
   BenchUut5.value := LREAL#72.0;
   BenchUut5.windowSize := INT#100;
   BenchUut5.reset := FALSE;
   TraceIn_cyclicExecution[204] := BenchUut5.cyclicExecution;
   TraceIn_trigger[204] := BenchUut5.trigger;
   TraceIn_value[204] := BenchUut5.value;
   TraceIn_windowSize[204] := BenchUut5.windowSize;
   TraceIn_reset[204] := BenchUut5.reset;
   BenchUut5();
   TraceOut_average[204] := BenchUut5.average;
   TraceOut_windowSizeReached[204] := BenchUut5.windowSizeReached;
   TraceOut_error[204] := BenchUut5.error;
   TraceOut_status[204] := BenchUut5.status;
   BenchCalls := BenchCalls + 1;
 205:
   BenchUut5.cyclicExecution := TRUE;
   BenchUut5.trigger := TRUE;
   BenchUut5.value := LREAL#73.0;
   BenchUut5.windowSize := INT#100;
   BenchUut5.reset := FALSE;
   TraceIn_cyclicExecution[205] := BenchUut5.cyclicExecution;
   TraceIn_trigger[205] := BenchUut5.trigger;
   TraceIn_value[205] := BenchUut5.value;
   TraceIn_windowSize[205] := BenchUut5.windowSize;
   TraceIn_reset[205] := BenchUut5.reset;
   BenchUut5();
   TraceOut_average[205] := BenchUut5.average;
   TraceOut_windowSizeReached[205] := BenchUut5.windowSizeReached;
   TraceOut_error[205] := BenchUut5.error;
   TraceOut_status[205] := BenchUut5.status;
   BenchCalls := BenchCalls + 1;
 206:
   BenchUut5.cyclicExecution := TRUE;
   BenchUut5.trigger := TRUE;
   BenchUut5.value := LREAL#74.0;
   BenchUut5.windowSize := INT#100;
   BenchUut5.reset := FALSE;
   TraceIn_cyclicExecution[206] := BenchUut5.cyclicExecution;
   TraceIn_trigger[206] := BenchUut5.trigger;
   TraceIn_value[206] := BenchUut5.value;
   TraceIn_windowSize[206] := BenchUut5.windowSize;
   TraceIn_reset[206] := BenchUut5.reset;
   BenchUut5();
   TraceOut_average[206] := BenchUut5.average;
   TraceOut_windowSizeReached[206] := BenchUut5.windowSizeReached;
   TraceOut_error[206] := BenchUut5.error;
   TraceOut_status[206] := BenchUut5.status;
   BenchCalls := BenchCalls + 1;
 207:
   BenchUut5.cyclicExecution := TRUE;
   BenchUut5.trigger := TRUE;
   BenchUut5.value := LREAL#75.0;
   BenchUut5.windowSize := INT#100;
   BenchUut5.reset := FALSE;
   TraceIn_cyclicExecution[207] := BenchUut5.cyclicExecution;
   TraceIn_trigger[207] := BenchUut5.trigger;
   TraceIn_value[207] := BenchUut5.value;
   TraceIn_windowSize[207] := BenchUut5.windowSize;
   TraceIn_reset[207] := BenchUut5.reset;
   BenchUut5();
   TraceOut_average[207] := BenchUut5.average;
   TraceOut_windowSizeReached[207] := BenchUut5.windowSizeReached;
   TraceOut_error[207] := BenchUut5.error;
   TraceOut_status[207] := BenchUut5.status;
   BenchCalls := BenchCalls + 1;
 208:
   BenchUut5.cyclicExecution := TRUE;
   BenchUut5.trigger := TRUE;
   BenchUut5.value := LREAL#76.0;
   BenchUut5.windowSize := INT#100;
   BenchUut5.reset := FALSE;
   TraceIn_cyclicExecution[208] := BenchUut5.cyclicExecution;
   TraceIn_trigger[208] := BenchUut5.trigger;
   TraceIn_value[208] := BenchUut5.value;
   TraceIn_windowSize[208] := BenchUut5.windowSize;
   TraceIn_reset[208] := BenchUut5.reset;
   BenchUut5();
   TraceOut_average[208] := BenchUut5.average;
   TraceOut_windowSizeReached[208] := BenchUut5.windowSizeReached;
   TraceOut_error[208] := BenchUut5.error;
   TraceOut_status[208] := BenchUut5.status;
   BenchCalls := BenchCalls + 1;
 209:
   BenchUut5.cyclicExecution := TRUE;
   BenchUut5.trigger := TRUE;
   BenchUut5.value := LREAL#77.0;
   BenchUut5.windowSize := INT#100;
   BenchUut5.reset := FALSE;
   TraceIn_cyclicExecution[209] := BenchUut5.cyclicExecution;
   TraceIn_trigger[209] := BenchUut5.trigger;
   TraceIn_value[209] := BenchUut5.value;
   TraceIn_windowSize[209] := BenchUut5.windowSize;
   TraceIn_reset[209] := BenchUut5.reset;
   BenchUut5();
   TraceOut_average[209] := BenchUut5.average;
   TraceOut_windowSizeReached[209] := BenchUut5.windowSizeReached;
   TraceOut_error[209] := BenchUut5.error;
   TraceOut_status[209] := BenchUut5.status;
   BenchCalls := BenchCalls + 1;
 210:
   BenchUut5.cyclicExecution := TRUE;
   BenchUut5.trigger := TRUE;
   BenchUut5.value := LREAL#78.0;
   BenchUut5.windowSize := INT#100;
   BenchUut5.reset := FALSE;
   TraceIn_cyclicExecution[210] := BenchUut5.cyclicExecution;
   TraceIn_trigger[210] := BenchUut5.trigger;
   TraceIn_value[210] := BenchUut5.value;
   TraceIn_windowSize[210] := BenchUut5.windowSize;
   TraceIn_reset[210] := BenchUut5.reset;
   BenchUut5();
   TraceOut_average[210] := BenchUut5.average;
   TraceOut_windowSizeReached[210] := BenchUut5.windowSizeReached;
   TraceOut_error[210] := BenchUut5.error;
   TraceOut_status[210] := BenchUut5.status;
   BenchCalls := BenchCalls + 1;
 211:
   BenchUut5.cyclicExecution := TRUE;
   BenchUut5.trigger := TRUE;
   BenchUut5.value := LREAL#79.0;
   BenchUut5.windowSize := INT#100;
   BenchUut5.reset := FALSE;
   TraceIn_cyclicExecution[211] := BenchUut5.cyclicExecution;
   TraceIn_trigger[211] := BenchUut5.trigger;
   TraceIn_value[211] := BenchUut5.value;
   TraceIn_windowSize[211] := BenchUut5.windowSize;
   TraceIn_reset[211] := BenchUut5.reset;
   BenchUut5();
   TraceOut_average[211] := BenchUut5.average;
   TraceOut_windowSizeReached[211] := BenchUut5.windowSizeReached;
   TraceOut_error[211] := BenchUut5.error;
   TraceOut_status[211] := BenchUut5.status;
   BenchCalls := BenchCalls + 1;
 212:
   BenchUut5.cyclicExecution := TRUE;
   BenchUut5.trigger := TRUE;
   BenchUut5.value := LREAL#80.0;
   BenchUut5.windowSize := INT#100;
   BenchUut5.reset := FALSE;
   TraceIn_cyclicExecution[212] := BenchUut5.cyclicExecution;
   TraceIn_trigger[212] := BenchUut5.trigger;
   TraceIn_value[212] := BenchUut5.value;
   TraceIn_windowSize[212] := BenchUut5.windowSize;
   TraceIn_reset[212] := BenchUut5.reset;
   BenchUut5();
   TraceOut_average[212] := BenchUut5.average;
   TraceOut_windowSizeReached[212] := BenchUut5.windowSizeReached;
   TraceOut_error[212] := BenchUut5.error;
   TraceOut_status[212] := BenchUut5.status;
   BenchCalls := BenchCalls + 1;
 213:
   BenchUut5.cyclicExecution := TRUE;
   BenchUut5.trigger := TRUE;
   BenchUut5.value := LREAL#81.0;
   BenchUut5.windowSize := INT#100;
   BenchUut5.reset := FALSE;
   TraceIn_cyclicExecution[213] := BenchUut5.cyclicExecution;
   TraceIn_trigger[213] := BenchUut5.trigger;
   TraceIn_value[213] := BenchUut5.value;
   TraceIn_windowSize[213] := BenchUut5.windowSize;
   TraceIn_reset[213] := BenchUut5.reset;
   BenchUut5();
   TraceOut_average[213] := BenchUut5.average;
   TraceOut_windowSizeReached[213] := BenchUut5.windowSizeReached;
   TraceOut_error[213] := BenchUut5.error;
   TraceOut_status[213] := BenchUut5.status;
   BenchCalls := BenchCalls + 1;
 214:
   BenchUut5.cyclicExecution := TRUE;
   BenchUut5.trigger := TRUE;
   BenchUut5.value := LREAL#82.0;
   BenchUut5.windowSize := INT#100;
   BenchUut5.reset := FALSE;
   TraceIn_cyclicExecution[214] := BenchUut5.cyclicExecution;
   TraceIn_trigger[214] := BenchUut5.trigger;
   TraceIn_value[214] := BenchUut5.value;
   TraceIn_windowSize[214] := BenchUut5.windowSize;
   TraceIn_reset[214] := BenchUut5.reset;
   BenchUut5();
   TraceOut_average[214] := BenchUut5.average;
   TraceOut_windowSizeReached[214] := BenchUut5.windowSizeReached;
   TraceOut_error[214] := BenchUut5.error;
   TraceOut_status[214] := BenchUut5.status;
   BenchCalls := BenchCalls + 1;
 215:
   BenchUut5.cyclicExecution := TRUE;
   BenchUut5.trigger := TRUE;
   BenchUut5.value := LREAL#83.0;
   BenchUut5.windowSize := INT#100;
   BenchUut5.reset := FALSE;
   TraceIn_cyclicExecution[215] := BenchUut5.cyclicExecution;
   TraceIn_trigger[215] := BenchUut5.trigger;
   TraceIn_value[215] := BenchUut5.value;
   TraceIn_windowSize[215] := BenchUut5.windowSize;
   TraceIn_reset[215] := BenchUut5.reset;
   BenchUut5();
   TraceOut_average[215] := BenchUut5.average;
   TraceOut_windowSizeReached[215] := BenchUut5.windowSizeReached;
   TraceOut_error[215] := BenchUut5.error;
   TraceOut_status[215] := BenchUut5.status;
   BenchCalls := BenchCalls + 1;
 216:
   BenchUut5.cyclicExecution := TRUE;
   BenchUut5.trigger := TRUE;
   BenchUut5.value := LREAL#84.0;
   BenchUut5.windowSize := INT#100;
   BenchUut5.reset := FALSE;
   TraceIn_cyclicExecution[216] := BenchUut5.cyclicExecution;
   TraceIn_trigger[216] := BenchUut5.trigger;
   TraceIn_value[216] := BenchUut5.value;
   TraceIn_windowSize[216] := BenchUut5.windowSize;
   TraceIn_reset[216] := BenchUut5.reset;
   BenchUut5();
   TraceOut_average[216] := BenchUut5.average;
   TraceOut_windowSizeReached[216] := BenchUut5.windowSizeReached;
   TraceOut_error[216] := BenchUut5.error;
   TraceOut_status[216] := BenchUut5.status;
   BenchCalls := BenchCalls + 1;
 217:
   BenchUut5.cyclicExecution := TRUE;
   BenchUut5.trigger := TRUE;
   BenchUut5.value := LREAL#85.0;
   BenchUut5.windowSize := INT#100;
   BenchUut5.reset := FALSE;
   TraceIn_cyclicExecution[217] := BenchUut5.cyclicExecution;
   TraceIn_trigger[217] := BenchUut5.trigger;
   TraceIn_value[217] := BenchUut5.value;
   TraceIn_windowSize[217] := BenchUut5.windowSize;
   TraceIn_reset[217] := BenchUut5.reset;
   BenchUut5();
   TraceOut_average[217] := BenchUut5.average;
   TraceOut_windowSizeReached[217] := BenchUut5.windowSizeReached;
   TraceOut_error[217] := BenchUut5.error;
   TraceOut_status[217] := BenchUut5.status;
   BenchCalls := BenchCalls + 1;
 218:
   BenchUut5.cyclicExecution := TRUE;
   BenchUut5.trigger := TRUE;
   BenchUut5.value := LREAL#86.0;
   BenchUut5.windowSize := INT#100;
   BenchUut5.reset := FALSE;
   TraceIn_cyclicExecution[218] := BenchUut5.cyclicExecution;
   TraceIn_trigger[218] := BenchUut5.trigger;
   TraceIn_value[218] := BenchUut5.value;
   TraceIn_windowSize[218] := BenchUut5.windowSize;
   TraceIn_reset[218] := BenchUut5.reset;
   BenchUut5();
   TraceOut_average[218] := BenchUut5.average;
   TraceOut_windowSizeReached[218] := BenchUut5.windowSizeReached;
   TraceOut_error[218] := BenchUut5.error;
   TraceOut_status[218] := BenchUut5.status;
   BenchCalls := BenchCalls + 1;
 219:
   BenchUut5.cyclicExecution := TRUE;
   BenchUut5.trigger := TRUE;
   BenchUut5.value := LREAL#87.0;
   BenchUut5.windowSize := INT#100;
   BenchUut5.reset := FALSE;
   TraceIn_cyclicExecution[219] := BenchUut5.cyclicExecution;
   TraceIn_trigger[219] := BenchUut5.trigger;
   TraceIn_value[219] := BenchUut5.value;
   TraceIn_windowSize[219] := BenchUut5.windowSize;
   TraceIn_reset[219] := BenchUut5.reset;
   BenchUut5();
   TraceOut_average[219] := BenchUut5.average;
   TraceOut_windowSizeReached[219] := BenchUut5.windowSizeReached;
   TraceOut_error[219] := BenchUut5.error;
   TraceOut_status[219] := BenchUut5.status;
   BenchCalls := BenchCalls + 1;
 220:
   BenchUut5.cyclicExecution := TRUE;
   BenchUut5.trigger := TRUE;
   BenchUut5.value := LREAL#88.0;
   BenchUut5.windowSize := INT#100;
   BenchUut5.reset := FALSE;
   TraceIn_cyclicExecution[220] := BenchUut5.cyclicExecution;
   TraceIn_trigger[220] := BenchUut5.trigger;
   TraceIn_value[220] := BenchUut5.value;
   TraceIn_windowSize[220] := BenchUut5.windowSize;
   TraceIn_reset[220] := BenchUut5.reset;
   BenchUut5();
   TraceOut_average[220] := BenchUut5.average;
   TraceOut_windowSizeReached[220] := BenchUut5.windowSizeReached;
   TraceOut_error[220] := BenchUut5.error;
   TraceOut_status[220] := BenchUut5.status;
   BenchCalls := BenchCalls + 1;
 221:
   BenchUut5.cyclicExecution := TRUE;
   BenchUut5.trigger := TRUE;
   BenchUut5.value := LREAL#89.0;
   BenchUut5.windowSize := INT#100;
   BenchUut5.reset := FALSE;
   TraceIn_cyclicExecution[221] := BenchUut5.cyclicExecution;
   TraceIn_trigger[221] := BenchUut5.trigger;
   TraceIn_value[221] := BenchUut5.value;
   TraceIn_windowSize[221] := BenchUut5.windowSize;
   TraceIn_reset[221] := BenchUut5.reset;
   BenchUut5();
   TraceOut_average[221] := BenchUut5.average;
   TraceOut_windowSizeReached[221] := BenchUut5.windowSizeReached;
   TraceOut_error[221] := BenchUut5.error;
   TraceOut_status[221] := BenchUut5.status;
   BenchCalls := BenchCalls + 1;
 222:
   BenchUut5.cyclicExecution := TRUE;
   BenchUut5.trigger := TRUE;
   BenchUut5.value := LREAL#90.0;
   BenchUut5.windowSize := INT#100;
   BenchUut5.reset := FALSE;
   TraceIn_cyclicExecution[222] := BenchUut5.cyclicExecution;
   TraceIn_trigger[222] := BenchUut5.trigger;
   TraceIn_value[222] := BenchUut5.value;
   TraceIn_windowSize[222] := BenchUut5.windowSize;
   TraceIn_reset[222] := BenchUut5.reset;
   BenchUut5();
   TraceOut_average[222] := BenchUut5.average;
   TraceOut_windowSizeReached[222] := BenchUut5.windowSizeReached;
   TraceOut_error[222] := BenchUut5.error;
   TraceOut_status[222] := BenchUut5.status;
   BenchCalls := BenchCalls + 1;
 223:
   BenchUut5.cyclicExecution := TRUE;
   BenchUut5.trigger := TRUE;
   BenchUut5.value := LREAL#91.0;
   BenchUut5.windowSize := INT#100;
   BenchUut5.reset := FALSE;
   TraceIn_cyclicExecution[223] := BenchUut5.cyclicExecution;
   TraceIn_trigger[223] := BenchUut5.trigger;
   TraceIn_value[223] := BenchUut5.value;
   TraceIn_windowSize[223] := BenchUut5.windowSize;
   TraceIn_reset[223] := BenchUut5.reset;
   BenchUut5();
   TraceOut_average[223] := BenchUut5.average;
   TraceOut_windowSizeReached[223] := BenchUut5.windowSizeReached;
   TraceOut_error[223] := BenchUut5.error;
   TraceOut_status[223] := BenchUut5.status;
   BenchCalls := BenchCalls + 1;
 224:
   BenchUut5.cyclicExecution := TRUE;
   BenchUut5.trigger := TRUE;
   BenchUut5.value := LREAL#92.0;
   BenchUut5.windowSize := INT#100;
   BenchUut5.reset := FALSE;
   TraceIn_cyclicExecution[224] := BenchUut5.cyclicExecution;
   TraceIn_trigger[224] := BenchUut5.trigger;
   TraceIn_value[224] := BenchUut5.value;
   TraceIn_windowSize[224] := BenchUut5.windowSize;
   TraceIn_reset[224] := BenchUut5.reset;
   BenchUut5();
   TraceOut_average[224] := BenchUut5.average;
   TraceOut_windowSizeReached[224] := BenchUut5.windowSizeReached;
   TraceOut_error[224] := BenchUut5.error;
   TraceOut_status[224] := BenchUut5.status;
   BenchCalls := BenchCalls + 1;
 225:
   BenchUut5.cyclicExecution := TRUE;
   BenchUut5.trigger := TRUE;
   BenchUut5.value := LREAL#93.0;
   BenchUut5.windowSize := INT#100;
   BenchUut5.reset := FALSE;
   TraceIn_cyclicExecution[225] := BenchUut5.cyclicExecution;
   TraceIn_trigger[225] := BenchUut5.trigger;
   TraceIn_value[225] := BenchUut5.value;
   TraceIn_windowSize[225] := BenchUut5.windowSize;
   TraceIn_reset[225] := BenchUut5.reset;
   BenchUut5();
   TraceOut_average[225] := BenchUut5.average;
   TraceOut_windowSizeReached[225] := BenchUut5.windowSizeReached;
   TraceOut_error[225] := BenchUut5.error;
   TraceOut_status[225] := BenchUut5.status;
   BenchCalls := BenchCalls + 1;
 226:
   BenchUut5.cyclicExecution := TRUE;
   BenchUut5.trigger := TRUE;
   BenchUut5.value := LREAL#94.0;
   BenchUut5.windowSize := INT#100;
   BenchUut5.reset := FALSE;
   TraceIn_cyclicExecution[226] := BenchUut5.cyclicExecution;
   TraceIn_trigger[226] := BenchUut5.trigger;
   TraceIn_value[226] := BenchUut5.value;
   TraceIn_windowSize[226] := BenchUut5.windowSize;
   TraceIn_reset[226] := BenchUut5.reset;
   BenchUut5();
   TraceOut_average[226] := BenchUut5.average;
   TraceOut_windowSizeReached[226] := BenchUut5.windowSizeReached;
   TraceOut_error[226] := BenchUut5.error;
   TraceOut_status[226] := BenchUut5.status;
   BenchCalls := BenchCalls + 1;
 227:
   BenchUut5.cyclicExecution := TRUE;
   BenchUut5.trigger := TRUE;
   BenchUut5.value := LREAL#95.0;
   BenchUut5.windowSize := INT#100;
   BenchUut5.reset := FALSE;
   TraceIn_cyclicExecution[227] := BenchUut5.cyclicExecution;
   TraceIn_trigger[227] := BenchUut5.trigger;
   TraceIn_value[227] := BenchUut5.value;
   TraceIn_windowSize[227] := BenchUut5.windowSize;
   TraceIn_reset[227] := BenchUut5.reset;
   BenchUut5();
   TraceOut_average[227] := BenchUut5.average;
   TraceOut_windowSizeReached[227] := BenchUut5.windowSizeReached;
   TraceOut_error[227] := BenchUut5.error;
   TraceOut_status[227] := BenchUut5.status;
   BenchCalls := BenchCalls + 1;
 228:
   BenchUut5.cyclicExecution := TRUE;
   BenchUut5.trigger := TRUE;
   BenchUut5.value := LREAL#96.0;
   BenchUut5.windowSize := INT#100;
   BenchUut5.reset := FALSE;
   TraceIn_cyclicExecution[228] := BenchUut5.cyclicExecution;
   TraceIn_trigger[228] := BenchUut5.trigger;
   TraceIn_value[228] := BenchUut5.value;
   TraceIn_windowSize[228] := BenchUut5.windowSize;
   TraceIn_reset[228] := BenchUut5.reset;
   BenchUut5();
   TraceOut_average[228] := BenchUut5.average;
   TraceOut_windowSizeReached[228] := BenchUut5.windowSizeReached;
   TraceOut_error[228] := BenchUut5.error;
   TraceOut_status[228] := BenchUut5.status;
   BenchCalls := BenchCalls + 1;
 229:
   BenchUut5.cyclicExecution := TRUE;
   BenchUut5.trigger := TRUE;
   BenchUut5.value := LREAL#97.0;
   BenchUut5.windowSize := INT#100;
   BenchUut5.reset := FALSE;
   TraceIn_cyclicExecution[229] := BenchUut5.cyclicExecution;
   TraceIn_trigger[229] := BenchUut5.trigger;
   TraceIn_value[229] := BenchUut5.value;
   TraceIn_windowSize[229] := BenchUut5.windowSize;
   TraceIn_reset[229] := BenchUut5.reset;
   BenchUut5();
   TraceOut_average[229] := BenchUut5.average;
   TraceOut_windowSizeReached[229] := BenchUut5.windowSizeReached;
   TraceOut_error[229] := BenchUut5.error;
   TraceOut_status[229] := BenchUut5.status;
   BenchCalls := BenchCalls + 1;
 230:
   BenchUut5.cyclicExecution := TRUE;
   BenchUut5.trigger := TRUE;
   BenchUut5.value := LREAL#98.0;
   BenchUut5.windowSize := INT#100;
   BenchUut5.reset := FALSE;
   TraceIn_cyclicExecution[230] := BenchUut5.cyclicExecution;
   TraceIn_trigger[230] := BenchUut5.trigger;
   TraceIn_value[230] := BenchUut5.value;
   TraceIn_windowSize[230] := BenchUut5.windowSize;
   TraceIn_reset[230] := BenchUut5.reset;
   BenchUut5();
   TraceOut_average[230] := BenchUut5.average;
   TraceOut_windowSizeReached[230] := BenchUut5.windowSizeReached;
   TraceOut_error[230] := BenchUut5.error;
   TraceOut_status[230] := BenchUut5.status;
   BenchCalls := BenchCalls + 1;
 231:
   BenchUut5.cyclicExecution := TRUE;
   BenchUut5.trigger := TRUE;
   BenchUut5.value := LREAL#99.0;
   BenchUut5.windowSize := INT#100;
   BenchUut5.reset := FALSE;
   TraceIn_cyclicExecution[231] := BenchUut5.cyclicExecution;
   TraceIn_trigger[231] := BenchUut5.trigger;
   TraceIn_value[231] := BenchUut5.value;
   TraceIn_windowSize[231] := BenchUut5.windowSize;
   TraceIn_reset[231] := BenchUut5.reset;
   BenchUut5();
   TraceOut_average[231] := BenchUut5.average;
   TraceOut_windowSizeReached[231] := BenchUut5.windowSizeReached;
   TraceOut_error[231] := BenchUut5.error;
   TraceOut_status[231] := BenchUut5.status;
   BenchCalls := BenchCalls + 1;
 232:
   BenchUut5.cyclicExecution := TRUE;
   BenchUut5.trigger := TRUE;
   BenchUut5.value := LREAL#100.0;
   BenchUut5.windowSize := INT#100;
   BenchUut5.reset := FALSE;
   TraceIn_cyclicExecution[232] := BenchUut5.cyclicExecution;
   TraceIn_trigger[232] := BenchUut5.trigger;
   TraceIn_value[232] := BenchUut5.value;
   TraceIn_windowSize[232] := BenchUut5.windowSize;
   TraceIn_reset[232] := BenchUut5.reset;
   BenchUut5();
   TraceOut_average[232] := BenchUut5.average;
   TraceOut_windowSizeReached[232] := BenchUut5.windowSizeReached;
   TraceOut_error[232] := BenchUut5.error;
   TraceOut_status[232] := BenchUut5.status;
   BenchCalls := BenchCalls + 1;
 233:
   BenchUut5.cyclicExecution := TRUE;
   BenchUut5.trigger := TRUE;
   BenchUut5.value := LREAL#101.0;
   BenchUut5.windowSize := INT#100;
   BenchUut5.reset := FALSE;
   TraceIn_cyclicExecution[233] := BenchUut5.cyclicExecution;
   TraceIn_trigger[233] := BenchUut5.trigger;
   TraceIn_value[233] := BenchUut5.value;
   TraceIn_windowSize[233] := BenchUut5.windowSize;
   TraceIn_reset[233] := BenchUut5.reset;
   BenchUut5();
   TraceOut_average[233] := BenchUut5.average;
   TraceOut_windowSizeReached[233] := BenchUut5.windowSizeReached;
   TraceOut_error[233] := BenchUut5.error;
   TraceOut_status[233] := BenchUut5.status;
   BenchCalls := BenchCalls + 1;
 234:
   BenchUut5.cyclicExecution := TRUE;
   BenchUut5.trigger := TRUE;
   BenchUut5.value := LREAL#102.0;
   BenchUut5.windowSize := INT#100;
   BenchUut5.reset := FALSE;
   TraceIn_cyclicExecution[234] := BenchUut5.cyclicExecution;
   TraceIn_trigger[234] := BenchUut5.trigger;
   TraceIn_value[234] := BenchUut5.value;
   TraceIn_windowSize[234] := BenchUut5.windowSize;
   TraceIn_reset[234] := BenchUut5.reset;
   BenchUut5();
   TraceOut_average[234] := BenchUut5.average;
   TraceOut_windowSizeReached[234] := BenchUut5.windowSizeReached;
   TraceOut_error[234] := BenchUut5.error;
   TraceOut_status[234] := BenchUut5.status;
   BenchCalls := BenchCalls + 1;
 235:
   BenchUut5.cyclicExecution := TRUE;
   BenchUut5.trigger := TRUE;
   BenchUut5.value := LREAL#103.0;
   BenchUut5.windowSize := INT#100;
   BenchUut5.reset := FALSE;
   TraceIn_cyclicExecution[235] := BenchUut5.cyclicExecution;
   TraceIn_trigger[235] := BenchUut5.trigger;
   TraceIn_value[235] := BenchUut5.value;
   TraceIn_windowSize[235] := BenchUut5.windowSize;
   TraceIn_reset[235] := BenchUut5.reset;
   BenchUut5();
   TraceOut_average[235] := BenchUut5.average;
   TraceOut_windowSizeReached[235] := BenchUut5.windowSizeReached;
   TraceOut_error[235] := BenchUut5.error;
   TraceOut_status[235] := BenchUut5.status;
   BenchCalls := BenchCalls + 1;
 236:
   BenchUut5.cyclicExecution := TRUE;
   BenchUut5.trigger := TRUE;
   BenchUut5.value := LREAL#104.0;
   BenchUut5.windowSize := INT#100;
   BenchUut5.reset := FALSE;
   TraceIn_cyclicExecution[236] := BenchUut5.cyclicExecution;
   TraceIn_trigger[236] := BenchUut5.trigger;
   TraceIn_value[236] := BenchUut5.value;
   TraceIn_windowSize[236] := BenchUut5.windowSize;
   TraceIn_reset[236] := BenchUut5.reset;
   BenchUut5();
   TraceOut_average[236] := BenchUut5.average;
   TraceOut_windowSizeReached[236] := BenchUut5.windowSizeReached;
   TraceOut_error[236] := BenchUut5.error;
   TraceOut_status[236] := BenchUut5.status;
   BenchCalls := BenchCalls + 1;
 237:
   BenchUut5.cyclicExecution := TRUE;
   BenchUut5.trigger := FALSE;
   BenchUut5.value := LREAL#104.0;
   BenchUut5.windowSize := INT#2;
   BenchUut5.reset := FALSE;
   TraceIn_cyclicExecution[237] := BenchUut5.cyclicExecution;
   TraceIn_trigger[237] := BenchUut5.trigger;
   TraceIn_value[237] := BenchUut5.value;
   TraceIn_windowSize[237] := BenchUut5.windowSize;
   TraceIn_reset[237] := BenchUut5.reset;
   BenchUut5();
   TraceOut_average[237] := BenchUut5.average;
   TraceOut_windowSizeReached[237] := BenchUut5.windowSizeReached;
   TraceOut_error[237] := BenchUut5.error;
   TraceOut_status[237] := BenchUut5.status;
   BenchCalls := BenchCalls + 1;
 238:
   BenchUut5.cyclicExecution := TRUE;
   BenchUut5.trigger := TRUE;
   BenchUut5.value := LREAL#5.0;
   BenchUut5.windowSize := INT#2;
   BenchUut5.reset := FALSE;
   TraceIn_cyclicExecution[238] := BenchUut5.cyclicExecution;
   TraceIn_trigger[238] := BenchUut5.trigger;
   TraceIn_value[238] := BenchUut5.value;
   TraceIn_windowSize[238] := BenchUut5.windowSize;
   TraceIn_reset[238] := BenchUut5.reset;
   BenchUut5();
   TraceOut_average[238] := BenchUut5.average;
   TraceOut_windowSizeReached[238] := BenchUut5.windowSizeReached;
   TraceOut_error[238] := BenchUut5.error;
   TraceOut_status[238] := BenchUut5.status;
   BenchCalls := BenchCalls + 1;
 239:
   BenchUut5.cyclicExecution := TRUE;
   BenchUut5.trigger := FALSE;
   BenchUut5.value := LREAL#5.0;
   BenchUut5.windowSize := INT#100;
   BenchUut5.reset := FALSE;
   TraceIn_cyclicExecution[239] := BenchUut5.cyclicExecution;
   TraceIn_trigger[239] := BenchUut5.trigger;
   TraceIn_value[239] := BenchUut5.value;
   TraceIn_windowSize[239] := BenchUut5.windowSize;
   TraceIn_reset[239] := BenchUut5.reset;
   BenchUut5();
   TraceOut_average[239] := BenchUut5.average;
   TraceOut_windowSizeReached[239] := BenchUut5.windowSizeReached;
   TraceOut_error[239] := BenchUut5.error;
   TraceOut_status[239] := BenchUut5.status;
   BenchCalls := BenchCalls + 1;
 240:
   BenchUut5.cyclicExecution := TRUE;
   BenchUut5.trigger := TRUE;
   BenchUut5.value := LREAL#7.0;
   BenchUut5.windowSize := INT#100;
   BenchUut5.reset := FALSE;
   TraceIn_cyclicExecution[240] := BenchUut5.cyclicExecution;
   TraceIn_trigger[240] := BenchUut5.trigger;
   TraceIn_value[240] := BenchUut5.value;
   TraceIn_windowSize[240] := BenchUut5.windowSize;
   TraceIn_reset[240] := BenchUut5.reset;
   BenchUut5();
   TraceOut_average[240] := BenchUut5.average;
   TraceOut_windowSizeReached[240] := BenchUut5.windowSizeReached;
   TraceOut_error[240] := BenchUut5.error;
   TraceOut_status[240] := BenchUut5.status;
   BenchCalls := BenchCalls + 1;
 241:
   BenchUut6.cyclicExecution := FALSE;
   BenchUut6.trigger := FALSE;
   BenchUut6.value := LREAL#3.0;
   BenchUut6.windowSize := INT#100;
   BenchUut6.reset := FALSE;
   TraceIn_cyclicExecution[241] := BenchUut6.cyclicExecution;
   TraceIn_trigger[241] := BenchUut6.trigger;
   TraceIn_value[241] := BenchUut6.value;
   TraceIn_windowSize[241] := BenchUut6.windowSize;
   TraceIn_reset[241] := BenchUut6.reset;
   BenchUut6();
   TraceOut_average[241] := BenchUut6.average;
   TraceOut_windowSizeReached[241] := BenchUut6.windowSizeReached;
   TraceOut_error[241] := BenchUut6.error;
   TraceOut_status[241] := BenchUut6.status;
   BenchCalls := BenchCalls + 1;
 242:
   BenchUut6.cyclicExecution := FALSE;
   BenchUut6.trigger := TRUE;
   BenchUut6.value := LREAL#0.0;
   BenchUut6.windowSize := INT#100;
   BenchUut6.reset := FALSE;
   TraceIn_cyclicExecution[242] := BenchUut6.cyclicExecution;
   TraceIn_trigger[242] := BenchUut6.trigger;
   TraceIn_value[242] := BenchUut6.value;
   TraceIn_windowSize[242] := BenchUut6.windowSize;
   TraceIn_reset[242] := BenchUut6.reset;
   BenchUut6();
   TraceOut_average[242] := BenchUut6.average;
   TraceOut_windowSizeReached[242] := BenchUut6.windowSizeReached;
   TraceOut_error[242] := BenchUut6.error;
   TraceOut_status[242] := BenchUut6.status;
   BenchCalls := BenchCalls + 1;
 243:
   BenchUut6.cyclicExecution := FALSE;
   BenchUut6.trigger := FALSE;
   BenchUut6.value := LREAL#0.0;
   BenchUut6.windowSize := INT#100;
   BenchUut6.reset := FALSE;
   TraceIn_cyclicExecution[243] := BenchUut6.cyclicExecution;
   TraceIn_trigger[243] := BenchUut6.trigger;
   TraceIn_value[243] := BenchUut6.value;
   TraceIn_windowSize[243] := BenchUut6.windowSize;
   TraceIn_reset[243] := BenchUut6.reset;
   BenchUut6();
   TraceOut_average[243] := BenchUut6.average;
   TraceOut_windowSizeReached[243] := BenchUut6.windowSizeReached;
   TraceOut_error[243] := BenchUut6.error;
   TraceOut_status[243] := BenchUut6.status;
   BenchCalls := BenchCalls + 1;
 244:
   BenchUut6.cyclicExecution := FALSE;
   BenchUut6.trigger := TRUE;
   BenchUut6.value := LREAL#1.0;
   BenchUut6.windowSize := INT#100;
   BenchUut6.reset := FALSE;
   TraceIn_cyclicExecution[244] := BenchUut6.cyclicExecution;
   TraceIn_trigger[244] := BenchUut6.trigger;
   TraceIn_value[244] := BenchUut6.value;
   TraceIn_windowSize[244] := BenchUut6.windowSize;
   TraceIn_reset[244] := BenchUut6.reset;
   BenchUut6();
   TraceOut_average[244] := BenchUut6.average;
   TraceOut_windowSizeReached[244] := BenchUut6.windowSizeReached;
   TraceOut_error[244] := BenchUut6.error;
   TraceOut_status[244] := BenchUut6.status;
   BenchCalls := BenchCalls + 1;
 245:
   BenchUut6.cyclicExecution := FALSE;
   BenchUut6.trigger := FALSE;
   BenchUut6.value := LREAL#1.0;
   BenchUut6.windowSize := INT#100;
   BenchUut6.reset := FALSE;
   TraceIn_cyclicExecution[245] := BenchUut6.cyclicExecution;
   TraceIn_trigger[245] := BenchUut6.trigger;
   TraceIn_value[245] := BenchUut6.value;
   TraceIn_windowSize[245] := BenchUut6.windowSize;
   TraceIn_reset[245] := BenchUut6.reset;
   BenchUut6();
   TraceOut_average[245] := BenchUut6.average;
   TraceOut_windowSizeReached[245] := BenchUut6.windowSizeReached;
   TraceOut_error[245] := BenchUut6.error;
   TraceOut_status[245] := BenchUut6.status;
   BenchCalls := BenchCalls + 1;
 246:
   BenchUut6.cyclicExecution := FALSE;
   BenchUut6.trigger := TRUE;
   BenchUut6.value := LREAL#2.0;
   BenchUut6.windowSize := INT#100;
   BenchUut6.reset := FALSE;
   TraceIn_cyclicExecution[246] := BenchUut6.cyclicExecution;
   TraceIn_trigger[246] := BenchUut6.trigger;
   TraceIn_value[246] := BenchUut6.value;
   TraceIn_windowSize[246] := BenchUut6.windowSize;
   TraceIn_reset[246] := BenchUut6.reset;
   BenchUut6();
   TraceOut_average[246] := BenchUut6.average;
   TraceOut_windowSizeReached[246] := BenchUut6.windowSizeReached;
   TraceOut_error[246] := BenchUut6.error;
   TraceOut_status[246] := BenchUut6.status;
   BenchCalls := BenchCalls + 1;
 247:
   BenchUut6.cyclicExecution := FALSE;
   BenchUut6.trigger := FALSE;
   BenchUut6.value := LREAL#2.0;
   BenchUut6.windowSize := INT#100;
   BenchUut6.reset := FALSE;
   TraceIn_cyclicExecution[247] := BenchUut6.cyclicExecution;
   TraceIn_trigger[247] := BenchUut6.trigger;
   TraceIn_value[247] := BenchUut6.value;
   TraceIn_windowSize[247] := BenchUut6.windowSize;
   TraceIn_reset[247] := BenchUut6.reset;
   BenchUut6();
   TraceOut_average[247] := BenchUut6.average;
   TraceOut_windowSizeReached[247] := BenchUut6.windowSizeReached;
   TraceOut_error[247] := BenchUut6.error;
   TraceOut_status[247] := BenchUut6.status;
   BenchCalls := BenchCalls + 1;
 248:
   BenchUut6.cyclicExecution := FALSE;
   BenchUut6.trigger := TRUE;
   BenchUut6.value := LREAL#3.0;
   BenchUut6.windowSize := INT#100;
   BenchUut6.reset := FALSE;
   TraceIn_cyclicExecution[248] := BenchUut6.cyclicExecution;
   TraceIn_trigger[248] := BenchUut6.trigger;
   TraceIn_value[248] := BenchUut6.value;
   TraceIn_windowSize[248] := BenchUut6.windowSize;
   TraceIn_reset[248] := BenchUut6.reset;
   BenchUut6();
   TraceOut_average[248] := BenchUut6.average;
   TraceOut_windowSizeReached[248] := BenchUut6.windowSizeReached;
   TraceOut_error[248] := BenchUut6.error;
   TraceOut_status[248] := BenchUut6.status;
   BenchCalls := BenchCalls + 1;
 249:
   BenchUut6.cyclicExecution := FALSE;
   BenchUut6.trigger := FALSE;
   BenchUut6.value := LREAL#3.0;
   BenchUut6.windowSize := INT#100;
   BenchUut6.reset := FALSE;
   TraceIn_cyclicExecution[249] := BenchUut6.cyclicExecution;
   TraceIn_trigger[249] := BenchUut6.trigger;
   TraceIn_value[249] := BenchUut6.value;
   TraceIn_windowSize[249] := BenchUut6.windowSize;
   TraceIn_reset[249] := BenchUut6.reset;
   BenchUut6();
   TraceOut_average[249] := BenchUut6.average;
   TraceOut_windowSizeReached[249] := BenchUut6.windowSizeReached;
   TraceOut_error[249] := BenchUut6.error;
   TraceOut_status[249] := BenchUut6.status;
   BenchCalls := BenchCalls + 1;
 250:
   BenchUut6.cyclicExecution := FALSE;
   BenchUut6.trigger := TRUE;
   BenchUut6.value := LREAL#4.0;
   BenchUut6.windowSize := INT#100;
   BenchUut6.reset := FALSE;
   TraceIn_cyclicExecution[250] := BenchUut6.cyclicExecution;
   TraceIn_trigger[250] := BenchUut6.trigger;
   TraceIn_value[250] := BenchUut6.value;
   TraceIn_windowSize[250] := BenchUut6.windowSize;
   TraceIn_reset[250] := BenchUut6.reset;
   BenchUut6();
   TraceOut_average[250] := BenchUut6.average;
   TraceOut_windowSizeReached[250] := BenchUut6.windowSizeReached;
   TraceOut_error[250] := BenchUut6.error;
   TraceOut_status[250] := BenchUut6.status;
   BenchCalls := BenchCalls + 1;
 251:
   BenchUut6.cyclicExecution := FALSE;
   BenchUut6.trigger := FALSE;
   BenchUut6.value := LREAL#4.0;
   BenchUut6.windowSize := INT#100;
   BenchUut6.reset := FALSE;
   TraceIn_cyclicExecution[251] := BenchUut6.cyclicExecution;
   TraceIn_trigger[251] := BenchUut6.trigger;
   TraceIn_value[251] := BenchUut6.value;
   TraceIn_windowSize[251] := BenchUut6.windowSize;
   TraceIn_reset[251] := BenchUut6.reset;
   BenchUut6();
   TraceOut_average[251] := BenchUut6.average;
   TraceOut_windowSizeReached[251] := BenchUut6.windowSizeReached;
   TraceOut_error[251] := BenchUut6.error;
   TraceOut_status[251] := BenchUut6.status;
   BenchCalls := BenchCalls + 1;
 252:
   BenchUut6.cyclicExecution := FALSE;
   BenchUut6.trigger := TRUE;
   BenchUut6.value := LREAL#5.0;
   BenchUut6.windowSize := INT#100;
   BenchUut6.reset := FALSE;
   TraceIn_cyclicExecution[252] := BenchUut6.cyclicExecution;
   TraceIn_trigger[252] := BenchUut6.trigger;
   TraceIn_value[252] := BenchUut6.value;
   TraceIn_windowSize[252] := BenchUut6.windowSize;
   TraceIn_reset[252] := BenchUut6.reset;
   BenchUut6();
   TraceOut_average[252] := BenchUut6.average;
   TraceOut_windowSizeReached[252] := BenchUut6.windowSizeReached;
   TraceOut_error[252] := BenchUut6.error;
   TraceOut_status[252] := BenchUut6.status;
   BenchCalls := BenchCalls + 1;
 253:
   BenchUut6.cyclicExecution := FALSE;
   BenchUut6.trigger := FALSE;
   BenchUut6.value := LREAL#5.0;
   BenchUut6.windowSize := INT#100;
   BenchUut6.reset := FALSE;
   TraceIn_cyclicExecution[253] := BenchUut6.cyclicExecution;
   TraceIn_trigger[253] := BenchUut6.trigger;
   TraceIn_value[253] := BenchUut6.value;
   TraceIn_windowSize[253] := BenchUut6.windowSize;
   TraceIn_reset[253] := BenchUut6.reset;
   BenchUut6();
   TraceOut_average[253] := BenchUut6.average;
   TraceOut_windowSizeReached[253] := BenchUut6.windowSizeReached;
   TraceOut_error[253] := BenchUut6.error;
   TraceOut_status[253] := BenchUut6.status;
   BenchCalls := BenchCalls + 1;
 254:
   BenchUut6.cyclicExecution := FALSE;
   BenchUut6.trigger := TRUE;
   BenchUut6.value := LREAL#6.0;
   BenchUut6.windowSize := INT#100;
   BenchUut6.reset := FALSE;
   TraceIn_cyclicExecution[254] := BenchUut6.cyclicExecution;
   TraceIn_trigger[254] := BenchUut6.trigger;
   TraceIn_value[254] := BenchUut6.value;
   TraceIn_windowSize[254] := BenchUut6.windowSize;
   TraceIn_reset[254] := BenchUut6.reset;
   BenchUut6();
   TraceOut_average[254] := BenchUut6.average;
   TraceOut_windowSizeReached[254] := BenchUut6.windowSizeReached;
   TraceOut_error[254] := BenchUut6.error;
   TraceOut_status[254] := BenchUut6.status;
   BenchCalls := BenchCalls + 1;
 255:
   BenchUut6.cyclicExecution := FALSE;
   BenchUut6.trigger := FALSE;
   BenchUut6.value := LREAL#6.0;
   BenchUut6.windowSize := INT#100;
   BenchUut6.reset := FALSE;
   TraceIn_cyclicExecution[255] := BenchUut6.cyclicExecution;
   TraceIn_trigger[255] := BenchUut6.trigger;
   TraceIn_value[255] := BenchUut6.value;
   TraceIn_windowSize[255] := BenchUut6.windowSize;
   TraceIn_reset[255] := BenchUut6.reset;
   BenchUut6();
   TraceOut_average[255] := BenchUut6.average;
   TraceOut_windowSizeReached[255] := BenchUut6.windowSizeReached;
   TraceOut_error[255] := BenchUut6.error;
   TraceOut_status[255] := BenchUut6.status;
   BenchCalls := BenchCalls + 1;
 256:
   BenchUut6.cyclicExecution := FALSE;
   BenchUut6.trigger := TRUE;
   BenchUut6.value := LREAL#7.0;
   BenchUut6.windowSize := INT#100;
   BenchUut6.reset := FALSE;
   TraceIn_cyclicExecution[256] := BenchUut6.cyclicExecution;
   TraceIn_trigger[256] := BenchUut6.trigger;
   TraceIn_value[256] := BenchUut6.value;
   TraceIn_windowSize[256] := BenchUut6.windowSize;
   TraceIn_reset[256] := BenchUut6.reset;
   BenchUut6();
   TraceOut_average[256] := BenchUut6.average;
   TraceOut_windowSizeReached[256] := BenchUut6.windowSizeReached;
   TraceOut_error[256] := BenchUut6.error;
   TraceOut_status[256] := BenchUut6.status;
   BenchCalls := BenchCalls + 1;
 257:
   BenchUut6.cyclicExecution := FALSE;
   BenchUut6.trigger := FALSE;
   BenchUut6.value := LREAL#7.0;
   BenchUut6.windowSize := INT#100;
   BenchUut6.reset := FALSE;
   TraceIn_cyclicExecution[257] := BenchUut6.cyclicExecution;
   TraceIn_trigger[257] := BenchUut6.trigger;
   TraceIn_value[257] := BenchUut6.value;
   TraceIn_windowSize[257] := BenchUut6.windowSize;
   TraceIn_reset[257] := BenchUut6.reset;
   BenchUut6();
   TraceOut_average[257] := BenchUut6.average;
   TraceOut_windowSizeReached[257] := BenchUut6.windowSizeReached;
   TraceOut_error[257] := BenchUut6.error;
   TraceOut_status[257] := BenchUut6.status;
   BenchCalls := BenchCalls + 1;
 258:
   BenchUut6.cyclicExecution := FALSE;
   BenchUut6.trigger := TRUE;
   BenchUut6.value := LREAL#8.0;
   BenchUut6.windowSize := INT#100;
   BenchUut6.reset := FALSE;
   TraceIn_cyclicExecution[258] := BenchUut6.cyclicExecution;
   TraceIn_trigger[258] := BenchUut6.trigger;
   TraceIn_value[258] := BenchUut6.value;
   TraceIn_windowSize[258] := BenchUut6.windowSize;
   TraceIn_reset[258] := BenchUut6.reset;
   BenchUut6();
   TraceOut_average[258] := BenchUut6.average;
   TraceOut_windowSizeReached[258] := BenchUut6.windowSizeReached;
   TraceOut_error[258] := BenchUut6.error;
   TraceOut_status[258] := BenchUut6.status;
   BenchCalls := BenchCalls + 1;
 259:
   BenchUut6.cyclicExecution := FALSE;
   BenchUut6.trigger := FALSE;
   BenchUut6.value := LREAL#8.0;
   BenchUut6.windowSize := INT#100;
   BenchUut6.reset := FALSE;
   TraceIn_cyclicExecution[259] := BenchUut6.cyclicExecution;
   TraceIn_trigger[259] := BenchUut6.trigger;
   TraceIn_value[259] := BenchUut6.value;
   TraceIn_windowSize[259] := BenchUut6.windowSize;
   TraceIn_reset[259] := BenchUut6.reset;
   BenchUut6();
   TraceOut_average[259] := BenchUut6.average;
   TraceOut_windowSizeReached[259] := BenchUut6.windowSizeReached;
   TraceOut_error[259] := BenchUut6.error;
   TraceOut_status[259] := BenchUut6.status;
   BenchCalls := BenchCalls + 1;
 260:
   BenchUut6.cyclicExecution := FALSE;
   BenchUut6.trigger := TRUE;
   BenchUut6.value := LREAL#9.0;
   BenchUut6.windowSize := INT#100;
   BenchUut6.reset := FALSE;
   TraceIn_cyclicExecution[260] := BenchUut6.cyclicExecution;
   TraceIn_trigger[260] := BenchUut6.trigger;
   TraceIn_value[260] := BenchUut6.value;
   TraceIn_windowSize[260] := BenchUut6.windowSize;
   TraceIn_reset[260] := BenchUut6.reset;
   BenchUut6();
   TraceOut_average[260] := BenchUut6.average;
   TraceOut_windowSizeReached[260] := BenchUut6.windowSizeReached;
   TraceOut_error[260] := BenchUut6.error;
   TraceOut_status[260] := BenchUut6.status;
   BenchCalls := BenchCalls + 1;
 261:
   BenchUut6.cyclicExecution := FALSE;
   BenchUut6.trigger := FALSE;
   BenchUut6.value := LREAL#9.0;
   BenchUut6.windowSize := INT#100;
   BenchUut6.reset := FALSE;
   TraceIn_cyclicExecution[261] := BenchUut6.cyclicExecution;
   TraceIn_trigger[261] := BenchUut6.trigger;
   TraceIn_value[261] := BenchUut6.value;
   TraceIn_windowSize[261] := BenchUut6.windowSize;
   TraceIn_reset[261] := BenchUut6.reset;
   BenchUut6();
   TraceOut_average[261] := BenchUut6.average;
   TraceOut_windowSizeReached[261] := BenchUut6.windowSizeReached;
   TraceOut_error[261] := BenchUut6.error;
   TraceOut_status[261] := BenchUut6.status;
   BenchCalls := BenchCalls + 1;
 262:
   BenchUut6.cyclicExecution := FALSE;
   BenchUut6.trigger := TRUE;
   BenchUut6.value := LREAL#10.0;
   BenchUut6.windowSize := INT#100;
   BenchUut6.reset := FALSE;
   TraceIn_cyclicExecution[262] := BenchUut6.cyclicExecution;
   TraceIn_trigger[262] := BenchUut6.trigger;
   TraceIn_value[262] := BenchUut6.value;
   TraceIn_windowSize[262] := BenchUut6.windowSize;
   TraceIn_reset[262] := BenchUut6.reset;
   BenchUut6();
   TraceOut_average[262] := BenchUut6.average;
   TraceOut_windowSizeReached[262] := BenchUut6.windowSizeReached;
   TraceOut_error[262] := BenchUut6.error;
   TraceOut_status[262] := BenchUut6.status;
   BenchCalls := BenchCalls + 1;
 263:
   BenchUut6.cyclicExecution := FALSE;
   BenchUut6.trigger := FALSE;
   BenchUut6.value := LREAL#10.0;
   BenchUut6.windowSize := INT#100;
   BenchUut6.reset := FALSE;
   TraceIn_cyclicExecution[263] := BenchUut6.cyclicExecution;
   TraceIn_trigger[263] := BenchUut6.trigger;
   TraceIn_value[263] := BenchUut6.value;
   TraceIn_windowSize[263] := BenchUut6.windowSize;
   TraceIn_reset[263] := BenchUut6.reset;
   BenchUut6();
   TraceOut_average[263] := BenchUut6.average;
   TraceOut_windowSizeReached[263] := BenchUut6.windowSizeReached;
   TraceOut_error[263] := BenchUut6.error;
   TraceOut_status[263] := BenchUut6.status;
   BenchCalls := BenchCalls + 1;
 264:
   BenchUut6.cyclicExecution := FALSE;
   BenchUut6.trigger := TRUE;
   BenchUut6.value := LREAL#11.0;
   BenchUut6.windowSize := INT#100;
   BenchUut6.reset := FALSE;
   TraceIn_cyclicExecution[264] := BenchUut6.cyclicExecution;
   TraceIn_trigger[264] := BenchUut6.trigger;
   TraceIn_value[264] := BenchUut6.value;
   TraceIn_windowSize[264] := BenchUut6.windowSize;
   TraceIn_reset[264] := BenchUut6.reset;
   BenchUut6();
   TraceOut_average[264] := BenchUut6.average;
   TraceOut_windowSizeReached[264] := BenchUut6.windowSizeReached;
   TraceOut_error[264] := BenchUut6.error;
   TraceOut_status[264] := BenchUut6.status;
   BenchCalls := BenchCalls + 1;
 265:
   BenchUut6.cyclicExecution := FALSE;
   BenchUut6.trigger := FALSE;
   BenchUut6.value := LREAL#11.0;
   BenchUut6.windowSize := INT#100;
   BenchUut6.reset := FALSE;
   TraceIn_cyclicExecution[265] := BenchUut6.cyclicExecution;
   TraceIn_trigger[265] := BenchUut6.trigger;
   TraceIn_value[265] := BenchUut6.value;
   TraceIn_windowSize[265] := BenchUut6.windowSize;
   TraceIn_reset[265] := BenchUut6.reset;
   BenchUut6();
   TraceOut_average[265] := BenchUut6.average;
   TraceOut_windowSizeReached[265] := BenchUut6.windowSizeReached;
   TraceOut_error[265] := BenchUut6.error;
   TraceOut_status[265] := BenchUut6.status;
   BenchCalls := BenchCalls + 1;
 266:
   BenchUut6.cyclicExecution := FALSE;
   BenchUut6.trigger := TRUE;
   BenchUut6.value := LREAL#12.0;
   BenchUut6.windowSize := INT#100;
   BenchUut6.reset := FALSE;
   TraceIn_cyclicExecution[266] := BenchUut6.cyclicExecution;
   TraceIn_trigger[266] := BenchUut6.trigger;
   TraceIn_value[266] := BenchUut6.value;
   TraceIn_windowSize[266] := BenchUut6.windowSize;
   TraceIn_reset[266] := BenchUut6.reset;
   BenchUut6();
   TraceOut_average[266] := BenchUut6.average;
   TraceOut_windowSizeReached[266] := BenchUut6.windowSizeReached;
   TraceOut_error[266] := BenchUut6.error;
   TraceOut_status[266] := BenchUut6.status;
   BenchCalls := BenchCalls + 1;
 267:
   BenchUut6.cyclicExecution := FALSE;
   BenchUut6.trigger := FALSE;
   BenchUut6.value := LREAL#12.0;
   BenchUut6.windowSize := INT#100;
   BenchUut6.reset := FALSE;
   TraceIn_cyclicExecution[267] := BenchUut6.cyclicExecution;
   TraceIn_trigger[267] := BenchUut6.trigger;
   TraceIn_value[267] := BenchUut6.value;
   TraceIn_windowSize[267] := BenchUut6.windowSize;
   TraceIn_reset[267] := BenchUut6.reset;
   BenchUut6();
   TraceOut_average[267] := BenchUut6.average;
   TraceOut_windowSizeReached[267] := BenchUut6.windowSizeReached;
   TraceOut_error[267] := BenchUut6.error;
   TraceOut_status[267] := BenchUut6.status;
   BenchCalls := BenchCalls + 1;
 268:
   BenchUut6.cyclicExecution := FALSE;
   BenchUut6.trigger := TRUE;
   BenchUut6.value := LREAL#13.0;
   BenchUut6.windowSize := INT#100;
   BenchUut6.reset := FALSE;
   TraceIn_cyclicExecution[268] := BenchUut6.cyclicExecution;
   TraceIn_trigger[268] := BenchUut6.trigger;
   TraceIn_value[268] := BenchUut6.value;
   TraceIn_windowSize[268] := BenchUut6.windowSize;
   TraceIn_reset[268] := BenchUut6.reset;
   BenchUut6();
   TraceOut_average[268] := BenchUut6.average;
   TraceOut_windowSizeReached[268] := BenchUut6.windowSizeReached;
   TraceOut_error[268] := BenchUut6.error;
   TraceOut_status[268] := BenchUut6.status;
   BenchCalls := BenchCalls + 1;
 269:
   BenchUut6.cyclicExecution := FALSE;
   BenchUut6.trigger := FALSE;
   BenchUut6.value := LREAL#13.0;
   BenchUut6.windowSize := INT#100;
   BenchUut6.reset := FALSE;
   TraceIn_cyclicExecution[269] := BenchUut6.cyclicExecution;
   TraceIn_trigger[269] := BenchUut6.trigger;
   TraceIn_value[269] := BenchUut6.value;
   TraceIn_windowSize[269] := BenchUut6.windowSize;
   TraceIn_reset[269] := BenchUut6.reset;
   BenchUut6();
   TraceOut_average[269] := BenchUut6.average;
   TraceOut_windowSizeReached[269] := BenchUut6.windowSizeReached;
   TraceOut_error[269] := BenchUut6.error;
   TraceOut_status[269] := BenchUut6.status;
   BenchCalls := BenchCalls + 1;
 270:
   BenchUut6.cyclicExecution := FALSE;
   BenchUut6.trigger := TRUE;
   BenchUut6.value := LREAL#14.0;
   BenchUut6.windowSize := INT#100;
   BenchUut6.reset := FALSE;
   TraceIn_cyclicExecution[270] := BenchUut6.cyclicExecution;
   TraceIn_trigger[270] := BenchUut6.trigger;
   TraceIn_value[270] := BenchUut6.value;
   TraceIn_windowSize[270] := BenchUut6.windowSize;
   TraceIn_reset[270] := BenchUut6.reset;
   BenchUut6();
   TraceOut_average[270] := BenchUut6.average;
   TraceOut_windowSizeReached[270] := BenchUut6.windowSizeReached;
   TraceOut_error[270] := BenchUut6.error;
   TraceOut_status[270] := BenchUut6.status;
   BenchCalls := BenchCalls + 1;
 271:
   BenchUut6.cyclicExecution := FALSE;
   BenchUut6.trigger := FALSE;
   BenchUut6.value := LREAL#14.0;
   BenchUut6.windowSize := INT#100;
   BenchUut6.reset := FALSE;
   TraceIn_cyclicExecution[271] := BenchUut6.cyclicExecution;
   TraceIn_trigger[271] := BenchUut6.trigger;
   TraceIn_value[271] := BenchUut6.value;
   TraceIn_windowSize[271] := BenchUut6.windowSize;
   TraceIn_reset[271] := BenchUut6.reset;
   BenchUut6();
   TraceOut_average[271] := BenchUut6.average;
   TraceOut_windowSizeReached[271] := BenchUut6.windowSizeReached;
   TraceOut_error[271] := BenchUut6.error;
   TraceOut_status[271] := BenchUut6.status;
   BenchCalls := BenchCalls + 1;
 272:
   BenchUut6.cyclicExecution := FALSE;
   BenchUut6.trigger := TRUE;
   BenchUut6.value := LREAL#15.0;
   BenchUut6.windowSize := INT#100;
   BenchUut6.reset := FALSE;
   TraceIn_cyclicExecution[272] := BenchUut6.cyclicExecution;
   TraceIn_trigger[272] := BenchUut6.trigger;
   TraceIn_value[272] := BenchUut6.value;
   TraceIn_windowSize[272] := BenchUut6.windowSize;
   TraceIn_reset[272] := BenchUut6.reset;
   BenchUut6();
   TraceOut_average[272] := BenchUut6.average;
   TraceOut_windowSizeReached[272] := BenchUut6.windowSizeReached;
   TraceOut_error[272] := BenchUut6.error;
   TraceOut_status[272] := BenchUut6.status;
   BenchCalls := BenchCalls + 1;
 273:
   BenchUut6.cyclicExecution := FALSE;
   BenchUut6.trigger := FALSE;
   BenchUut6.value := LREAL#15.0;
   BenchUut6.windowSize := INT#100;
   BenchUut6.reset := FALSE;
   TraceIn_cyclicExecution[273] := BenchUut6.cyclicExecution;
   TraceIn_trigger[273] := BenchUut6.trigger;
   TraceIn_value[273] := BenchUut6.value;
   TraceIn_windowSize[273] := BenchUut6.windowSize;
   TraceIn_reset[273] := BenchUut6.reset;
   BenchUut6();
   TraceOut_average[273] := BenchUut6.average;
   TraceOut_windowSizeReached[273] := BenchUut6.windowSizeReached;
   TraceOut_error[273] := BenchUut6.error;
   TraceOut_status[273] := BenchUut6.status;
   BenchCalls := BenchCalls + 1;
 274:
   BenchUut6.cyclicExecution := FALSE;
   BenchUut6.trigger := TRUE;
   BenchUut6.value := LREAL#16.0;
   BenchUut6.windowSize := INT#100;
   BenchUut6.reset := FALSE;
   TraceIn_cyclicExecution[274] := BenchUut6.cyclicExecution;
   TraceIn_trigger[274] := BenchUut6.trigger;
   TraceIn_value[274] := BenchUut6.value;
   TraceIn_windowSize[274] := BenchUut6.windowSize;
   TraceIn_reset[274] := BenchUut6.reset;
   BenchUut6();
   TraceOut_average[274] := BenchUut6.average;
   TraceOut_windowSizeReached[274] := BenchUut6.windowSizeReached;
   TraceOut_error[274] := BenchUut6.error;
   TraceOut_status[274] := BenchUut6.status;
   BenchCalls := BenchCalls + 1;
 275:
   BenchUut6.cyclicExecution := FALSE;
   BenchUut6.trigger := FALSE;
   BenchUut6.value := LREAL#16.0;
   BenchUut6.windowSize := INT#100;
   BenchUut6.reset := FALSE;
   TraceIn_cyclicExecution[275] := BenchUut6.cyclicExecution;
   TraceIn_trigger[275] := BenchUut6.trigger;
   TraceIn_value[275] := BenchUut6.value;
   TraceIn_windowSize[275] := BenchUut6.windowSize;
   TraceIn_reset[275] := BenchUut6.reset;
   BenchUut6();
   TraceOut_average[275] := BenchUut6.average;
   TraceOut_windowSizeReached[275] := BenchUut6.windowSizeReached;
   TraceOut_error[275] := BenchUut6.error;
   TraceOut_status[275] := BenchUut6.status;
   BenchCalls := BenchCalls + 1;
 276:
   BenchUut6.cyclicExecution := FALSE;
   BenchUut6.trigger := TRUE;
   BenchUut6.value := LREAL#17.0;
   BenchUut6.windowSize := INT#100;
   BenchUut6.reset := FALSE;
   TraceIn_cyclicExecution[276] := BenchUut6.cyclicExecution;
   TraceIn_trigger[276] := BenchUut6.trigger;
   TraceIn_value[276] := BenchUut6.value;
   TraceIn_windowSize[276] := BenchUut6.windowSize;
   TraceIn_reset[276] := BenchUut6.reset;
   BenchUut6();
   TraceOut_average[276] := BenchUut6.average;
   TraceOut_windowSizeReached[276] := BenchUut6.windowSizeReached;
   TraceOut_error[276] := BenchUut6.error;
   TraceOut_status[276] := BenchUut6.status;
   BenchCalls := BenchCalls + 1;
 277:
   BenchUut6.cyclicExecution := FALSE;
   BenchUut6.trigger := FALSE;
   BenchUut6.value := LREAL#17.0;
   BenchUut6.windowSize := INT#100;
   BenchUut6.reset := FALSE;
   TraceIn_cyclicExecution[277] := BenchUut6.cyclicExecution;
   TraceIn_trigger[277] := BenchUut6.trigger;
   TraceIn_value[277] := BenchUut6.value;
   TraceIn_windowSize[277] := BenchUut6.windowSize;
   TraceIn_reset[277] := BenchUut6.reset;
   BenchUut6();
   TraceOut_average[277] := BenchUut6.average;
   TraceOut_windowSizeReached[277] := BenchUut6.windowSizeReached;
   TraceOut_error[277] := BenchUut6.error;
   TraceOut_status[277] := BenchUut6.status;
   BenchCalls := BenchCalls + 1;
 278:
   BenchUut6.cyclicExecution := FALSE;
   BenchUut6.trigger := TRUE;
   BenchUut6.value := LREAL#18.0;
   BenchUut6.windowSize := INT#100;
   BenchUut6.reset := FALSE;
   TraceIn_cyclicExecution[278] := BenchUut6.cyclicExecution;
   TraceIn_trigger[278] := BenchUut6.trigger;
   TraceIn_value[278] := BenchUut6.value;
   TraceIn_windowSize[278] := BenchUut6.windowSize;
   TraceIn_reset[278] := BenchUut6.reset;
   BenchUut6();
   TraceOut_average[278] := BenchUut6.average;
   TraceOut_windowSizeReached[278] := BenchUut6.windowSizeReached;
   TraceOut_error[278] := BenchUut6.error;
   TraceOut_status[278] := BenchUut6.status;
   BenchCalls := BenchCalls + 1;
 279:
   BenchUut6.cyclicExecution := FALSE;
   BenchUut6.trigger := FALSE;
   BenchUut6.value := LREAL#18.0;
   BenchUut6.windowSize := INT#100;
   BenchUut6.reset := FALSE;
   TraceIn_cyclicExecution[279] := BenchUut6.cyclicExecution;
   TraceIn_trigger[279] := BenchUut6.trigger;
   TraceIn_value[279] := BenchUut6.value;
   TraceIn_windowSize[279] := BenchUut6.windowSize;
   TraceIn_reset[279] := BenchUut6.reset;
   BenchUut6();
   TraceOut_average[279] := BenchUut6.average;
   TraceOut_windowSizeReached[279] := BenchUut6.windowSizeReached;
   TraceOut_error[279] := BenchUut6.error;
   TraceOut_status[279] := BenchUut6.status;
   BenchCalls := BenchCalls + 1;
 280:
   BenchUut6.cyclicExecution := FALSE;
   BenchUut6.trigger := TRUE;
   BenchUut6.value := LREAL#19.0;
   BenchUut6.windowSize := INT#100;
   BenchUut6.reset := FALSE;
   TraceIn_cyclicExecution[280] := BenchUut6.cyclicExecution;
   TraceIn_trigger[280] := BenchUut6.trigger;
   TraceIn_value[280] := BenchUut6.value;
   TraceIn_windowSize[280] := BenchUut6.windowSize;
   TraceIn_reset[280] := BenchUut6.reset;
   BenchUut6();
   TraceOut_average[280] := BenchUut6.average;
   TraceOut_windowSizeReached[280] := BenchUut6.windowSizeReached;
   TraceOut_error[280] := BenchUut6.error;
   TraceOut_status[280] := BenchUut6.status;
   BenchCalls := BenchCalls + 1;
 281:
   BenchUut6.cyclicExecution := FALSE;
   BenchUut6.trigger := FALSE;
   BenchUut6.value := LREAL#19.0;
   BenchUut6.windowSize := INT#100;
   BenchUut6.reset := FALSE;
   TraceIn_cyclicExecution[281] := BenchUut6.cyclicExecution;
   TraceIn_trigger[281] := BenchUut6.trigger;
   TraceIn_value[281] := BenchUut6.value;
   TraceIn_windowSize[281] := BenchUut6.windowSize;
   TraceIn_reset[281] := BenchUut6.reset;
   BenchUut6();
   TraceOut_average[281] := BenchUut6.average;
   TraceOut_windowSizeReached[281] := BenchUut6.windowSizeReached;
   TraceOut_error[281] := BenchUut6.error;
   TraceOut_status[281] := BenchUut6.status;
   BenchCalls := BenchCalls + 1;
 282:
   BenchUut6.cyclicExecution := FALSE;
   BenchUut6.trigger := TRUE;
   BenchUut6.value := LREAL#20.0;
   BenchUut6.windowSize := INT#100;
   BenchUut6.reset := FALSE;
   TraceIn_cyclicExecution[282] := BenchUut6.cyclicExecution;
   TraceIn_trigger[282] := BenchUut6.trigger;
   TraceIn_value[282] := BenchUut6.value;
   TraceIn_windowSize[282] := BenchUut6.windowSize;
   TraceIn_reset[282] := BenchUut6.reset;
   BenchUut6();
   TraceOut_average[282] := BenchUut6.average;
   TraceOut_windowSizeReached[282] := BenchUut6.windowSizeReached;
   TraceOut_error[282] := BenchUut6.error;
   TraceOut_status[282] := BenchUut6.status;
   BenchCalls := BenchCalls + 1;
 283:
   BenchUut6.cyclicExecution := FALSE;
   BenchUut6.trigger := FALSE;
   BenchUut6.value := LREAL#20.0;
   BenchUut6.windowSize := INT#100;
   BenchUut6.reset := FALSE;
   TraceIn_cyclicExecution[283] := BenchUut6.cyclicExecution;
   TraceIn_trigger[283] := BenchUut6.trigger;
   TraceIn_value[283] := BenchUut6.value;
   TraceIn_windowSize[283] := BenchUut6.windowSize;
   TraceIn_reset[283] := BenchUut6.reset;
   BenchUut6();
   TraceOut_average[283] := BenchUut6.average;
   TraceOut_windowSizeReached[283] := BenchUut6.windowSizeReached;
   TraceOut_error[283] := BenchUut6.error;
   TraceOut_status[283] := BenchUut6.status;
   BenchCalls := BenchCalls + 1;
 284:
   BenchUut6.cyclicExecution := FALSE;
   BenchUut6.trigger := TRUE;
   BenchUut6.value := LREAL#21.0;
   BenchUut6.windowSize := INT#100;
   BenchUut6.reset := FALSE;
   TraceIn_cyclicExecution[284] := BenchUut6.cyclicExecution;
   TraceIn_trigger[284] := BenchUut6.trigger;
   TraceIn_value[284] := BenchUut6.value;
   TraceIn_windowSize[284] := BenchUut6.windowSize;
   TraceIn_reset[284] := BenchUut6.reset;
   BenchUut6();
   TraceOut_average[284] := BenchUut6.average;
   TraceOut_windowSizeReached[284] := BenchUut6.windowSizeReached;
   TraceOut_error[284] := BenchUut6.error;
   TraceOut_status[284] := BenchUut6.status;
   BenchCalls := BenchCalls + 1;
 285:
   BenchUut6.cyclicExecution := FALSE;
   BenchUut6.trigger := FALSE;
   BenchUut6.value := LREAL#21.0;
   BenchUut6.windowSize := INT#100;
   BenchUut6.reset := FALSE;
   TraceIn_cyclicExecution[285] := BenchUut6.cyclicExecution;
   TraceIn_trigger[285] := BenchUut6.trigger;
   TraceIn_value[285] := BenchUut6.value;
   TraceIn_windowSize[285] := BenchUut6.windowSize;
   TraceIn_reset[285] := BenchUut6.reset;
   BenchUut6();
   TraceOut_average[285] := BenchUut6.average;
   TraceOut_windowSizeReached[285] := BenchUut6.windowSizeReached;
   TraceOut_error[285] := BenchUut6.error;
   TraceOut_status[285] := BenchUut6.status;
   BenchCalls := BenchCalls + 1;
 286:
   BenchUut6.cyclicExecution := FALSE;
   BenchUut6.trigger := TRUE;
   BenchUut6.value := LREAL#22.0;
   BenchUut6.windowSize := INT#100;
   BenchUut6.reset := FALSE;
   TraceIn_cyclicExecution[286] := BenchUut6.cyclicExecution;
   TraceIn_trigger[286] := BenchUut6.trigger;
   TraceIn_value[286] := BenchUut6.value;
   TraceIn_windowSize[286] := BenchUut6.windowSize;
   TraceIn_reset[286] := BenchUut6.reset;
   BenchUut6();
   TraceOut_average[286] := BenchUut6.average;
   TraceOut_windowSizeReached[286] := BenchUut6.windowSizeReached;
   TraceOut_error[286] := BenchUut6.error;
   TraceOut_status[286] := BenchUut6.status;
   BenchCalls := BenchCalls + 1;
 287:
   BenchUut6.cyclicExecution := FALSE;
   BenchUut6.trigger := FALSE;
   BenchUut6.value := LREAL#22.0;
   BenchUut6.windowSize := INT#100;
   BenchUut6.reset := FALSE;
   TraceIn_cyclicExecution[287] := BenchUut6.cyclicExecution;
   TraceIn_trigger[287] := BenchUut6.trigger;
   TraceIn_value[287] := BenchUut6.value;
   TraceIn_windowSize[287] := BenchUut6.windowSize;
   TraceIn_reset[287] := BenchUut6.reset;
   BenchUut6();
   TraceOut_average[287] := BenchUut6.average;
   TraceOut_windowSizeReached[287] := BenchUut6.windowSizeReached;
   TraceOut_error[287] := BenchUut6.error;
   TraceOut_status[287] := BenchUut6.status;
   BenchCalls := BenchCalls + 1;
 288:
   BenchUut6.cyclicExecution := FALSE;
   BenchUut6.trigger := TRUE;
   BenchUut6.value := LREAL#23.0;
   BenchUut6.windowSize := INT#100;
   BenchUut6.reset := FALSE;
   TraceIn_cyclicExecution[288] := BenchUut6.cyclicExecution;
   TraceIn_trigger[288] := BenchUut6.trigger;
   TraceIn_value[288] := BenchUut6.value;
   TraceIn_windowSize[288] := BenchUut6.windowSize;
   TraceIn_reset[288] := BenchUut6.reset;
   BenchUut6();
   TraceOut_average[288] := BenchUut6.average;
   TraceOut_windowSizeReached[288] := BenchUut6.windowSizeReached;
   TraceOut_error[288] := BenchUut6.error;
   TraceOut_status[288] := BenchUut6.status;
   BenchCalls := BenchCalls + 1;
 289:
   BenchUut6.cyclicExecution := FALSE;
   BenchUut6.trigger := FALSE;
   BenchUut6.value := LREAL#23.0;
   BenchUut6.windowSize := INT#100;
   BenchUut6.reset := FALSE;
   TraceIn_cyclicExecution[289] := BenchUut6.cyclicExecution;
   TraceIn_trigger[289] := BenchUut6.trigger;
   TraceIn_value[289] := BenchUut6.value;
   TraceIn_windowSize[289] := BenchUut6.windowSize;
   TraceIn_reset[289] := BenchUut6.reset;
   BenchUut6();
   TraceOut_average[289] := BenchUut6.average;
   TraceOut_windowSizeReached[289] := BenchUut6.windowSizeReached;
   TraceOut_error[289] := BenchUut6.error;
   TraceOut_status[289] := BenchUut6.status;
   BenchCalls := BenchCalls + 1;
 290:
   BenchUut6.cyclicExecution := FALSE;
   BenchUut6.trigger := TRUE;
   BenchUut6.value := LREAL#24.0;
   BenchUut6.windowSize := INT#100;
   BenchUut6.reset := FALSE;
   TraceIn_cyclicExecution[290] := BenchUut6.cyclicExecution;
   TraceIn_trigger[290] := BenchUut6.trigger;
   TraceIn_value[290] := BenchUut6.value;
   TraceIn_windowSize[290] := BenchUut6.windowSize;
   TraceIn_reset[290] := BenchUut6.reset;
   BenchUut6();
   TraceOut_average[290] := BenchUut6.average;
   TraceOut_windowSizeReached[290] := BenchUut6.windowSizeReached;
   TraceOut_error[290] := BenchUut6.error;
   TraceOut_status[290] := BenchUut6.status;
   BenchCalls := BenchCalls + 1;
 291:
   BenchUut6.cyclicExecution := FALSE;
   BenchUut6.trigger := FALSE;
   BenchUut6.value := LREAL#24.0;
   BenchUut6.windowSize := INT#100;
   BenchUut6.reset := FALSE;
   TraceIn_cyclicExecution[291] := BenchUut6.cyclicExecution;
   TraceIn_trigger[291] := BenchUut6.trigger;
   TraceIn_value[291] := BenchUut6.value;
   TraceIn_windowSize[291] := BenchUut6.windowSize;
   TraceIn_reset[291] := BenchUut6.reset;
   BenchUut6();
   TraceOut_average[291] := BenchUut6.average;
   TraceOut_windowSizeReached[291] := BenchUut6.windowSizeReached;
   TraceOut_error[291] := BenchUut6.error;
   TraceOut_status[291] := BenchUut6.status;
   BenchCalls := BenchCalls + 1;
 292:
   BenchUut6.cyclicExecution := FALSE;
   BenchUut6.trigger := TRUE;
   BenchUut6.value := LREAL#25.0;
   BenchUut6.windowSize := INT#100;
   BenchUut6.reset := FALSE;
   TraceIn_cyclicExecution[292] := BenchUut6.cyclicExecution;
   TraceIn_trigger[292] := BenchUut6.trigger;
   TraceIn_value[292] := BenchUut6.value;
   TraceIn_windowSize[292] := BenchUut6.windowSize;
   TraceIn_reset[292] := BenchUut6.reset;
   BenchUut6();
   TraceOut_average[292] := BenchUut6.average;
   TraceOut_windowSizeReached[292] := BenchUut6.windowSizeReached;
   TraceOut_error[292] := BenchUut6.error;
   TraceOut_status[292] := BenchUut6.status;
   BenchCalls := BenchCalls + 1;
 293:
   BenchUut6.cyclicExecution := FALSE;
   BenchUut6.trigger := FALSE;
   BenchUut6.value := LREAL#25.0;
   BenchUut6.windowSize := INT#100;
   BenchUut6.reset := FALSE;
   TraceIn_cyclicExecution[293] := BenchUut6.cyclicExecution;
   TraceIn_trigger[293] := BenchUut6.trigger;
   TraceIn_value[293] := BenchUut6.value;
   TraceIn_windowSize[293] := BenchUut6.windowSize;
   TraceIn_reset[293] := BenchUut6.reset;
   BenchUut6();
   TraceOut_average[293] := BenchUut6.average;
   TraceOut_windowSizeReached[293] := BenchUut6.windowSizeReached;
   TraceOut_error[293] := BenchUut6.error;
   TraceOut_status[293] := BenchUut6.status;
   BenchCalls := BenchCalls + 1;
 294:
   BenchUut6.cyclicExecution := FALSE;
   BenchUut6.trigger := TRUE;
   BenchUut6.value := LREAL#26.0;
   BenchUut6.windowSize := INT#100;
   BenchUut6.reset := FALSE;
   TraceIn_cyclicExecution[294] := BenchUut6.cyclicExecution;
   TraceIn_trigger[294] := BenchUut6.trigger;
   TraceIn_value[294] := BenchUut6.value;
   TraceIn_windowSize[294] := BenchUut6.windowSize;
   TraceIn_reset[294] := BenchUut6.reset;
   BenchUut6();
   TraceOut_average[294] := BenchUut6.average;
   TraceOut_windowSizeReached[294] := BenchUut6.windowSizeReached;
   TraceOut_error[294] := BenchUut6.error;
   TraceOut_status[294] := BenchUut6.status;
   BenchCalls := BenchCalls + 1;
 295:
   BenchUut6.cyclicExecution := FALSE;
   BenchUut6.trigger := FALSE;
   BenchUut6.value := LREAL#26.0;
   BenchUut6.windowSize := INT#100;
   BenchUut6.reset := FALSE;
   TraceIn_cyclicExecution[295] := BenchUut6.cyclicExecution;
   TraceIn_trigger[295] := BenchUut6.trigger;
   TraceIn_value[295] := BenchUut6.value;
   TraceIn_windowSize[295] := BenchUut6.windowSize;
   TraceIn_reset[295] := BenchUut6.reset;
   BenchUut6();
   TraceOut_average[295] := BenchUut6.average;
   TraceOut_windowSizeReached[295] := BenchUut6.windowSizeReached;
   TraceOut_error[295] := BenchUut6.error;
   TraceOut_status[295] := BenchUut6.status;
   BenchCalls := BenchCalls + 1;
 296:
   BenchUut6.cyclicExecution := FALSE;
   BenchUut6.trigger := TRUE;
   BenchUut6.value := LREAL#27.0;
   BenchUut6.windowSize := INT#100;
   BenchUut6.reset := FALSE;
   TraceIn_cyclicExecution[296] := BenchUut6.cyclicExecution;
   TraceIn_trigger[296] := BenchUut6.trigger;
   TraceIn_value[296] := BenchUut6.value;
   TraceIn_windowSize[296] := BenchUut6.windowSize;
   TraceIn_reset[296] := BenchUut6.reset;
   BenchUut6();
   TraceOut_average[296] := BenchUut6.average;
   TraceOut_windowSizeReached[296] := BenchUut6.windowSizeReached;
   TraceOut_error[296] := BenchUut6.error;
   TraceOut_status[296] := BenchUut6.status;
   BenchCalls := BenchCalls + 1;
 297:
   BenchUut6.cyclicExecution := FALSE;
   BenchUut6.trigger := FALSE;
   BenchUut6.value := LREAL#27.0;
   BenchUut6.windowSize := INT#100;
   BenchUut6.reset := FALSE;
   TraceIn_cyclicExecution[297] := BenchUut6.cyclicExecution;
   TraceIn_trigger[297] := BenchUut6.trigger;
   TraceIn_value[297] := BenchUut6.value;
   TraceIn_windowSize[297] := BenchUut6.windowSize;
   TraceIn_reset[297] := BenchUut6.reset;
   BenchUut6();
   TraceOut_average[297] := BenchUut6.average;
   TraceOut_windowSizeReached[297] := BenchUut6.windowSizeReached;
   TraceOut_error[297] := BenchUut6.error;
   TraceOut_status[297] := BenchUut6.status;
   BenchCalls := BenchCalls + 1;
 298:
   BenchUut6.cyclicExecution := FALSE;
   BenchUut6.trigger := TRUE;
   BenchUut6.value := LREAL#28.0;
   BenchUut6.windowSize := INT#100;
   BenchUut6.reset := FALSE;
   TraceIn_cyclicExecution[298] := BenchUut6.cyclicExecution;
   TraceIn_trigger[298] := BenchUut6.trigger;
   TraceIn_value[298] := BenchUut6.value;
   TraceIn_windowSize[298] := BenchUut6.windowSize;
   TraceIn_reset[298] := BenchUut6.reset;
   BenchUut6();
   TraceOut_average[298] := BenchUut6.average;
   TraceOut_windowSizeReached[298] := BenchUut6.windowSizeReached;
   TraceOut_error[298] := BenchUut6.error;
   TraceOut_status[298] := BenchUut6.status;
   BenchCalls := BenchCalls + 1;
 299:
   BenchUut6.cyclicExecution := FALSE;
   BenchUut6.trigger := FALSE;
   BenchUut6.value := LREAL#28.0;
   BenchUut6.windowSize := INT#100;
   BenchUut6.reset := FALSE;
   TraceIn_cyclicExecution[299] := BenchUut6.cyclicExecution;
   TraceIn_trigger[299] := BenchUut6.trigger;
   TraceIn_value[299] := BenchUut6.value;
   TraceIn_windowSize[299] := BenchUut6.windowSize;
   TraceIn_reset[299] := BenchUut6.reset;
   BenchUut6();
   TraceOut_average[299] := BenchUut6.average;
   TraceOut_windowSizeReached[299] := BenchUut6.windowSizeReached;
   TraceOut_error[299] := BenchUut6.error;
   TraceOut_status[299] := BenchUut6.status;
   BenchCalls := BenchCalls + 1;
 300:
   BenchUut6.cyclicExecution := FALSE;
   BenchUut6.trigger := TRUE;
   BenchUut6.value := LREAL#29.0;
   BenchUut6.windowSize := INT#100;
   BenchUut6.reset := FALSE;
   TraceIn_cyclicExecution[300] := BenchUut6.cyclicExecution;
   TraceIn_trigger[300] := BenchUut6.trigger;
   TraceIn_value[300] := BenchUut6.value;
   TraceIn_windowSize[300] := BenchUut6.windowSize;
   TraceIn_reset[300] := BenchUut6.reset;
   BenchUut6();
   TraceOut_average[300] := BenchUut6.average;
   TraceOut_windowSizeReached[300] := BenchUut6.windowSizeReached;
   TraceOut_error[300] := BenchUut6.error;
   TraceOut_status[300] := BenchUut6.status;
   BenchCalls := BenchCalls + 1;
 301:
   BenchUut6.cyclicExecution := FALSE;
   BenchUut6.trigger := FALSE;
   BenchUut6.value := LREAL#29.0;
   BenchUut6.windowSize := INT#100;
   BenchUut6.reset := FALSE;
   TraceIn_cyclicExecution[301] := BenchUut6.cyclicExecution;
   TraceIn_trigger[301] := BenchUut6.trigger;
   TraceIn_value[301] := BenchUut6.value;
   TraceIn_windowSize[301] := BenchUut6.windowSize;
   TraceIn_reset[301] := BenchUut6.reset;
   BenchUut6();
   TraceOut_average[301] := BenchUut6.average;
   TraceOut_windowSizeReached[301] := BenchUut6.windowSizeReached;
   TraceOut_error[301] := BenchUut6.error;
   TraceOut_status[301] := BenchUut6.status;
   BenchCalls := BenchCalls + 1;
 302:
   BenchUut6.cyclicExecution := FALSE;
   BenchUut6.trigger := TRUE;
   BenchUut6.value := LREAL#30.0;
   BenchUut6.windowSize := INT#100;
   BenchUut6.reset := FALSE;
   TraceIn_cyclicExecution[302] := BenchUut6.cyclicExecution;
   TraceIn_trigger[302] := BenchUut6.trigger;
   TraceIn_value[302] := BenchUut6.value;
   TraceIn_windowSize[302] := BenchUut6.windowSize;
   TraceIn_reset[302] := BenchUut6.reset;
   BenchUut6();
   TraceOut_average[302] := BenchUut6.average;
   TraceOut_windowSizeReached[302] := BenchUut6.windowSizeReached;
   TraceOut_error[302] := BenchUut6.error;
   TraceOut_status[302] := BenchUut6.status;
   BenchCalls := BenchCalls + 1;
 303:
   BenchUut6.cyclicExecution := FALSE;
   BenchUut6.trigger := FALSE;
   BenchUut6.value := LREAL#30.0;
   BenchUut6.windowSize := INT#100;
   BenchUut6.reset := FALSE;
   TraceIn_cyclicExecution[303] := BenchUut6.cyclicExecution;
   TraceIn_trigger[303] := BenchUut6.trigger;
   TraceIn_value[303] := BenchUut6.value;
   TraceIn_windowSize[303] := BenchUut6.windowSize;
   TraceIn_reset[303] := BenchUut6.reset;
   BenchUut6();
   TraceOut_average[303] := BenchUut6.average;
   TraceOut_windowSizeReached[303] := BenchUut6.windowSizeReached;
   TraceOut_error[303] := BenchUut6.error;
   TraceOut_status[303] := BenchUut6.status;
   BenchCalls := BenchCalls + 1;
 304:
   BenchUut6.cyclicExecution := FALSE;
   BenchUut6.trigger := TRUE;
   BenchUut6.value := LREAL#31.0;
   BenchUut6.windowSize := INT#100;
   BenchUut6.reset := FALSE;
   TraceIn_cyclicExecution[304] := BenchUut6.cyclicExecution;
   TraceIn_trigger[304] := BenchUut6.trigger;
   TraceIn_value[304] := BenchUut6.value;
   TraceIn_windowSize[304] := BenchUut6.windowSize;
   TraceIn_reset[304] := BenchUut6.reset;
   BenchUut6();
   TraceOut_average[304] := BenchUut6.average;
   TraceOut_windowSizeReached[304] := BenchUut6.windowSizeReached;
   TraceOut_error[304] := BenchUut6.error;
   TraceOut_status[304] := BenchUut6.status;
   BenchCalls := BenchCalls + 1;
 305:
   BenchUut6.cyclicExecution := FALSE;
   BenchUut6.trigger := FALSE;
   BenchUut6.value := LREAL#31.0;
   BenchUut6.windowSize := INT#100;
   BenchUut6.reset := FALSE;
   TraceIn_cyclicExecution[305] := BenchUut6.cyclicExecution;
   TraceIn_trigger[305] := BenchUut6.trigger;
   TraceIn_value[305] := BenchUut6.value;
   TraceIn_windowSize[305] := BenchUut6.windowSize;
   TraceIn_reset[305] := BenchUut6.reset;
   BenchUut6();
   TraceOut_average[305] := BenchUut6.average;
   TraceOut_windowSizeReached[305] := BenchUut6.windowSizeReached;
   TraceOut_error[305] := BenchUut6.error;
   TraceOut_status[305] := BenchUut6.status;
   BenchCalls := BenchCalls + 1;
 306:
   BenchUut6.cyclicExecution := FALSE;
   BenchUut6.trigger := TRUE;
   BenchUut6.value := LREAL#32.0;
   BenchUut6.windowSize := INT#100;
   BenchUut6.reset := FALSE;
   TraceIn_cyclicExecution[306] := BenchUut6.cyclicExecution;
   TraceIn_trigger[306] := BenchUut6.trigger;
   TraceIn_value[306] := BenchUut6.value;
   TraceIn_windowSize[306] := BenchUut6.windowSize;
   TraceIn_reset[306] := BenchUut6.reset;
   BenchUut6();
   TraceOut_average[306] := BenchUut6.average;
   TraceOut_windowSizeReached[306] := BenchUut6.windowSizeReached;
   TraceOut_error[306] := BenchUut6.error;
   TraceOut_status[306] := BenchUut6.status;
   BenchCalls := BenchCalls + 1;
 307:
   BenchUut6.cyclicExecution := FALSE;
   BenchUut6.trigger := FALSE;
   BenchUut6.value := LREAL#32.0;
   BenchUut6.windowSize := INT#100;
   BenchUut6.reset := FALSE;
   TraceIn_cyclicExecution[307] := BenchUut6.cyclicExecution;
   TraceIn_trigger[307] := BenchUut6.trigger;
   TraceIn_value[307] := BenchUut6.value;
   TraceIn_windowSize[307] := BenchUut6.windowSize;
   TraceIn_reset[307] := BenchUut6.reset;
   BenchUut6();
   TraceOut_average[307] := BenchUut6.average;
   TraceOut_windowSizeReached[307] := BenchUut6.windowSizeReached;
   TraceOut_error[307] := BenchUut6.error;
   TraceOut_status[307] := BenchUut6.status;
   BenchCalls := BenchCalls + 1;
 308:
   BenchUut6.cyclicExecution := FALSE;
   BenchUut6.trigger := TRUE;
   BenchUut6.value := LREAL#33.0;
   BenchUut6.windowSize := INT#100;
   BenchUut6.reset := FALSE;
   TraceIn_cyclicExecution[308] := BenchUut6.cyclicExecution;
   TraceIn_trigger[308] := BenchUut6.trigger;
   TraceIn_value[308] := BenchUut6.value;
   TraceIn_windowSize[308] := BenchUut6.windowSize;
   TraceIn_reset[308] := BenchUut6.reset;
   BenchUut6();
   TraceOut_average[308] := BenchUut6.average;
   TraceOut_windowSizeReached[308] := BenchUut6.windowSizeReached;
   TraceOut_error[308] := BenchUut6.error;
   TraceOut_status[308] := BenchUut6.status;
   BenchCalls := BenchCalls + 1;
 309:
   BenchUut6.cyclicExecution := FALSE;
   BenchUut6.trigger := FALSE;
   BenchUut6.value := LREAL#33.0;
   BenchUut6.windowSize := INT#100;
   BenchUut6.reset := FALSE;
   TraceIn_cyclicExecution[309] := BenchUut6.cyclicExecution;
   TraceIn_trigger[309] := BenchUut6.trigger;
   TraceIn_value[309] := BenchUut6.value;
   TraceIn_windowSize[309] := BenchUut6.windowSize;
   TraceIn_reset[309] := BenchUut6.reset;
   BenchUut6();
   TraceOut_average[309] := BenchUut6.average;
   TraceOut_windowSizeReached[309] := BenchUut6.windowSizeReached;
   TraceOut_error[309] := BenchUut6.error;
   TraceOut_status[309] := BenchUut6.status;
   BenchCalls := BenchCalls + 1;
 310:
   BenchUut6.cyclicExecution := FALSE;
   BenchUut6.trigger := TRUE;
   BenchUut6.value := LREAL#34.0;
   BenchUut6.windowSize := INT#100;
   BenchUut6.reset := FALSE;
   TraceIn_cyclicExecution[310] := BenchUut6.cyclicExecution;
   TraceIn_trigger[310] := BenchUut6.trigger;
   TraceIn_value[310] := BenchUut6.value;
   TraceIn_windowSize[310] := BenchUut6.windowSize;
   TraceIn_reset[310] := BenchUut6.reset;
   BenchUut6();
   TraceOut_average[310] := BenchUut6.average;
   TraceOut_windowSizeReached[310] := BenchUut6.windowSizeReached;
   TraceOut_error[310] := BenchUut6.error;
   TraceOut_status[310] := BenchUut6.status;
   BenchCalls := BenchCalls + 1;
 311:
   BenchUut6.cyclicExecution := FALSE;
   BenchUut6.trigger := FALSE;
   BenchUut6.value := LREAL#34.0;
   BenchUut6.windowSize := INT#100;
   BenchUut6.reset := FALSE;
   TraceIn_cyclicExecution[311] := BenchUut6.cyclicExecution;
   TraceIn_trigger[311] := BenchUut6.trigger;
   TraceIn_value[311] := BenchUut6.value;
   TraceIn_windowSize[311] := BenchUut6.windowSize;
   TraceIn_reset[311] := BenchUut6.reset;
   BenchUut6();
   TraceOut_average[311] := BenchUut6.average;
   TraceOut_windowSizeReached[311] := BenchUut6.windowSizeReached;
   TraceOut_error[311] := BenchUut6.error;
   TraceOut_status[311] := BenchUut6.status;
   BenchCalls := BenchCalls + 1;
 312:
   BenchUut6.cyclicExecution := FALSE;
   BenchUut6.trigger := TRUE;
   BenchUut6.value := LREAL#35.0;
   BenchUut6.windowSize := INT#100;
   BenchUut6.reset := FALSE;
   TraceIn_cyclicExecution[312] := BenchUut6.cyclicExecution;
   TraceIn_trigger[312] := BenchUut6.trigger;
   TraceIn_value[312] := BenchUut6.value;
   TraceIn_windowSize[312] := BenchUut6.windowSize;
   TraceIn_reset[312] := BenchUut6.reset;
   BenchUut6();
   TraceOut_average[312] := BenchUut6.average;
   TraceOut_windowSizeReached[312] := BenchUut6.windowSizeReached;
   TraceOut_error[312] := BenchUut6.error;
   TraceOut_status[312] := BenchUut6.status;
   BenchCalls := BenchCalls + 1;
 313:
   BenchUut6.cyclicExecution := FALSE;
   BenchUut6.trigger := FALSE;
   BenchUut6.value := LREAL#35.0;
   BenchUut6.windowSize := INT#100;
   BenchUut6.reset := FALSE;
   TraceIn_cyclicExecution[313] := BenchUut6.cyclicExecution;
   TraceIn_trigger[313] := BenchUut6.trigger;
   TraceIn_value[313] := BenchUut6.value;
   TraceIn_windowSize[313] := BenchUut6.windowSize;
   TraceIn_reset[313] := BenchUut6.reset;
   BenchUut6();
   TraceOut_average[313] := BenchUut6.average;
   TraceOut_windowSizeReached[313] := BenchUut6.windowSizeReached;
   TraceOut_error[313] := BenchUut6.error;
   TraceOut_status[313] := BenchUut6.status;
   BenchCalls := BenchCalls + 1;
 314:
   BenchUut6.cyclicExecution := FALSE;
   BenchUut6.trigger := TRUE;
   BenchUut6.value := LREAL#36.0;
   BenchUut6.windowSize := INT#100;
   BenchUut6.reset := FALSE;
   TraceIn_cyclicExecution[314] := BenchUut6.cyclicExecution;
   TraceIn_trigger[314] := BenchUut6.trigger;
   TraceIn_value[314] := BenchUut6.value;
   TraceIn_windowSize[314] := BenchUut6.windowSize;
   TraceIn_reset[314] := BenchUut6.reset;
   BenchUut6();
   TraceOut_average[314] := BenchUut6.average;
   TraceOut_windowSizeReached[314] := BenchUut6.windowSizeReached;
   TraceOut_error[314] := BenchUut6.error;
   TraceOut_status[314] := BenchUut6.status;
   BenchCalls := BenchCalls + 1;
 315:
   BenchUut6.cyclicExecution := FALSE;
   BenchUut6.trigger := FALSE;
   BenchUut6.value := LREAL#36.0;
   BenchUut6.windowSize := INT#100;
   BenchUut6.reset := FALSE;
   TraceIn_cyclicExecution[315] := BenchUut6.cyclicExecution;
   TraceIn_trigger[315] := BenchUut6.trigger;
   TraceIn_value[315] := BenchUut6.value;
   TraceIn_windowSize[315] := BenchUut6.windowSize;
   TraceIn_reset[315] := BenchUut6.reset;
   BenchUut6();
   TraceOut_average[315] := BenchUut6.average;
   TraceOut_windowSizeReached[315] := BenchUut6.windowSizeReached;
   TraceOut_error[315] := BenchUut6.error;
   TraceOut_status[315] := BenchUut6.status;
   BenchCalls := BenchCalls + 1;
 316:
   BenchUut6.cyclicExecution := FALSE;
   BenchUut6.trigger := TRUE;
   BenchUut6.value := LREAL#37.0;
   BenchUut6.windowSize := INT#100;
   BenchUut6.reset := FALSE;
   TraceIn_cyclicExecution[316] := BenchUut6.cyclicExecution;
   TraceIn_trigger[316] := BenchUut6.trigger;
   TraceIn_value[316] := BenchUut6.value;
   TraceIn_windowSize[316] := BenchUut6.windowSize;
   TraceIn_reset[316] := BenchUut6.reset;
   BenchUut6();
   TraceOut_average[316] := BenchUut6.average;
   TraceOut_windowSizeReached[316] := BenchUut6.windowSizeReached;
   TraceOut_error[316] := BenchUut6.error;
   TraceOut_status[316] := BenchUut6.status;
   BenchCalls := BenchCalls + 1;
 317:
   BenchUut6.cyclicExecution := FALSE;
   BenchUut6.trigger := FALSE;
   BenchUut6.value := LREAL#37.0;
   BenchUut6.windowSize := INT#100;
   BenchUut6.reset := FALSE;
   TraceIn_cyclicExecution[317] := BenchUut6.cyclicExecution;
   TraceIn_trigger[317] := BenchUut6.trigger;
   TraceIn_value[317] := BenchUut6.value;
   TraceIn_windowSize[317] := BenchUut6.windowSize;
   TraceIn_reset[317] := BenchUut6.reset;
   BenchUut6();
   TraceOut_average[317] := BenchUut6.average;
   TraceOut_windowSizeReached[317] := BenchUut6.windowSizeReached;
   TraceOut_error[317] := BenchUut6.error;
   TraceOut_status[317] := BenchUut6.status;
   BenchCalls := BenchCalls + 1;
 318:
   BenchUut6.cyclicExecution := FALSE;
   BenchUut6.trigger := TRUE;
   BenchUut6.value := LREAL#38.0;
   BenchUut6.windowSize := INT#100;
   BenchUut6.reset := FALSE;
   TraceIn_cyclicExecution[318] := BenchUut6.cyclicExecution;
   TraceIn_trigger[318] := BenchUut6.trigger;
   TraceIn_value[318] := BenchUut6.value;
   TraceIn_windowSize[318] := BenchUut6.windowSize;
   TraceIn_reset[318] := BenchUut6.reset;
   BenchUut6();
   TraceOut_average[318] := BenchUut6.average;
   TraceOut_windowSizeReached[318] := BenchUut6.windowSizeReached;
   TraceOut_error[318] := BenchUut6.error;
   TraceOut_status[318] := BenchUut6.status;
   BenchCalls := BenchCalls + 1;
 319:
   BenchUut6.cyclicExecution := FALSE;
   BenchUut6.trigger := FALSE;
   BenchUut6.value := LREAL#38.0;
   BenchUut6.windowSize := INT#100;
   BenchUut6.reset := FALSE;
   TraceIn_cyclicExecution[319] := BenchUut6.cyclicExecution;
   TraceIn_trigger[319] := BenchUut6.trigger;
   TraceIn_value[319] := BenchUut6.value;
   TraceIn_windowSize[319] := BenchUut6.windowSize;
   TraceIn_reset[319] := BenchUut6.reset;
   BenchUut6();
   TraceOut_average[319] := BenchUut6.average;
   TraceOut_windowSizeReached[319] := BenchUut6.windowSizeReached;
   TraceOut_error[319] := BenchUut6.error;
   TraceOut_status[319] := BenchUut6.status;
   BenchCalls := BenchCalls + 1;
 320:
   BenchUut6.cyclicExecution := FALSE;
   BenchUut6.trigger := TRUE;
   BenchUut6.value := LREAL#39.0;
   BenchUut6.windowSize := INT#100;
   BenchUut6.reset := FALSE;
   TraceIn_cyclicExecution[320] := BenchUut6.cyclicExecution;
   TraceIn_trigger[320] := BenchUut6.trigger;
   TraceIn_value[320] := BenchUut6.value;
   TraceIn_windowSize[320] := BenchUut6.windowSize;
   TraceIn_reset[320] := BenchUut6.reset;
   BenchUut6();
   TraceOut_average[320] := BenchUut6.average;
   TraceOut_windowSizeReached[320] := BenchUut6.windowSizeReached;
   TraceOut_error[320] := BenchUut6.error;
   TraceOut_status[320] := BenchUut6.status;
   BenchCalls := BenchCalls + 1;
 321:
   BenchUut6.cyclicExecution := FALSE;
   BenchUut6.trigger := FALSE;
   BenchUut6.value := LREAL#39.0;
   BenchUut6.windowSize := INT#100;
   BenchUut6.reset := FALSE;
   TraceIn_cyclicExecution[321] := BenchUut6.cyclicExecution;
   TraceIn_trigger[321] := BenchUut6.trigger;
   TraceIn_value[321] := BenchUut6.value;
   TraceIn_windowSize[321] := BenchUut6.windowSize;
   TraceIn_reset[321] := BenchUut6.reset;
   BenchUut6();
   TraceOut_average[321] := BenchUut6.average;
   TraceOut_windowSizeReached[321] := BenchUut6.windowSizeReached;
   TraceOut_error[321] := BenchUut6.error;
   TraceOut_status[321] := BenchUut6.status;
   BenchCalls := BenchCalls + 1;
 322:
   BenchUut6.cyclicExecution := FALSE;
   BenchUut6.trigger := TRUE;
   BenchUut6.value := LREAL#40.0;
   BenchUut6.windowSize := INT#100;
   BenchUut6.reset := FALSE;
   TraceIn_cyclicExecution[322] := BenchUut6.cyclicExecution;
   TraceIn_trigger[322] := BenchUut6.trigger;
   TraceIn_value[322] := BenchUut6.value;
   TraceIn_windowSize[322] := BenchUut6.windowSize;
   TraceIn_reset[322] := BenchUut6.reset;
   BenchUut6();
   TraceOut_average[322] := BenchUut6.average;
   TraceOut_windowSizeReached[322] := BenchUut6.windowSizeReached;
   TraceOut_error[322] := BenchUut6.error;
   TraceOut_status[322] := BenchUut6.status;
   BenchCalls := BenchCalls + 1;
 323:
   BenchUut6.cyclicExecution := FALSE;
   BenchUut6.trigger := FALSE;
   BenchUut6.value := LREAL#40.0;
   BenchUut6.windowSize := INT#100;
   BenchUut6.reset := FALSE;
   TraceIn_cyclicExecution[323] := BenchUut6.cyclicExecution;
   TraceIn_trigger[323] := BenchUut6.trigger;
   TraceIn_value[323] := BenchUut6.value;
   TraceIn_windowSize[323] := BenchUut6.windowSize;
   TraceIn_reset[323] := BenchUut6.reset;
   BenchUut6();
   TraceOut_average[323] := BenchUut6.average;
   TraceOut_windowSizeReached[323] := BenchUut6.windowSizeReached;
   TraceOut_error[323] := BenchUut6.error;
   TraceOut_status[323] := BenchUut6.status;
   BenchCalls := BenchCalls + 1;
 324:
   BenchUut6.cyclicExecution := FALSE;
   BenchUut6.trigger := TRUE;
   BenchUut6.value := LREAL#41.0;
   BenchUut6.windowSize := INT#100;
   BenchUut6.reset := FALSE;
   TraceIn_cyclicExecution[324] := BenchUut6.cyclicExecution;
   TraceIn_trigger[324] := BenchUut6.trigger;
   TraceIn_value[324] := BenchUut6.value;
   TraceIn_windowSize[324] := BenchUut6.windowSize;
   TraceIn_reset[324] := BenchUut6.reset;
   BenchUut6();
   TraceOut_average[324] := BenchUut6.average;
   TraceOut_windowSizeReached[324] := BenchUut6.windowSizeReached;
   TraceOut_error[324] := BenchUut6.error;
   TraceOut_status[324] := BenchUut6.status;
   BenchCalls := BenchCalls + 1;
 325:
   BenchUut6.cyclicExecution := FALSE;
   BenchUut6.trigger := FALSE;
   BenchUut6.value := LREAL#41.0;
   BenchUut6.windowSize := INT#100;
   BenchUut6.reset := FALSE;
   TraceIn_cyclicExecution[325] := BenchUut6.cyclicExecution;
   TraceIn_trigger[325] := BenchUut6.trigger;
   TraceIn_value[325] := BenchUut6.value;
   TraceIn_windowSize[325] := BenchUut6.windowSize;
   TraceIn_reset[325] := BenchUut6.reset;
   BenchUut6();
   TraceOut_average[325] := BenchUut6.average;
   TraceOut_windowSizeReached[325] := BenchUut6.windowSizeReached;
   TraceOut_error[325] := BenchUut6.error;
   TraceOut_status[325] := BenchUut6.status;
   BenchCalls := BenchCalls + 1;
 326:
   BenchUut6.cyclicExecution := FALSE;
   BenchUut6.trigger := TRUE;
   BenchUut6.value := LREAL#42.0;
   BenchUut6.windowSize := INT#100;
   BenchUut6.reset := FALSE;
   TraceIn_cyclicExecution[326] := BenchUut6.cyclicExecution;
   TraceIn_trigger[326] := BenchUut6.trigger;
   TraceIn_value[326] := BenchUut6.value;
   TraceIn_windowSize[326] := BenchUut6.windowSize;
   TraceIn_reset[326] := BenchUut6.reset;
   BenchUut6();
   TraceOut_average[326] := BenchUut6.average;
   TraceOut_windowSizeReached[326] := BenchUut6.windowSizeReached;
   TraceOut_error[326] := BenchUut6.error;
   TraceOut_status[326] := BenchUut6.status;
   BenchCalls := BenchCalls + 1;
 327:
   BenchUut6.cyclicExecution := FALSE;
   BenchUut6.trigger := FALSE;
   BenchUut6.value := LREAL#42.0;
   BenchUut6.windowSize := INT#100;
   BenchUut6.reset := FALSE;
   TraceIn_cyclicExecution[327] := BenchUut6.cyclicExecution;
   TraceIn_trigger[327] := BenchUut6.trigger;
   TraceIn_value[327] := BenchUut6.value;
   TraceIn_windowSize[327] := BenchUut6.windowSize;
   TraceIn_reset[327] := BenchUut6.reset;
   BenchUut6();
   TraceOut_average[327] := BenchUut6.average;
   TraceOut_windowSizeReached[327] := BenchUut6.windowSizeReached;
   TraceOut_error[327] := BenchUut6.error;
   TraceOut_status[327] := BenchUut6.status;
   BenchCalls := BenchCalls + 1;
 328:
   BenchUut6.cyclicExecution := FALSE;
   BenchUut6.trigger := TRUE;
   BenchUut6.value := LREAL#43.0;
   BenchUut6.windowSize := INT#100;
   BenchUut6.reset := FALSE;
   TraceIn_cyclicExecution[328] := BenchUut6.cyclicExecution;
   TraceIn_trigger[328] := BenchUut6.trigger;
   TraceIn_value[328] := BenchUut6.value;
   TraceIn_windowSize[328] := BenchUut6.windowSize;
   TraceIn_reset[328] := BenchUut6.reset;
   BenchUut6();
   TraceOut_average[328] := BenchUut6.average;
   TraceOut_windowSizeReached[328] := BenchUut6.windowSizeReached;
   TraceOut_error[328] := BenchUut6.error;
   TraceOut_status[328] := BenchUut6.status;
   BenchCalls := BenchCalls + 1;
 329:
   BenchUut6.cyclicExecution := FALSE;
   BenchUut6.trigger := FALSE;
   BenchUut6.value := LREAL#43.0;
   BenchUut6.windowSize := INT#100;
   BenchUut6.reset := FALSE;
   TraceIn_cyclicExecution[329] := BenchUut6.cyclicExecution;
   TraceIn_trigger[329] := BenchUut6.trigger;
   TraceIn_value[329] := BenchUut6.value;
   TraceIn_windowSize[329] := BenchUut6.windowSize;
   TraceIn_reset[329] := BenchUut6.reset;
   BenchUut6();
   TraceOut_average[329] := BenchUut6.average;
   TraceOut_windowSizeReached[329] := BenchUut6.windowSizeReached;
   TraceOut_error[329] := BenchUut6.error;
   TraceOut_status[329] := BenchUut6.status;
   BenchCalls := BenchCalls + 1;
 330:
   BenchUut6.cyclicExecution := FALSE;
   BenchUut6.trigger := TRUE;
   BenchUut6.value := LREAL#44.0;
   BenchUut6.windowSize := INT#100;
   BenchUut6.reset := FALSE;
   TraceIn_cyclicExecution[330] := BenchUut6.cyclicExecution;
   TraceIn_trigger[330] := BenchUut6.trigger;
   TraceIn_value[330] := BenchUut6.value;
   TraceIn_windowSize[330] := BenchUut6.windowSize;
   TraceIn_reset[330] := BenchUut6.reset;
   BenchUut6();
   TraceOut_average[330] := BenchUut6.average;
   TraceOut_windowSizeReached[330] := BenchUut6.windowSizeReached;
   TraceOut_error[330] := BenchUut6.error;
   TraceOut_status[330] := BenchUut6.status;
   BenchCalls := BenchCalls + 1;
 331:
   BenchUut6.cyclicExecution := FALSE;
   BenchUut6.trigger := FALSE;
   BenchUut6.value := LREAL#44.0;
   BenchUut6.windowSize := INT#100;
   BenchUut6.reset := FALSE;
   TraceIn_cyclicExecution[331] := BenchUut6.cyclicExecution;
   TraceIn_trigger[331] := BenchUut6.trigger;
   TraceIn_value[331] := BenchUut6.value;
   TraceIn_windowSize[331] := BenchUut6.windowSize;
   TraceIn_reset[331] := BenchUut6.reset;
   BenchUut6();
   TraceOut_average[331] := BenchUut6.average;
   TraceOut_windowSizeReached[331] := BenchUut6.windowSizeReached;
   TraceOut_error[331] := BenchUut6.error;
   TraceOut_status[331] := BenchUut6.status;
   BenchCalls := BenchCalls + 1;
 332:
   BenchUut6.cyclicExecution := FALSE;
   BenchUut6.trigger := TRUE;
   BenchUut6.value := LREAL#45.0;
   BenchUut6.windowSize := INT#100;
   BenchUut6.reset := FALSE;
   TraceIn_cyclicExecution[332] := BenchUut6.cyclicExecution;
   TraceIn_trigger[332] := BenchUut6.trigger;
   TraceIn_value[332] := BenchUut6.value;
   TraceIn_windowSize[332] := BenchUut6.windowSize;
   TraceIn_reset[332] := BenchUut6.reset;
   BenchUut6();
   TraceOut_average[332] := BenchUut6.average;
   TraceOut_windowSizeReached[332] := BenchUut6.windowSizeReached;
   TraceOut_error[332] := BenchUut6.error;
   TraceOut_status[332] := BenchUut6.status;
   BenchCalls := BenchCalls + 1;
 333:
   BenchUut6.cyclicExecution := FALSE;
   BenchUut6.trigger := FALSE;
   BenchUut6.value := LREAL#45.0;
   BenchUut6.windowSize := INT#100;
   BenchUut6.reset := FALSE;
   TraceIn_cyclicExecution[333] := BenchUut6.cyclicExecution;
   TraceIn_trigger[333] := BenchUut6.trigger;
   TraceIn_value[333] := BenchUut6.value;
   TraceIn_windowSize[333] := BenchUut6.windowSize;
   TraceIn_reset[333] := BenchUut6.reset;
   BenchUut6();
   TraceOut_average[333] := BenchUut6.average;
   TraceOut_windowSizeReached[333] := BenchUut6.windowSizeReached;
   TraceOut_error[333] := BenchUut6.error;
   TraceOut_status[333] := BenchUut6.status;
   BenchCalls := BenchCalls + 1;
 334:
   BenchUut6.cyclicExecution := FALSE;
   BenchUut6.trigger := TRUE;
   BenchUut6.value := LREAL#46.0;
   BenchUut6.windowSize := INT#100;
   BenchUut6.reset := FALSE;
   TraceIn_cyclicExecution[334] := BenchUut6.cyclicExecution;
   TraceIn_trigger[334] := BenchUut6.trigger;
   TraceIn_value[334] := BenchUut6.value;
   TraceIn_windowSize[334] := BenchUut6.windowSize;
   TraceIn_reset[334] := BenchUut6.reset;
   BenchUut6();
   TraceOut_average[334] := BenchUut6.average;
   TraceOut_windowSizeReached[334] := BenchUut6.windowSizeReached;
   TraceOut_error[334] := BenchUut6.error;
   TraceOut_status[334] := BenchUut6.status;
   BenchCalls := BenchCalls + 1;
 335:
   BenchUut6.cyclicExecution := FALSE;
   BenchUut6.trigger := FALSE;
   BenchUut6.value := LREAL#46.0;
   BenchUut6.windowSize := INT#100;
   BenchUut6.reset := FALSE;
   TraceIn_cyclicExecution[335] := BenchUut6.cyclicExecution;
   TraceIn_trigger[335] := BenchUut6.trigger;
   TraceIn_value[335] := BenchUut6.value;
   TraceIn_windowSize[335] := BenchUut6.windowSize;
   TraceIn_reset[335] := BenchUut6.reset;
   BenchUut6();
   TraceOut_average[335] := BenchUut6.average;
   TraceOut_windowSizeReached[335] := BenchUut6.windowSizeReached;
   TraceOut_error[335] := BenchUut6.error;
   TraceOut_status[335] := BenchUut6.status;
   BenchCalls := BenchCalls + 1;
 336:
   BenchUut6.cyclicExecution := FALSE;
   BenchUut6.trigger := TRUE;
   BenchUut6.value := LREAL#47.0;
   BenchUut6.windowSize := INT#100;
   BenchUut6.reset := FALSE;
   TraceIn_cyclicExecution[336] := BenchUut6.cyclicExecution;
   TraceIn_trigger[336] := BenchUut6.trigger;
   TraceIn_value[336] := BenchUut6.value;
   TraceIn_windowSize[336] := BenchUut6.windowSize;
   TraceIn_reset[336] := BenchUut6.reset;
   BenchUut6();
   TraceOut_average[336] := BenchUut6.average;
   TraceOut_windowSizeReached[336] := BenchUut6.windowSizeReached;
   TraceOut_error[336] := BenchUut6.error;
   TraceOut_status[336] := BenchUut6.status;
   BenchCalls := BenchCalls + 1;
 337:
   BenchUut6.cyclicExecution := FALSE;
   BenchUut6.trigger := FALSE;
   BenchUut6.value := LREAL#47.0;
   BenchUut6.windowSize := INT#100;
   BenchUut6.reset := FALSE;
   TraceIn_cyclicExecution[337] := BenchUut6.cyclicExecution;
   TraceIn_trigger[337] := BenchUut6.trigger;
   TraceIn_value[337] := BenchUut6.value;
   TraceIn_windowSize[337] := BenchUut6.windowSize;
   TraceIn_reset[337] := BenchUut6.reset;
   BenchUut6();
   TraceOut_average[337] := BenchUut6.average;
   TraceOut_windowSizeReached[337] := BenchUut6.windowSizeReached;
   TraceOut_error[337] := BenchUut6.error;
   TraceOut_status[337] := BenchUut6.status;
   BenchCalls := BenchCalls + 1;
 338:
   BenchUut6.cyclicExecution := FALSE;
   BenchUut6.trigger := TRUE;
   BenchUut6.value := LREAL#48.0;
   BenchUut6.windowSize := INT#100;
   BenchUut6.reset := FALSE;
   TraceIn_cyclicExecution[338] := BenchUut6.cyclicExecution;
   TraceIn_trigger[338] := BenchUut6.trigger;
   TraceIn_value[338] := BenchUut6.value;
   TraceIn_windowSize[338] := BenchUut6.windowSize;
   TraceIn_reset[338] := BenchUut6.reset;
   BenchUut6();
   TraceOut_average[338] := BenchUut6.average;
   TraceOut_windowSizeReached[338] := BenchUut6.windowSizeReached;
   TraceOut_error[338] := BenchUut6.error;
   TraceOut_status[338] := BenchUut6.status;
   BenchCalls := BenchCalls + 1;
 339:
   BenchUut6.cyclicExecution := FALSE;
   BenchUut6.trigger := FALSE;
   BenchUut6.value := LREAL#48.0;
   BenchUut6.windowSize := INT#100;
   BenchUut6.reset := FALSE;
   TraceIn_cyclicExecution[339] := BenchUut6.cyclicExecution;
   TraceIn_trigger[339] := BenchUut6.trigger;
   TraceIn_value[339] := BenchUut6.value;
   TraceIn_windowSize[339] := BenchUut6.windowSize;
   TraceIn_reset[339] := BenchUut6.reset;
   BenchUut6();
   TraceOut_average[339] := BenchUut6.average;
   TraceOut_windowSizeReached[339] := BenchUut6.windowSizeReached;
   TraceOut_error[339] := BenchUut6.error;
   TraceOut_status[339] := BenchUut6.status;
   BenchCalls := BenchCalls + 1;
 340:
   BenchUut6.cyclicExecution := FALSE;
   BenchUut6.trigger := TRUE;
   BenchUut6.value := LREAL#49.0;
   BenchUut6.windowSize := INT#100;
   BenchUut6.reset := FALSE;
   TraceIn_cyclicExecution[340] := BenchUut6.cyclicExecution;
   TraceIn_trigger[340] := BenchUut6.trigger;
   TraceIn_value[340] := BenchUut6.value;
   TraceIn_windowSize[340] := BenchUut6.windowSize;
   TraceIn_reset[340] := BenchUut6.reset;
   BenchUut6();
   TraceOut_average[340] := BenchUut6.average;
   TraceOut_windowSizeReached[340] := BenchUut6.windowSizeReached;
   TraceOut_error[340] := BenchUut6.error;
   TraceOut_status[340] := BenchUut6.status;
   BenchCalls := BenchCalls + 1;
 341:
   BenchUut6.cyclicExecution := FALSE;
   BenchUut6.trigger := FALSE;
   BenchUut6.value := LREAL#49.0;
   BenchUut6.windowSize := INT#100;
   BenchUut6.reset := FALSE;
   TraceIn_cyclicExecution[341] := BenchUut6.cyclicExecution;
   TraceIn_trigger[341] := BenchUut6.trigger;
   TraceIn_value[341] := BenchUut6.value;
   TraceIn_windowSize[341] := BenchUut6.windowSize;
   TraceIn_reset[341] := BenchUut6.reset;
   BenchUut6();
   TraceOut_average[341] := BenchUut6.average;
   TraceOut_windowSizeReached[341] := BenchUut6.windowSizeReached;
   TraceOut_error[341] := BenchUut6.error;
   TraceOut_status[341] := BenchUut6.status;
   BenchCalls := BenchCalls + 1;
 342:
   BenchUut6.cyclicExecution := FALSE;
   BenchUut6.trigger := TRUE;
   BenchUut6.value := LREAL#50.0;
   BenchUut6.windowSize := INT#100;
   BenchUut6.reset := FALSE;
   TraceIn_cyclicExecution[342] := BenchUut6.cyclicExecution;
   TraceIn_trigger[342] := BenchUut6.trigger;
   TraceIn_value[342] := BenchUut6.value;
   TraceIn_windowSize[342] := BenchUut6.windowSize;
   TraceIn_reset[342] := BenchUut6.reset;
   BenchUut6();
   TraceOut_average[342] := BenchUut6.average;
   TraceOut_windowSizeReached[342] := BenchUut6.windowSizeReached;
   TraceOut_error[342] := BenchUut6.error;
   TraceOut_status[342] := BenchUut6.status;
   BenchCalls := BenchCalls + 1;
 343:
   BenchUut6.cyclicExecution := FALSE;
   BenchUut6.trigger := FALSE;
   BenchUut6.value := LREAL#50.0;
   BenchUut6.windowSize := INT#100;
   BenchUut6.reset := FALSE;
   TraceIn_cyclicExecution[343] := BenchUut6.cyclicExecution;
   TraceIn_trigger[343] := BenchUut6.trigger;
   TraceIn_value[343] := BenchUut6.value;
   TraceIn_windowSize[343] := BenchUut6.windowSize;
   TraceIn_reset[343] := BenchUut6.reset;
   BenchUut6();
   TraceOut_average[343] := BenchUut6.average;
   TraceOut_windowSizeReached[343] := BenchUut6.windowSizeReached;
   TraceOut_error[343] := BenchUut6.error;
   TraceOut_status[343] := BenchUut6.status;
   BenchCalls := BenchCalls + 1;
 344:
   BenchUut6.cyclicExecution := FALSE;
   BenchUut6.trigger := TRUE;
   BenchUut6.value := LREAL#51.0;
   BenchUut6.windowSize := INT#100;
   BenchUut6.reset := FALSE;
   TraceIn_cyclicExecution[344] := BenchUut6.cyclicExecution;
   TraceIn_trigger[344] := BenchUut6.trigger;
   TraceIn_value[344] := BenchUut6.value;
   TraceIn_windowSize[344] := BenchUut6.windowSize;
   TraceIn_reset[344] := BenchUut6.reset;
   BenchUut6();
   TraceOut_average[344] := BenchUut6.average;
   TraceOut_windowSizeReached[344] := BenchUut6.windowSizeReached;
   TraceOut_error[344] := BenchUut6.error;
   TraceOut_status[344] := BenchUut6.status;
   BenchCalls := BenchCalls + 1;
 345:
   BenchUut6.cyclicExecution := FALSE;
   BenchUut6.trigger := FALSE;
   BenchUut6.value := LREAL#51.0;
   BenchUut6.windowSize := INT#100;
   BenchUut6.reset := FALSE;
   TraceIn_cyclicExecution[345] := BenchUut6.cyclicExecution;
   TraceIn_trigger[345] := BenchUut6.trigger;
   TraceIn_value[345] := BenchUut6.value;
   TraceIn_windowSize[345] := BenchUut6.windowSize;
   TraceIn_reset[345] := BenchUut6.reset;
   BenchUut6();
   TraceOut_average[345] := BenchUut6.average;
   TraceOut_windowSizeReached[345] := BenchUut6.windowSizeReached;
   TraceOut_error[345] := BenchUut6.error;
   TraceOut_status[345] := BenchUut6.status;
   BenchCalls := BenchCalls + 1;
 346:
   BenchUut6.cyclicExecution := FALSE;
   BenchUut6.trigger := TRUE;
   BenchUut6.value := LREAL#52.0;
   BenchUut6.windowSize := INT#100;
   BenchUut6.reset := FALSE;
   TraceIn_cyclicExecution[346] := BenchUut6.cyclicExecution;
   TraceIn_trigger[346] := BenchUut6.trigger;
   TraceIn_value[346] := BenchUut6.value;
   TraceIn_windowSize[346] := BenchUut6.windowSize;
   TraceIn_reset[346] := BenchUut6.reset;
   BenchUut6();
   TraceOut_average[346] := BenchUut6.average;
   TraceOut_windowSizeReached[346] := BenchUut6.windowSizeReached;
   TraceOut_error[346] := BenchUut6.error;
   TraceOut_status[346] := BenchUut6.status;
   BenchCalls := BenchCalls + 1;
 347:
   BenchUut6.cyclicExecution := FALSE;
   BenchUut6.trigger := FALSE;
   BenchUut6.value := LREAL#52.0;
   BenchUut6.windowSize := INT#100;
   BenchUut6.reset := FALSE;
   TraceIn_cyclicExecution[347] := BenchUut6.cyclicExecution;
   TraceIn_trigger[347] := BenchUut6.trigger;
   TraceIn_value[347] := BenchUut6.value;
   TraceIn_windowSize[347] := BenchUut6.windowSize;
   TraceIn_reset[347] := BenchUut6.reset;
   BenchUut6();
   TraceOut_average[347] := BenchUut6.average;
   TraceOut_windowSizeReached[347] := BenchUut6.windowSizeReached;
   TraceOut_error[347] := BenchUut6.error;
   TraceOut_status[347] := BenchUut6.status;
   BenchCalls := BenchCalls + 1;
 348:
   BenchUut6.cyclicExecution := FALSE;
   BenchUut6.trigger := TRUE;
   BenchUut6.value := LREAL#53.0;
   BenchUut6.windowSize := INT#100;
   BenchUut6.reset := FALSE;
   TraceIn_cyclicExecution[348] := BenchUut6.cyclicExecution;
   TraceIn_trigger[348] := BenchUut6.trigger;
   TraceIn_value[348] := BenchUut6.value;
   TraceIn_windowSize[348] := BenchUut6.windowSize;
   TraceIn_reset[348] := BenchUut6.reset;
   BenchUut6();
   TraceOut_average[348] := BenchUut6.average;
   TraceOut_windowSizeReached[348] := BenchUut6.windowSizeReached;
   TraceOut_error[348] := BenchUut6.error;
   TraceOut_status[348] := BenchUut6.status;
   BenchCalls := BenchCalls + 1;
 349:
   BenchUut6.cyclicExecution := FALSE;
   BenchUut6.trigger := FALSE;
   BenchUut6.value := LREAL#53.0;
   BenchUut6.windowSize := INT#100;
   BenchUut6.reset := FALSE;
   TraceIn_cyclicExecution[349] := BenchUut6.cyclicExecution;
   TraceIn_trigger[349] := BenchUut6.trigger;
   TraceIn_value[349] := BenchUut6.value;
   TraceIn_windowSize[349] := BenchUut6.windowSize;
   TraceIn_reset[349] := BenchUut6.reset;
   BenchUut6();
   TraceOut_average[349] := BenchUut6.average;
   TraceOut_windowSizeReached[349] := BenchUut6.windowSizeReached;
   TraceOut_error[349] := BenchUut6.error;
   TraceOut_status[349] := BenchUut6.status;
   BenchCalls := BenchCalls + 1;
 350:
   BenchUut6.cyclicExecution := FALSE;
   BenchUut6.trigger := TRUE;
   BenchUut6.value := LREAL#54.0;
   BenchUut6.windowSize := INT#100;
   BenchUut6.reset := FALSE;
   TraceIn_cyclicExecution[350] := BenchUut6.cyclicExecution;
   TraceIn_trigger[350] := BenchUut6.trigger;
   TraceIn_value[350] := BenchUut6.value;
   TraceIn_windowSize[350] := BenchUut6.windowSize;
   TraceIn_reset[350] := BenchUut6.reset;
   BenchUut6();
   TraceOut_average[350] := BenchUut6.average;
   TraceOut_windowSizeReached[350] := BenchUut6.windowSizeReached;
   TraceOut_error[350] := BenchUut6.error;
   TraceOut_status[350] := BenchUut6.status;
   BenchCalls := BenchCalls + 1;
 351:
   BenchUut6.cyclicExecution := FALSE;
   BenchUut6.trigger := FALSE;
   BenchUut6.value := LREAL#54.0;
   BenchUut6.windowSize := INT#100;
   BenchUut6.reset := FALSE;
   TraceIn_cyclicExecution[351] := BenchUut6.cyclicExecution;
   TraceIn_trigger[351] := BenchUut6.trigger;
   TraceIn_value[351] := BenchUut6.value;
   TraceIn_windowSize[351] := BenchUut6.windowSize;
   TraceIn_reset[351] := BenchUut6.reset;
   BenchUut6();
   TraceOut_average[351] := BenchUut6.average;
   TraceOut_windowSizeReached[351] := BenchUut6.windowSizeReached;
   TraceOut_error[351] := BenchUut6.error;
   TraceOut_status[351] := BenchUut6.status;
   BenchCalls := BenchCalls + 1;
 352:
   BenchUut6.cyclicExecution := FALSE;
   BenchUut6.trigger := TRUE;
   BenchUut6.value := LREAL#55.0;
   BenchUut6.windowSize := INT#100;
   BenchUut6.reset := FALSE;
   TraceIn_cyclicExecution[352] := BenchUut6.cyclicExecution;
   TraceIn_trigger[352] := BenchUut6.trigger;
   TraceIn_value[352] := BenchUut6.value;
   TraceIn_windowSize[352] := BenchUut6.windowSize;
   TraceIn_reset[352] := BenchUut6.reset;
   BenchUut6();
   TraceOut_average[352] := BenchUut6.average;
   TraceOut_windowSizeReached[352] := BenchUut6.windowSizeReached;
   TraceOut_error[352] := BenchUut6.error;
   TraceOut_status[352] := BenchUut6.status;
   BenchCalls := BenchCalls + 1;
 353:
   BenchUut6.cyclicExecution := FALSE;
   BenchUut6.trigger := FALSE;
   BenchUut6.value := LREAL#55.0;
   BenchUut6.windowSize := INT#100;
   BenchUut6.reset := FALSE;
   TraceIn_cyclicExecution[353] := BenchUut6.cyclicExecution;
   TraceIn_trigger[353] := BenchUut6.trigger;
   TraceIn_value[353] := BenchUut6.value;
   TraceIn_windowSize[353] := BenchUut6.windowSize;
   TraceIn_reset[353] := BenchUut6.reset;
   BenchUut6();
   TraceOut_average[353] := BenchUut6.average;
   TraceOut_windowSizeReached[353] := BenchUut6.windowSizeReached;
   TraceOut_error[353] := BenchUut6.error;
   TraceOut_status[353] := BenchUut6.status;
   BenchCalls := BenchCalls + 1;
 354:
   BenchUut6.cyclicExecution := FALSE;
   BenchUut6.trigger := TRUE;
   BenchUut6.value := LREAL#56.0;
   BenchUut6.windowSize := INT#100;
   BenchUut6.reset := FALSE;
   TraceIn_cyclicExecution[354] := BenchUut6.cyclicExecution;
   TraceIn_trigger[354] := BenchUut6.trigger;
   TraceIn_value[354] := BenchUut6.value;
   TraceIn_windowSize[354] := BenchUut6.windowSize;
   TraceIn_reset[354] := BenchUut6.reset;
   BenchUut6();
   TraceOut_average[354] := BenchUut6.average;
   TraceOut_windowSizeReached[354] := BenchUut6.windowSizeReached;
   TraceOut_error[354] := BenchUut6.error;
   TraceOut_status[354] := BenchUut6.status;
   BenchCalls := BenchCalls + 1;
 355:
   BenchUut6.cyclicExecution := FALSE;
   BenchUut6.trigger := FALSE;
   BenchUut6.value := LREAL#56.0;
   BenchUut6.windowSize := INT#100;
   BenchUut6.reset := FALSE;
   TraceIn_cyclicExecution[355] := BenchUut6.cyclicExecution;
   TraceIn_trigger[355] := BenchUut6.trigger;
   TraceIn_value[355] := BenchUut6.value;
   TraceIn_windowSize[355] := BenchUut6.windowSize;
   TraceIn_reset[355] := BenchUut6.reset;
   BenchUut6();
   TraceOut_average[355] := BenchUut6.average;
   TraceOut_windowSizeReached[355] := BenchUut6.windowSizeReached;
   TraceOut_error[355] := BenchUut6.error;
   TraceOut_status[355] := BenchUut6.status;
   BenchCalls := BenchCalls + 1;
 356:
   BenchUut6.cyclicExecution := FALSE;
   BenchUut6.trigger := TRUE;
   BenchUut6.value := LREAL#57.0;
   BenchUut6.windowSize := INT#100;
   BenchUut6.reset := FALSE;
   TraceIn_cyclicExecution[356] := BenchUut6.cyclicExecution;
   TraceIn_trigger[356] := BenchUut6.trigger;
   TraceIn_value[356] := BenchUut6.value;
   TraceIn_windowSize[356] := BenchUut6.windowSize;
   TraceIn_reset[356] := BenchUut6.reset;
   BenchUut6();
   TraceOut_average[356] := BenchUut6.average;
   TraceOut_windowSizeReached[356] := BenchUut6.windowSizeReached;
   TraceOut_error[356] := BenchUut6.error;
   TraceOut_status[356] := BenchUut6.status;
   BenchCalls := BenchCalls + 1;
 357:
   BenchUut6.cyclicExecution := FALSE;
   BenchUut6.trigger := FALSE;
   BenchUut6.value := LREAL#57.0;
   BenchUut6.windowSize := INT#100;
   BenchUut6.reset := FALSE;
   TraceIn_cyclicExecution[357] := BenchUut6.cyclicExecution;
   TraceIn_trigger[357] := BenchUut6.trigger;
   TraceIn_value[357] := BenchUut6.value;
   TraceIn_windowSize[357] := BenchUut6.windowSize;
   TraceIn_reset[357] := BenchUut6.reset;
   BenchUut6();
   TraceOut_average[357] := BenchUut6.average;
   TraceOut_windowSizeReached[357] := BenchUut6.windowSizeReached;
   TraceOut_error[357] := BenchUut6.error;
   TraceOut_status[357] := BenchUut6.status;
   BenchCalls := BenchCalls + 1;
 358:
   BenchUut6.cyclicExecution := FALSE;
   BenchUut6.trigger := TRUE;
   BenchUut6.value := LREAL#58.0;
   BenchUut6.windowSize := INT#100;
   BenchUut6.reset := FALSE;
   TraceIn_cyclicExecution[358] := BenchUut6.cyclicExecution;
   TraceIn_trigger[358] := BenchUut6.trigger;
   TraceIn_value[358] := BenchUut6.value;
   TraceIn_windowSize[358] := BenchUut6.windowSize;
   TraceIn_reset[358] := BenchUut6.reset;
   BenchUut6();
   TraceOut_average[358] := BenchUut6.average;
   TraceOut_windowSizeReached[358] := BenchUut6.windowSizeReached;
   TraceOut_error[358] := BenchUut6.error;
   TraceOut_status[358] := BenchUut6.status;
   BenchCalls := BenchCalls + 1;
 359:
   BenchUut6.cyclicExecution := FALSE;
   BenchUut6.trigger := FALSE;
   BenchUut6.value := LREAL#58.0;
   BenchUut6.windowSize := INT#100;
   BenchUut6.reset := FALSE;
   TraceIn_cyclicExecution[359] := BenchUut6.cyclicExecution;
   TraceIn_trigger[359] := BenchUut6.trigger;
   TraceIn_value[359] := BenchUut6.value;
   TraceIn_windowSize[359] := BenchUut6.windowSize;
   TraceIn_reset[359] := BenchUut6.reset;
   BenchUut6();
   TraceOut_average[359] := BenchUut6.average;
   TraceOut_windowSizeReached[359] := BenchUut6.windowSizeReached;
   TraceOut_error[359] := BenchUut6.error;
   TraceOut_status[359] := BenchUut6.status;
   BenchCalls := BenchCalls + 1;
 360:
   BenchUut6.cyclicExecution := FALSE;
   BenchUut6.trigger := TRUE;
   BenchUut6.value := LREAL#59.0;
   BenchUut6.windowSize := INT#100;
   BenchUut6.reset := FALSE;
   TraceIn_cyclicExecution[360] := BenchUut6.cyclicExecution;
   TraceIn_trigger[360] := BenchUut6.trigger;
   TraceIn_value[360] := BenchUut6.value;
   TraceIn_windowSize[360] := BenchUut6.windowSize;
   TraceIn_reset[360] := BenchUut6.reset;
   BenchUut6();
   TraceOut_average[360] := BenchUut6.average;
   TraceOut_windowSizeReached[360] := BenchUut6.windowSizeReached;
   TraceOut_error[360] := BenchUut6.error;
   TraceOut_status[360] := BenchUut6.status;
   BenchCalls := BenchCalls + 1;
 361:
   BenchUut6.cyclicExecution := FALSE;
   BenchUut6.trigger := FALSE;
   BenchUut6.value := LREAL#59.0;
   BenchUut6.windowSize := INT#100;
   BenchUut6.reset := FALSE;
   TraceIn_cyclicExecution[361] := BenchUut6.cyclicExecution;
   TraceIn_trigger[361] := BenchUut6.trigger;
   TraceIn_value[361] := BenchUut6.value;
   TraceIn_windowSize[361] := BenchUut6.windowSize;
   TraceIn_reset[361] := BenchUut6.reset;
   BenchUut6();
   TraceOut_average[361] := BenchUut6.average;
   TraceOut_windowSizeReached[361] := BenchUut6.windowSizeReached;
   TraceOut_error[361] := BenchUut6.error;
   TraceOut_status[361] := BenchUut6.status;
   BenchCalls := BenchCalls + 1;
 362:
   BenchUut6.cyclicExecution := FALSE;
   BenchUut6.trigger := TRUE;
   BenchUut6.value := LREAL#60.0;
   BenchUut6.windowSize := INT#100;
   BenchUut6.reset := FALSE;
   TraceIn_cyclicExecution[362] := BenchUut6.cyclicExecution;
   TraceIn_trigger[362] := BenchUut6.trigger;
   TraceIn_value[362] := BenchUut6.value;
   TraceIn_windowSize[362] := BenchUut6.windowSize;
   TraceIn_reset[362] := BenchUut6.reset;
   BenchUut6();
   TraceOut_average[362] := BenchUut6.average;
   TraceOut_windowSizeReached[362] := BenchUut6.windowSizeReached;
   TraceOut_error[362] := BenchUut6.error;
   TraceOut_status[362] := BenchUut6.status;
   BenchCalls := BenchCalls + 1;
 363:
   BenchUut6.cyclicExecution := FALSE;
   BenchUut6.trigger := FALSE;
   BenchUut6.value := LREAL#60.0;
   BenchUut6.windowSize := INT#100;
   BenchUut6.reset := FALSE;
   TraceIn_cyclicExecution[363] := BenchUut6.cyclicExecution;
   TraceIn_trigger[363] := BenchUut6.trigger;
   TraceIn_value[363] := BenchUut6.value;
   TraceIn_windowSize[363] := BenchUut6.windowSize;
   TraceIn_reset[363] := BenchUut6.reset;
   BenchUut6();
   TraceOut_average[363] := BenchUut6.average;
   TraceOut_windowSizeReached[363] := BenchUut6.windowSizeReached;
   TraceOut_error[363] := BenchUut6.error;
   TraceOut_status[363] := BenchUut6.status;
   BenchCalls := BenchCalls + 1;
 364:
   BenchUut6.cyclicExecution := FALSE;
   BenchUut6.trigger := TRUE;
   BenchUut6.value := LREAL#61.0;
   BenchUut6.windowSize := INT#100;
   BenchUut6.reset := FALSE;
   TraceIn_cyclicExecution[364] := BenchUut6.cyclicExecution;
   TraceIn_trigger[364] := BenchUut6.trigger;
   TraceIn_value[364] := BenchUut6.value;
   TraceIn_windowSize[364] := BenchUut6.windowSize;
   TraceIn_reset[364] := BenchUut6.reset;
   BenchUut6();
   TraceOut_average[364] := BenchUut6.average;
   TraceOut_windowSizeReached[364] := BenchUut6.windowSizeReached;
   TraceOut_error[364] := BenchUut6.error;
   TraceOut_status[364] := BenchUut6.status;
   BenchCalls := BenchCalls + 1;
 365:
   BenchUut6.cyclicExecution := FALSE;
   BenchUut6.trigger := FALSE;
   BenchUut6.value := LREAL#61.0;
   BenchUut6.windowSize := INT#100;
   BenchUut6.reset := FALSE;
   TraceIn_cyclicExecution[365] := BenchUut6.cyclicExecution;
   TraceIn_trigger[365] := BenchUut6.trigger;
   TraceIn_value[365] := BenchUut6.value;
   TraceIn_windowSize[365] := BenchUut6.windowSize;
   TraceIn_reset[365] := BenchUut6.reset;
   BenchUut6();
   TraceOut_average[365] := BenchUut6.average;
   TraceOut_windowSizeReached[365] := BenchUut6.windowSizeReached;
   TraceOut_error[365] := BenchUut6.error;
   TraceOut_status[365] := BenchUut6.status;
   BenchCalls := BenchCalls + 1;
 366:
   BenchUut6.cyclicExecution := FALSE;
   BenchUut6.trigger := TRUE;
   BenchUut6.value := LREAL#62.0;
   BenchUut6.windowSize := INT#100;
   BenchUut6.reset := FALSE;
   TraceIn_cyclicExecution[366] := BenchUut6.cyclicExecution;
   TraceIn_trigger[366] := BenchUut6.trigger;
   TraceIn_value[366] := BenchUut6.value;
   TraceIn_windowSize[366] := BenchUut6.windowSize;
   TraceIn_reset[366] := BenchUut6.reset;
   BenchUut6();
   TraceOut_average[366] := BenchUut6.average;
   TraceOut_windowSizeReached[366] := BenchUut6.windowSizeReached;
   TraceOut_error[366] := BenchUut6.error;
   TraceOut_status[366] := BenchUut6.status;
   BenchCalls := BenchCalls + 1;
 367:
   BenchUut6.cyclicExecution := FALSE;
   BenchUut6.trigger := FALSE;
   BenchUut6.value := LREAL#62.0;
   BenchUut6.windowSize := INT#100;
   BenchUut6.reset := FALSE;
   TraceIn_cyclicExecution[367] := BenchUut6.cyclicExecution;
   TraceIn_trigger[367] := BenchUut6.trigger;
   TraceIn_value[367] := BenchUut6.value;
   TraceIn_windowSize[367] := BenchUut6.windowSize;
   TraceIn_reset[367] := BenchUut6.reset;
   BenchUut6();
   TraceOut_average[367] := BenchUut6.average;
   TraceOut_windowSizeReached[367] := BenchUut6.windowSizeReached;
   TraceOut_error[367] := BenchUut6.error;
   TraceOut_status[367] := BenchUut6.status;
   BenchCalls := BenchCalls + 1;
 368:
   BenchUut6.cyclicExecution := FALSE;
   BenchUut6.trigger := TRUE;
   BenchUut6.value := LREAL#63.0;
   BenchUut6.windowSize := INT#100;
   BenchUut6.reset := FALSE;
   TraceIn_cyclicExecution[368] := BenchUut6.cyclicExecution;
   TraceIn_trigger[368] := BenchUut6.trigger;
   TraceIn_value[368] := BenchUut6.value;
   TraceIn_windowSize[368] := BenchUut6.windowSize;
   TraceIn_reset[368] := BenchUut6.reset;
   BenchUut6();
   TraceOut_average[368] := BenchUut6.average;
   TraceOut_windowSizeReached[368] := BenchUut6.windowSizeReached;
   TraceOut_error[368] := BenchUut6.error;
   TraceOut_status[368] := BenchUut6.status;
   BenchCalls := BenchCalls + 1;
 369:
   BenchUut6.cyclicExecution := FALSE;
   BenchUut6.trigger := FALSE;
   BenchUut6.value := LREAL#63.0;
   BenchUut6.windowSize := INT#100;
   BenchUut6.reset := FALSE;
   TraceIn_cyclicExecution[369] := BenchUut6.cyclicExecution;
   TraceIn_trigger[369] := BenchUut6.trigger;
   TraceIn_value[369] := BenchUut6.value;
   TraceIn_windowSize[369] := BenchUut6.windowSize;
   TraceIn_reset[369] := BenchUut6.reset;
   BenchUut6();
   TraceOut_average[369] := BenchUut6.average;
   TraceOut_windowSizeReached[369] := BenchUut6.windowSizeReached;
   TraceOut_error[369] := BenchUut6.error;
   TraceOut_status[369] := BenchUut6.status;
   BenchCalls := BenchCalls + 1;
 370:
   BenchUut6.cyclicExecution := FALSE;
   BenchUut6.trigger := TRUE;
   BenchUut6.value := LREAL#64.0;
   BenchUut6.windowSize := INT#100;
   BenchUut6.reset := FALSE;
   TraceIn_cyclicExecution[370] := BenchUut6.cyclicExecution;
   TraceIn_trigger[370] := BenchUut6.trigger;
   TraceIn_value[370] := BenchUut6.value;
   TraceIn_windowSize[370] := BenchUut6.windowSize;
   TraceIn_reset[370] := BenchUut6.reset;
   BenchUut6();
   TraceOut_average[370] := BenchUut6.average;
   TraceOut_windowSizeReached[370] := BenchUut6.windowSizeReached;
   TraceOut_error[370] := BenchUut6.error;
   TraceOut_status[370] := BenchUut6.status;
   BenchCalls := BenchCalls + 1;
 371:
   BenchUut6.cyclicExecution := FALSE;
   BenchUut6.trigger := FALSE;
   BenchUut6.value := LREAL#64.0;
   BenchUut6.windowSize := INT#100;
   BenchUut6.reset := FALSE;
   TraceIn_cyclicExecution[371] := BenchUut6.cyclicExecution;
   TraceIn_trigger[371] := BenchUut6.trigger;
   TraceIn_value[371] := BenchUut6.value;
   TraceIn_windowSize[371] := BenchUut6.windowSize;
   TraceIn_reset[371] := BenchUut6.reset;
   BenchUut6();
   TraceOut_average[371] := BenchUut6.average;
   TraceOut_windowSizeReached[371] := BenchUut6.windowSizeReached;
   TraceOut_error[371] := BenchUut6.error;
   TraceOut_status[371] := BenchUut6.status;
   BenchCalls := BenchCalls + 1;
 372:
   BenchUut6.cyclicExecution := FALSE;
   BenchUut6.trigger := TRUE;
   BenchUut6.value := LREAL#65.0;
   BenchUut6.windowSize := INT#100;
   BenchUut6.reset := FALSE;
   TraceIn_cyclicExecution[372] := BenchUut6.cyclicExecution;
   TraceIn_trigger[372] := BenchUut6.trigger;
   TraceIn_value[372] := BenchUut6.value;
   TraceIn_windowSize[372] := BenchUut6.windowSize;
   TraceIn_reset[372] := BenchUut6.reset;
   BenchUut6();
   TraceOut_average[372] := BenchUut6.average;
   TraceOut_windowSizeReached[372] := BenchUut6.windowSizeReached;
   TraceOut_error[372] := BenchUut6.error;
   TraceOut_status[372] := BenchUut6.status;
   BenchCalls := BenchCalls + 1;
 373:
   BenchUut6.cyclicExecution := FALSE;
   BenchUut6.trigger := FALSE;
   BenchUut6.value := LREAL#65.0;
   BenchUut6.windowSize := INT#100;
   BenchUut6.reset := FALSE;
   TraceIn_cyclicExecution[373] := BenchUut6.cyclicExecution;
   TraceIn_trigger[373] := BenchUut6.trigger;
   TraceIn_value[373] := BenchUut6.value;
   TraceIn_windowSize[373] := BenchUut6.windowSize;
   TraceIn_reset[373] := BenchUut6.reset;
   BenchUut6();
   TraceOut_average[373] := BenchUut6.average;
   TraceOut_windowSizeReached[373] := BenchUut6.windowSizeReached;
   TraceOut_error[373] := BenchUut6.error;
   TraceOut_status[373] := BenchUut6.status;
   BenchCalls := BenchCalls + 1;
 374:
   BenchUut6.cyclicExecution := FALSE;
   BenchUut6.trigger := TRUE;
   BenchUut6.value := LREAL#66.0;
   BenchUut6.windowSize := INT#100;
   BenchUut6.reset := FALSE;
   TraceIn_cyclicExecution[374] := BenchUut6.cyclicExecution;
   TraceIn_trigger[374] := BenchUut6.trigger;
   TraceIn_value[374] := BenchUut6.value;
   TraceIn_windowSize[374] := BenchUut6.windowSize;
   TraceIn_reset[374] := BenchUut6.reset;
   BenchUut6();
   TraceOut_average[374] := BenchUut6.average;
   TraceOut_windowSizeReached[374] := BenchUut6.windowSizeReached;
   TraceOut_error[374] := BenchUut6.error;
   TraceOut_status[374] := BenchUut6.status;
   BenchCalls := BenchCalls + 1;
 375:
   BenchUut6.cyclicExecution := FALSE;
   BenchUut6.trigger := FALSE;
   BenchUut6.value := LREAL#66.0;
   BenchUut6.windowSize := INT#100;
   BenchUut6.reset := FALSE;
   TraceIn_cyclicExecution[375] := BenchUut6.cyclicExecution;
   TraceIn_trigger[375] := BenchUut6.trigger;
   TraceIn_value[375] := BenchUut6.value;
   TraceIn_windowSize[375] := BenchUut6.windowSize;
   TraceIn_reset[375] := BenchUut6.reset;
   BenchUut6();
   TraceOut_average[375] := BenchUut6.average;
   TraceOut_windowSizeReached[375] := BenchUut6.windowSizeReached;
   TraceOut_error[375] := BenchUut6.error;
   TraceOut_status[375] := BenchUut6.status;
   BenchCalls := BenchCalls + 1;
 376:
   BenchUut6.cyclicExecution := FALSE;
   BenchUut6.trigger := TRUE;
   BenchUut6.value := LREAL#67.0;
   BenchUut6.windowSize := INT#100;
   BenchUut6.reset := FALSE;
   TraceIn_cyclicExecution[376] := BenchUut6.cyclicExecution;
   TraceIn_trigger[376] := BenchUut6.trigger;
   TraceIn_value[376] := BenchUut6.value;
   TraceIn_windowSize[376] := BenchUut6.windowSize;
   TraceIn_reset[376] := BenchUut6.reset;
   BenchUut6();
   TraceOut_average[376] := BenchUut6.average;
   TraceOut_windowSizeReached[376] := BenchUut6.windowSizeReached;
   TraceOut_error[376] := BenchUut6.error;
   TraceOut_status[376] := BenchUut6.status;
   BenchCalls := BenchCalls + 1;
 377:
   BenchUut6.cyclicExecution := FALSE;
   BenchUut6.trigger := FALSE;
   BenchUut6.value := LREAL#67.0;
   BenchUut6.windowSize := INT#100;
   BenchUut6.reset := FALSE;
   TraceIn_cyclicExecution[377] := BenchUut6.cyclicExecution;
   TraceIn_trigger[377] := BenchUut6.trigger;
   TraceIn_value[377] := BenchUut6.value;
   TraceIn_windowSize[377] := BenchUut6.windowSize;
   TraceIn_reset[377] := BenchUut6.reset;
   BenchUut6();
   TraceOut_average[377] := BenchUut6.average;
   TraceOut_windowSizeReached[377] := BenchUut6.windowSizeReached;
   TraceOut_error[377] := BenchUut6.error;
   TraceOut_status[377] := BenchUut6.status;
   BenchCalls := BenchCalls + 1;
 378:
   BenchUut6.cyclicExecution := FALSE;
   BenchUut6.trigger := TRUE;
   BenchUut6.value := LREAL#68.0;
   BenchUut6.windowSize := INT#100;
   BenchUut6.reset := FALSE;
   TraceIn_cyclicExecution[378] := BenchUut6.cyclicExecution;
   TraceIn_trigger[378] := BenchUut6.trigger;
   TraceIn_value[378] := BenchUut6.value;
   TraceIn_windowSize[378] := BenchUut6.windowSize;
   TraceIn_reset[378] := BenchUut6.reset;
   BenchUut6();
   TraceOut_average[378] := BenchUut6.average;
   TraceOut_windowSizeReached[378] := BenchUut6.windowSizeReached;
   TraceOut_error[378] := BenchUut6.error;
   TraceOut_status[378] := BenchUut6.status;
   BenchCalls := BenchCalls + 1;
 379:
   BenchUut6.cyclicExecution := FALSE;
   BenchUut6.trigger := FALSE;
   BenchUut6.value := LREAL#68.0;
   BenchUut6.windowSize := INT#100;
   BenchUut6.reset := FALSE;
   TraceIn_cyclicExecution[379] := BenchUut6.cyclicExecution;
   TraceIn_trigger[379] := BenchUut6.trigger;
   TraceIn_value[379] := BenchUut6.value;
   TraceIn_windowSize[379] := BenchUut6.windowSize;
   TraceIn_reset[379] := BenchUut6.reset;
   BenchUut6();
   TraceOut_average[379] := BenchUut6.average;
   TraceOut_windowSizeReached[379] := BenchUut6.windowSizeReached;
   TraceOut_error[379] := BenchUut6.error;
   TraceOut_status[379] := BenchUut6.status;
   BenchCalls := BenchCalls + 1;
 380:
   BenchUut6.cyclicExecution := FALSE;
   BenchUut6.trigger := TRUE;
   BenchUut6.value := LREAL#69.0;
   BenchUut6.windowSize := INT#100;
   BenchUut6.reset := FALSE;
   TraceIn_cyclicExecution[380] := BenchUut6.cyclicExecution;
   TraceIn_trigger[380] := BenchUut6.trigger;
   TraceIn_value[380] := BenchUut6.value;
   TraceIn_windowSize[380] := BenchUut6.windowSize;
   TraceIn_reset[380] := BenchUut6.reset;
   BenchUut6();
   TraceOut_average[380] := BenchUut6.average;
   TraceOut_windowSizeReached[380] := BenchUut6.windowSizeReached;
   TraceOut_error[380] := BenchUut6.error;
   TraceOut_status[380] := BenchUut6.status;
   BenchCalls := BenchCalls + 1;
 381:
   BenchUut6.cyclicExecution := FALSE;
   BenchUut6.trigger := FALSE;
   BenchUut6.value := LREAL#69.0;
   BenchUut6.windowSize := INT#100;
   BenchUut6.reset := FALSE;
   TraceIn_cyclicExecution[381] := BenchUut6.cyclicExecution;
   TraceIn_trigger[381] := BenchUut6.trigger;
   TraceIn_value[381] := BenchUut6.value;
   TraceIn_windowSize[381] := BenchUut6.windowSize;
   TraceIn_reset[381] := BenchUut6.reset;
   BenchUut6();
   TraceOut_average[381] := BenchUut6.average;
   TraceOut_windowSizeReached[381] := BenchUut6.windowSizeReached;
   TraceOut_error[381] := BenchUut6.error;
   TraceOut_status[381] := BenchUut6.status;
   BenchCalls := BenchCalls + 1;
 382:
   BenchUut6.cyclicExecution := FALSE;
   BenchUut6.trigger := TRUE;
   BenchUut6.value := LREAL#70.0;
   BenchUut6.windowSize := INT#100;
   BenchUut6.reset := FALSE;
   TraceIn_cyclicExecution[382] := BenchUut6.cyclicExecution;
   TraceIn_trigger[382] := BenchUut6.trigger;
   TraceIn_value[382] := BenchUut6.value;
   TraceIn_windowSize[382] := BenchUut6.windowSize;
   TraceIn_reset[382] := BenchUut6.reset;
   BenchUut6();
   TraceOut_average[382] := BenchUut6.average;
   TraceOut_windowSizeReached[382] := BenchUut6.windowSizeReached;
   TraceOut_error[382] := BenchUut6.error;
   TraceOut_status[382] := BenchUut6.status;
   BenchCalls := BenchCalls + 1;
 383:
   BenchUut6.cyclicExecution := FALSE;
   BenchUut6.trigger := FALSE;
   BenchUut6.value := LREAL#70.0;
   BenchUut6.windowSize := INT#100;
   BenchUut6.reset := FALSE;
   TraceIn_cyclicExecution[383] := BenchUut6.cyclicExecution;
   TraceIn_trigger[383] := BenchUut6.trigger;
   TraceIn_value[383] := BenchUut6.value;
   TraceIn_windowSize[383] := BenchUut6.windowSize;
   TraceIn_reset[383] := BenchUut6.reset;
   BenchUut6();
   TraceOut_average[383] := BenchUut6.average;
   TraceOut_windowSizeReached[383] := BenchUut6.windowSizeReached;
   TraceOut_error[383] := BenchUut6.error;
   TraceOut_status[383] := BenchUut6.status;
   BenchCalls := BenchCalls + 1;
 384:
   BenchUut6.cyclicExecution := FALSE;
   BenchUut6.trigger := TRUE;
   BenchUut6.value := LREAL#71.0;
   BenchUut6.windowSize := INT#100;
   BenchUut6.reset := FALSE;
   TraceIn_cyclicExecution[384] := BenchUut6.cyclicExecution;
   TraceIn_trigger[384] := BenchUut6.trigger;
   TraceIn_value[384] := BenchUut6.value;
   TraceIn_windowSize[384] := BenchUut6.windowSize;
   TraceIn_reset[384] := BenchUut6.reset;
   BenchUut6();
   TraceOut_average[384] := BenchUut6.average;
   TraceOut_windowSizeReached[384] := BenchUut6.windowSizeReached;
   TraceOut_error[384] := BenchUut6.error;
   TraceOut_status[384] := BenchUut6.status;
   BenchCalls := BenchCalls + 1;
 385:
   BenchUut6.cyclicExecution := FALSE;
   BenchUut6.trigger := FALSE;
   BenchUut6.value := LREAL#71.0;
   BenchUut6.windowSize := INT#100;
   BenchUut6.reset := FALSE;
   TraceIn_cyclicExecution[385] := BenchUut6.cyclicExecution;
   TraceIn_trigger[385] := BenchUut6.trigger;
   TraceIn_value[385] := BenchUut6.value;
   TraceIn_windowSize[385] := BenchUut6.windowSize;
   TraceIn_reset[385] := BenchUut6.reset;
   BenchUut6();
   TraceOut_average[385] := BenchUut6.average;
   TraceOut_windowSizeReached[385] := BenchUut6.windowSizeReached;
   TraceOut_error[385] := BenchUut6.error;
   TraceOut_status[385] := BenchUut6.status;
   BenchCalls := BenchCalls + 1;
 386:
   BenchUut6.cyclicExecution := FALSE;
   BenchUut6.trigger := TRUE;
   BenchUut6.value := LREAL#72.0;
   BenchUut6.windowSize := INT#100;
   BenchUut6.reset := FALSE;
   TraceIn_cyclicExecution[386] := BenchUut6.cyclicExecution;
   TraceIn_trigger[386] := BenchUut6.trigger;
   TraceIn_value[386] := BenchUut6.value;
   TraceIn_windowSize[386] := BenchUut6.windowSize;
   TraceIn_reset[386] := BenchUut6.reset;
   BenchUut6();
   TraceOut_average[386] := BenchUut6.average;
   TraceOut_windowSizeReached[386] := BenchUut6.windowSizeReached;
   TraceOut_error[386] := BenchUut6.error;
   TraceOut_status[386] := BenchUut6.status;
   BenchCalls := BenchCalls + 1;
 387:
   BenchUut6.cyclicExecution := FALSE;
   BenchUut6.trigger := FALSE;
   BenchUut6.value := LREAL#72.0;
   BenchUut6.windowSize := INT#100;
   BenchUut6.reset := FALSE;
   TraceIn_cyclicExecution[387] := BenchUut6.cyclicExecution;
   TraceIn_trigger[387] := BenchUut6.trigger;
   TraceIn_value[387] := BenchUut6.value;
   TraceIn_windowSize[387] := BenchUut6.windowSize;
   TraceIn_reset[387] := BenchUut6.reset;
   BenchUut6();
   TraceOut_average[387] := BenchUut6.average;
   TraceOut_windowSizeReached[387] := BenchUut6.windowSizeReached;
   TraceOut_error[387] := BenchUut6.error;
   TraceOut_status[387] := BenchUut6.status;
   BenchCalls := BenchCalls + 1;
 388:
   BenchUut6.cyclicExecution := FALSE;
   BenchUut6.trigger := TRUE;
   BenchUut6.value := LREAL#73.0;
   BenchUut6.windowSize := INT#100;
   BenchUut6.reset := FALSE;
   TraceIn_cyclicExecution[388] := BenchUut6.cyclicExecution;
   TraceIn_trigger[388] := BenchUut6.trigger;
   TraceIn_value[388] := BenchUut6.value;
   TraceIn_windowSize[388] := BenchUut6.windowSize;
   TraceIn_reset[388] := BenchUut6.reset;
   BenchUut6();
   TraceOut_average[388] := BenchUut6.average;
   TraceOut_windowSizeReached[388] := BenchUut6.windowSizeReached;
   TraceOut_error[388] := BenchUut6.error;
   TraceOut_status[388] := BenchUut6.status;
   BenchCalls := BenchCalls + 1;
 389:
   BenchUut6.cyclicExecution := FALSE;
   BenchUut6.trigger := FALSE;
   BenchUut6.value := LREAL#73.0;
   BenchUut6.windowSize := INT#100;
   BenchUut6.reset := FALSE;
   TraceIn_cyclicExecution[389] := BenchUut6.cyclicExecution;
   TraceIn_trigger[389] := BenchUut6.trigger;
   TraceIn_value[389] := BenchUut6.value;
   TraceIn_windowSize[389] := BenchUut6.windowSize;
   TraceIn_reset[389] := BenchUut6.reset;
   BenchUut6();
   TraceOut_average[389] := BenchUut6.average;
   TraceOut_windowSizeReached[389] := BenchUut6.windowSizeReached;
   TraceOut_error[389] := BenchUut6.error;
   TraceOut_status[389] := BenchUut6.status;
   BenchCalls := BenchCalls + 1;
 390:
   BenchUut6.cyclicExecution := FALSE;
   BenchUut6.trigger := TRUE;
   BenchUut6.value := LREAL#74.0;
   BenchUut6.windowSize := INT#100;
   BenchUut6.reset := FALSE;
   TraceIn_cyclicExecution[390] := BenchUut6.cyclicExecution;
   TraceIn_trigger[390] := BenchUut6.trigger;
   TraceIn_value[390] := BenchUut6.value;
   TraceIn_windowSize[390] := BenchUut6.windowSize;
   TraceIn_reset[390] := BenchUut6.reset;
   BenchUut6();
   TraceOut_average[390] := BenchUut6.average;
   TraceOut_windowSizeReached[390] := BenchUut6.windowSizeReached;
   TraceOut_error[390] := BenchUut6.error;
   TraceOut_status[390] := BenchUut6.status;
   BenchCalls := BenchCalls + 1;
 391:
   BenchUut6.cyclicExecution := FALSE;
   BenchUut6.trigger := FALSE;
   BenchUut6.value := LREAL#74.0;
   BenchUut6.windowSize := INT#100;
   BenchUut6.reset := FALSE;
   TraceIn_cyclicExecution[391] := BenchUut6.cyclicExecution;
   TraceIn_trigger[391] := BenchUut6.trigger;
   TraceIn_value[391] := BenchUut6.value;
   TraceIn_windowSize[391] := BenchUut6.windowSize;
   TraceIn_reset[391] := BenchUut6.reset;
   BenchUut6();
   TraceOut_average[391] := BenchUut6.average;
   TraceOut_windowSizeReached[391] := BenchUut6.windowSizeReached;
   TraceOut_error[391] := BenchUut6.error;
   TraceOut_status[391] := BenchUut6.status;
   BenchCalls := BenchCalls + 1;
 392:
   BenchUut6.cyclicExecution := FALSE;
   BenchUut6.trigger := TRUE;
   BenchUut6.value := LREAL#75.0;
   BenchUut6.windowSize := INT#100;
   BenchUut6.reset := FALSE;
   TraceIn_cyclicExecution[392] := BenchUut6.cyclicExecution;
   TraceIn_trigger[392] := BenchUut6.trigger;
   TraceIn_value[392] := BenchUut6.value;
   TraceIn_windowSize[392] := BenchUut6.windowSize;
   TraceIn_reset[392] := BenchUut6.reset;
   BenchUut6();
   TraceOut_average[392] := BenchUut6.average;
   TraceOut_windowSizeReached[392] := BenchUut6.windowSizeReached;
   TraceOut_error[392] := BenchUut6.error;
   TraceOut_status[392] := BenchUut6.status;
   BenchCalls := BenchCalls + 1;
 393:
   BenchUut6.cyclicExecution := FALSE;
   BenchUut6.trigger := FALSE;
   BenchUut6.value := LREAL#75.0;
   BenchUut6.windowSize := INT#100;
   BenchUut6.reset := FALSE;
   TraceIn_cyclicExecution[393] := BenchUut6.cyclicExecution;
   TraceIn_trigger[393] := BenchUut6.trigger;
   TraceIn_value[393] := BenchUut6.value;
   TraceIn_windowSize[393] := BenchUut6.windowSize;
   TraceIn_reset[393] := BenchUut6.reset;
   BenchUut6();
   TraceOut_average[393] := BenchUut6.average;
   TraceOut_windowSizeReached[393] := BenchUut6.windowSizeReached;
   TraceOut_error[393] := BenchUut6.error;
   TraceOut_status[393] := BenchUut6.status;
   BenchCalls := BenchCalls + 1;
 394:
   BenchUut6.cyclicExecution := FALSE;
   BenchUut6.trigger := TRUE;
   BenchUut6.value := LREAL#76.0;
   BenchUut6.windowSize := INT#100;
   BenchUut6.reset := FALSE;
   TraceIn_cyclicExecution[394] := BenchUut6.cyclicExecution;
   TraceIn_trigger[394] := BenchUut6.trigger;
   TraceIn_value[394] := BenchUut6.value;
   TraceIn_windowSize[394] := BenchUut6.windowSize;
   TraceIn_reset[394] := BenchUut6.reset;
   BenchUut6();
   TraceOut_average[394] := BenchUut6.average;
   TraceOut_windowSizeReached[394] := BenchUut6.windowSizeReached;
   TraceOut_error[394] := BenchUut6.error;
   TraceOut_status[394] := BenchUut6.status;
   BenchCalls := BenchCalls + 1;
 395:
   BenchUut6.cyclicExecution := FALSE;
   BenchUut6.trigger := FALSE;
   BenchUut6.value := LREAL#76.0;
   BenchUut6.windowSize := INT#100;
   BenchUut6.reset := FALSE;
   TraceIn_cyclicExecution[395] := BenchUut6.cyclicExecution;
   TraceIn_trigger[395] := BenchUut6.trigger;
   TraceIn_value[395] := BenchUut6.value;
   TraceIn_windowSize[395] := BenchUut6.windowSize;
   TraceIn_reset[395] := BenchUut6.reset;
   BenchUut6();
   TraceOut_average[395] := BenchUut6.average;
   TraceOut_windowSizeReached[395] := BenchUut6.windowSizeReached;
   TraceOut_error[395] := BenchUut6.error;
   TraceOut_status[395] := BenchUut6.status;
   BenchCalls := BenchCalls + 1;
 396:
   BenchUut6.cyclicExecution := FALSE;
   BenchUut6.trigger := TRUE;
   BenchUut6.value := LREAL#77.0;
   BenchUut6.windowSize := INT#100;
   BenchUut6.reset := FALSE;
   TraceIn_cyclicExecution[396] := BenchUut6.cyclicExecution;
   TraceIn_trigger[396] := BenchUut6.trigger;
   TraceIn_value[396] := BenchUut6.value;
   TraceIn_windowSize[396] := BenchUut6.windowSize;
   TraceIn_reset[396] := BenchUut6.reset;
   BenchUut6();
   TraceOut_average[396] := BenchUut6.average;
   TraceOut_windowSizeReached[396] := BenchUut6.windowSizeReached;
   TraceOut_error[396] := BenchUut6.error;
   TraceOut_status[396] := BenchUut6.status;
   BenchCalls := BenchCalls + 1;
 397:
   BenchUut6.cyclicExecution := FALSE;
   BenchUut6.trigger := FALSE;
   BenchUut6.value := LREAL#77.0;
   BenchUut6.windowSize := INT#100;
   BenchUut6.reset := FALSE;
   TraceIn_cyclicExecution[397] := BenchUut6.cyclicExecution;
   TraceIn_trigger[397] := BenchUut6.trigger;
   TraceIn_value[397] := BenchUut6.value;
   TraceIn_windowSize[397] := BenchUut6.windowSize;
   TraceIn_reset[397] := BenchUut6.reset;
   BenchUut6();
   TraceOut_average[397] := BenchUut6.average;
   TraceOut_windowSizeReached[397] := BenchUut6.windowSizeReached;
   TraceOut_error[397] := BenchUut6.error;
   TraceOut_status[397] := BenchUut6.status;
   BenchCalls := BenchCalls + 1;
 398:
   BenchUut6.cyclicExecution := FALSE;
   BenchUut6.trigger := TRUE;
   BenchUut6.value := LREAL#78.0;
   BenchUut6.windowSize := INT#100;
   BenchUut6.reset := FALSE;
   TraceIn_cyclicExecution[398] := BenchUut6.cyclicExecution;
   TraceIn_trigger[398] := BenchUut6.trigger;
   TraceIn_value[398] := BenchUut6.value;
   TraceIn_windowSize[398] := BenchUut6.windowSize;
   TraceIn_reset[398] := BenchUut6.reset;
   BenchUut6();
   TraceOut_average[398] := BenchUut6.average;
   TraceOut_windowSizeReached[398] := BenchUut6.windowSizeReached;
   TraceOut_error[398] := BenchUut6.error;
   TraceOut_status[398] := BenchUut6.status;
   BenchCalls := BenchCalls + 1;
 399:
   BenchUut6.cyclicExecution := FALSE;
   BenchUut6.trigger := FALSE;
   BenchUut6.value := LREAL#78.0;
   BenchUut6.windowSize := INT#100;
   BenchUut6.reset := FALSE;
   TraceIn_cyclicExecution[399] := BenchUut6.cyclicExecution;
   TraceIn_trigger[399] := BenchUut6.trigger;
   TraceIn_value[399] := BenchUut6.value;
   TraceIn_windowSize[399] := BenchUut6.windowSize;
   TraceIn_reset[399] := BenchUut6.reset;
   BenchUut6();
   TraceOut_average[399] := BenchUut6.average;
   TraceOut_windowSizeReached[399] := BenchUut6.windowSizeReached;
   TraceOut_error[399] := BenchUut6.error;
   TraceOut_status[399] := BenchUut6.status;
   BenchCalls := BenchCalls + 1;
 400:
   BenchUut6.cyclicExecution := FALSE;
   BenchUut6.trigger := TRUE;
   BenchUut6.value := LREAL#79.0;
   BenchUut6.windowSize := INT#100;
   BenchUut6.reset := FALSE;
   TraceIn_cyclicExecution[400] := BenchUut6.cyclicExecution;
   TraceIn_trigger[400] := BenchUut6.trigger;
   TraceIn_value[400] := BenchUut6.value;
   TraceIn_windowSize[400] := BenchUut6.windowSize;
   TraceIn_reset[400] := BenchUut6.reset;
   BenchUut6();
   TraceOut_average[400] := BenchUut6.average;
   TraceOut_windowSizeReached[400] := BenchUut6.windowSizeReached;
   TraceOut_error[400] := BenchUut6.error;
   TraceOut_status[400] := BenchUut6.status;
   BenchCalls := BenchCalls + 1;
 401:
   BenchUut6.cyclicExecution := FALSE;
   BenchUut6.trigger := FALSE;
   BenchUut6.value := LREAL#79.0;
   BenchUut6.windowSize := INT#100;
   BenchUut6.reset := FALSE;
   TraceIn_cyclicExecution[401] := BenchUut6.cyclicExecution;
   TraceIn_trigger[401] := BenchUut6.trigger;
   TraceIn_value[401] := BenchUut6.value;
   TraceIn_windowSize[401] := BenchUut6.windowSize;
   TraceIn_reset[401] := BenchUut6.reset;
   BenchUut6();
   TraceOut_average[401] := BenchUut6.average;
   TraceOut_windowSizeReached[401] := BenchUut6.windowSizeReached;
   TraceOut_error[401] := BenchUut6.error;
   TraceOut_status[401] := BenchUut6.status;
   BenchCalls := BenchCalls + 1;
 402:
   BenchUut6.cyclicExecution := FALSE;
   BenchUut6.trigger := TRUE;
   BenchUut6.value := LREAL#80.0;
   BenchUut6.windowSize := INT#100;
   BenchUut6.reset := FALSE;
   TraceIn_cyclicExecution[402] := BenchUut6.cyclicExecution;
   TraceIn_trigger[402] := BenchUut6.trigger;
   TraceIn_value[402] := BenchUut6.value;
   TraceIn_windowSize[402] := BenchUut6.windowSize;
   TraceIn_reset[402] := BenchUut6.reset;
   BenchUut6();
   TraceOut_average[402] := BenchUut6.average;
   TraceOut_windowSizeReached[402] := BenchUut6.windowSizeReached;
   TraceOut_error[402] := BenchUut6.error;
   TraceOut_status[402] := BenchUut6.status;
   BenchCalls := BenchCalls + 1;
 403:
   BenchUut6.cyclicExecution := FALSE;
   BenchUut6.trigger := FALSE;
   BenchUut6.value := LREAL#80.0;
   BenchUut6.windowSize := INT#100;
   BenchUut6.reset := FALSE;
   TraceIn_cyclicExecution[403] := BenchUut6.cyclicExecution;
   TraceIn_trigger[403] := BenchUut6.trigger;
   TraceIn_value[403] := BenchUut6.value;
   TraceIn_windowSize[403] := BenchUut6.windowSize;
   TraceIn_reset[403] := BenchUut6.reset;
   BenchUut6();
   TraceOut_average[403] := BenchUut6.average;
   TraceOut_windowSizeReached[403] := BenchUut6.windowSizeReached;
   TraceOut_error[403] := BenchUut6.error;
   TraceOut_status[403] := BenchUut6.status;
   BenchCalls := BenchCalls + 1;
 404:
   BenchUut6.cyclicExecution := FALSE;
   BenchUut6.trigger := TRUE;
   BenchUut6.value := LREAL#81.0;
   BenchUut6.windowSize := INT#100;
   BenchUut6.reset := FALSE;
   TraceIn_cyclicExecution[404] := BenchUut6.cyclicExecution;
   TraceIn_trigger[404] := BenchUut6.trigger;
   TraceIn_value[404] := BenchUut6.value;
   TraceIn_windowSize[404] := BenchUut6.windowSize;
   TraceIn_reset[404] := BenchUut6.reset;
   BenchUut6();
   TraceOut_average[404] := BenchUut6.average;
   TraceOut_windowSizeReached[404] := BenchUut6.windowSizeReached;
   TraceOut_error[404] := BenchUut6.error;
   TraceOut_status[404] := BenchUut6.status;
   BenchCalls := BenchCalls + 1;
 405:
   BenchUut6.cyclicExecution := FALSE;
   BenchUut6.trigger := FALSE;
   BenchUut6.value := LREAL#81.0;
   BenchUut6.windowSize := INT#100;
   BenchUut6.reset := FALSE;
   TraceIn_cyclicExecution[405] := BenchUut6.cyclicExecution;
   TraceIn_trigger[405] := BenchUut6.trigger;
   TraceIn_value[405] := BenchUut6.value;
   TraceIn_windowSize[405] := BenchUut6.windowSize;
   TraceIn_reset[405] := BenchUut6.reset;
   BenchUut6();
   TraceOut_average[405] := BenchUut6.average;
   TraceOut_windowSizeReached[405] := BenchUut6.windowSizeReached;
   TraceOut_error[405] := BenchUut6.error;
   TraceOut_status[405] := BenchUut6.status;
   BenchCalls := BenchCalls + 1;
 406:
   BenchUut6.cyclicExecution := FALSE;
   BenchUut6.trigger := TRUE;
   BenchUut6.value := LREAL#82.0;
   BenchUut6.windowSize := INT#100;
   BenchUut6.reset := FALSE;
   TraceIn_cyclicExecution[406] := BenchUut6.cyclicExecution;
   TraceIn_trigger[406] := BenchUut6.trigger;
   TraceIn_value[406] := BenchUut6.value;
   TraceIn_windowSize[406] := BenchUut6.windowSize;
   TraceIn_reset[406] := BenchUut6.reset;
   BenchUut6();
   TraceOut_average[406] := BenchUut6.average;
   TraceOut_windowSizeReached[406] := BenchUut6.windowSizeReached;
   TraceOut_error[406] := BenchUut6.error;
   TraceOut_status[406] := BenchUut6.status;
   BenchCalls := BenchCalls + 1;
 407:
   BenchUut6.cyclicExecution := FALSE;
   BenchUut6.trigger := FALSE;
   BenchUut6.value := LREAL#82.0;
   BenchUut6.windowSize := INT#100;
   BenchUut6.reset := FALSE;
   TraceIn_cyclicExecution[407] := BenchUut6.cyclicExecution;
   TraceIn_trigger[407] := BenchUut6.trigger;
   TraceIn_value[407] := BenchUut6.value;
   TraceIn_windowSize[407] := BenchUut6.windowSize;
   TraceIn_reset[407] := BenchUut6.reset;
   BenchUut6();
   TraceOut_average[407] := BenchUut6.average;
   TraceOut_windowSizeReached[407] := BenchUut6.windowSizeReached;
   TraceOut_error[407] := BenchUut6.error;
   TraceOut_status[407] := BenchUut6.status;
   BenchCalls := BenchCalls + 1;
 408:
   BenchUut6.cyclicExecution := FALSE;
   BenchUut6.trigger := TRUE;
   BenchUut6.value := LREAL#83.0;
   BenchUut6.windowSize := INT#100;
   BenchUut6.reset := FALSE;
   TraceIn_cyclicExecution[408] := BenchUut6.cyclicExecution;
   TraceIn_trigger[408] := BenchUut6.trigger;
   TraceIn_value[408] := BenchUut6.value;
   TraceIn_windowSize[408] := BenchUut6.windowSize;
   TraceIn_reset[408] := BenchUut6.reset;
   BenchUut6();
   TraceOut_average[408] := BenchUut6.average;
   TraceOut_windowSizeReached[408] := BenchUut6.windowSizeReached;
   TraceOut_error[408] := BenchUut6.error;
   TraceOut_status[408] := BenchUut6.status;
   BenchCalls := BenchCalls + 1;
 409:
   BenchUut6.cyclicExecution := FALSE;
   BenchUut6.trigger := FALSE;
   BenchUut6.value := LREAL#83.0;
   BenchUut6.windowSize := INT#100;
   BenchUut6.reset := FALSE;
   TraceIn_cyclicExecution[409] := BenchUut6.cyclicExecution;
   TraceIn_trigger[409] := BenchUut6.trigger;
   TraceIn_value[409] := BenchUut6.value;
   TraceIn_windowSize[409] := BenchUut6.windowSize;
   TraceIn_reset[409] := BenchUut6.reset;
   BenchUut6();
   TraceOut_average[409] := BenchUut6.average;
   TraceOut_windowSizeReached[409] := BenchUut6.windowSizeReached;
   TraceOut_error[409] := BenchUut6.error;
   TraceOut_status[409] := BenchUut6.status;
   BenchCalls := BenchCalls + 1;
 410:
   BenchUut6.cyclicExecution := FALSE;
   BenchUut6.trigger := TRUE;
   BenchUut6.value := LREAL#84.0;
   BenchUut6.windowSize := INT#100;
   BenchUut6.reset := FALSE;
   TraceIn_cyclicExecution[410] := BenchUut6.cyclicExecution;
   TraceIn_trigger[410] := BenchUut6.trigger;
   TraceIn_value[410] := BenchUut6.value;
   TraceIn_windowSize[410] := BenchUut6.windowSize;
   TraceIn_reset[410] := BenchUut6.reset;
   BenchUut6();
   TraceOut_average[410] := BenchUut6.average;
   TraceOut_windowSizeReached[410] := BenchUut6.windowSizeReached;
   TraceOut_error[410] := BenchUut6.error;
   TraceOut_status[410] := BenchUut6.status;
   BenchCalls := BenchCalls + 1;
 411:
   BenchUut6.cyclicExecution := FALSE;
   BenchUut6.trigger := FALSE;
   BenchUut6.value := LREAL#84.0;
   BenchUut6.windowSize := INT#100;
   BenchUut6.reset := FALSE;
   TraceIn_cyclicExecution[411] := BenchUut6.cyclicExecution;
   TraceIn_trigger[411] := BenchUut6.trigger;
   TraceIn_value[411] := BenchUut6.value;
   TraceIn_windowSize[411] := BenchUut6.windowSize;
   TraceIn_reset[411] := BenchUut6.reset;
   BenchUut6();
   TraceOut_average[411] := BenchUut6.average;
   TraceOut_windowSizeReached[411] := BenchUut6.windowSizeReached;
   TraceOut_error[411] := BenchUut6.error;
   TraceOut_status[411] := BenchUut6.status;
   BenchCalls := BenchCalls + 1;
 412:
   BenchUut6.cyclicExecution := FALSE;
   BenchUut6.trigger := TRUE;
   BenchUut6.value := LREAL#85.0;
   BenchUut6.windowSize := INT#100;
   BenchUut6.reset := FALSE;
   TraceIn_cyclicExecution[412] := BenchUut6.cyclicExecution;
   TraceIn_trigger[412] := BenchUut6.trigger;
   TraceIn_value[412] := BenchUut6.value;
   TraceIn_windowSize[412] := BenchUut6.windowSize;
   TraceIn_reset[412] := BenchUut6.reset;
   BenchUut6();
   TraceOut_average[412] := BenchUut6.average;
   TraceOut_windowSizeReached[412] := BenchUut6.windowSizeReached;
   TraceOut_error[412] := BenchUut6.error;
   TraceOut_status[412] := BenchUut6.status;
   BenchCalls := BenchCalls + 1;
 413:
   BenchUut6.cyclicExecution := FALSE;
   BenchUut6.trigger := FALSE;
   BenchUut6.value := LREAL#85.0;
   BenchUut6.windowSize := INT#100;
   BenchUut6.reset := FALSE;
   TraceIn_cyclicExecution[413] := BenchUut6.cyclicExecution;
   TraceIn_trigger[413] := BenchUut6.trigger;
   TraceIn_value[413] := BenchUut6.value;
   TraceIn_windowSize[413] := BenchUut6.windowSize;
   TraceIn_reset[413] := BenchUut6.reset;
   BenchUut6();
   TraceOut_average[413] := BenchUut6.average;
   TraceOut_windowSizeReached[413] := BenchUut6.windowSizeReached;
   TraceOut_error[413] := BenchUut6.error;
   TraceOut_status[413] := BenchUut6.status;
   BenchCalls := BenchCalls + 1;
 414:
   BenchUut6.cyclicExecution := FALSE;
   BenchUut6.trigger := TRUE;
   BenchUut6.value := LREAL#86.0;
   BenchUut6.windowSize := INT#100;
   BenchUut6.reset := FALSE;
   TraceIn_cyclicExecution[414] := BenchUut6.cyclicExecution;
   TraceIn_trigger[414] := BenchUut6.trigger;
   TraceIn_value[414] := BenchUut6.value;
   TraceIn_windowSize[414] := BenchUut6.windowSize;
   TraceIn_reset[414] := BenchUut6.reset;
   BenchUut6();
   TraceOut_average[414] := BenchUut6.average;
   TraceOut_windowSizeReached[414] := BenchUut6.windowSizeReached;
   TraceOut_error[414] := BenchUut6.error;
   TraceOut_status[414] := BenchUut6.status;
   BenchCalls := BenchCalls + 1;
 415:
   BenchUut6.cyclicExecution := FALSE;
   BenchUut6.trigger := FALSE;
   BenchUut6.value := LREAL#86.0;
   BenchUut6.windowSize := INT#100;
   BenchUut6.reset := FALSE;
   TraceIn_cyclicExecution[415] := BenchUut6.cyclicExecution;
   TraceIn_trigger[415] := BenchUut6.trigger;
   TraceIn_value[415] := BenchUut6.value;
   TraceIn_windowSize[415] := BenchUut6.windowSize;
   TraceIn_reset[415] := BenchUut6.reset;
   BenchUut6();
   TraceOut_average[415] := BenchUut6.average;
   TraceOut_windowSizeReached[415] := BenchUut6.windowSizeReached;
   TraceOut_error[415] := BenchUut6.error;
   TraceOut_status[415] := BenchUut6.status;
   BenchCalls := BenchCalls + 1;
 416:
   BenchUut6.cyclicExecution := FALSE;
   BenchUut6.trigger := TRUE;
   BenchUut6.value := LREAL#87.0;
   BenchUut6.windowSize := INT#100;
   BenchUut6.reset := FALSE;
   TraceIn_cyclicExecution[416] := BenchUut6.cyclicExecution;
   TraceIn_trigger[416] := BenchUut6.trigger;
   TraceIn_value[416] := BenchUut6.value;
   TraceIn_windowSize[416] := BenchUut6.windowSize;
   TraceIn_reset[416] := BenchUut6.reset;
   BenchUut6();
   TraceOut_average[416] := BenchUut6.average;
   TraceOut_windowSizeReached[416] := BenchUut6.windowSizeReached;
   TraceOut_error[416] := BenchUut6.error;
   TraceOut_status[416] := BenchUut6.status;
   BenchCalls := BenchCalls + 1;
 417:
   BenchUut6.cyclicExecution := FALSE;
   BenchUut6.trigger := FALSE;
   BenchUut6.value := LREAL#87.0;
   BenchUut6.windowSize := INT#100;
   BenchUut6.reset := FALSE;
   TraceIn_cyclicExecution[417] := BenchUut6.cyclicExecution;
   TraceIn_trigger[417] := BenchUut6.trigger;
   TraceIn_value[417] := BenchUut6.value;
   TraceIn_windowSize[417] := BenchUut6.windowSize;
   TraceIn_reset[417] := BenchUut6.reset;
   BenchUut6();
   TraceOut_average[417] := BenchUut6.average;
   TraceOut_windowSizeReached[417] := BenchUut6.windowSizeReached;
   TraceOut_error[417] := BenchUut6.error;
   TraceOut_status[417] := BenchUut6.status;
   BenchCalls := BenchCalls + 1;
 418:
   BenchUut6.cyclicExecution := FALSE;
   BenchUut6.trigger := TRUE;
   BenchUut6.value := LREAL#88.0;
   BenchUut6.windowSize := INT#100;
   BenchUut6.reset := FALSE;
   TraceIn_cyclicExecution[418] := BenchUut6.cyclicExecution;
   TraceIn_trigger[418] := BenchUut6.trigger;
   TraceIn_value[418] := BenchUut6.value;
   TraceIn_windowSize[418] := BenchUut6.windowSize;
   TraceIn_reset[418] := BenchUut6.reset;
   BenchUut6();
   TraceOut_average[418] := BenchUut6.average;
   TraceOut_windowSizeReached[418] := BenchUut6.windowSizeReached;
   TraceOut_error[418] := BenchUut6.error;
   TraceOut_status[418] := BenchUut6.status;
   BenchCalls := BenchCalls + 1;
 419:
   BenchUut6.cyclicExecution := FALSE;
   BenchUut6.trigger := FALSE;
   BenchUut6.value := LREAL#88.0;
   BenchUut6.windowSize := INT#100;
   BenchUut6.reset := FALSE;
   TraceIn_cyclicExecution[419] := BenchUut6.cyclicExecution;
   TraceIn_trigger[419] := BenchUut6.trigger;
   TraceIn_value[419] := BenchUut6.value;
   TraceIn_windowSize[419] := BenchUut6.windowSize;
   TraceIn_reset[419] := BenchUut6.reset;
   BenchUut6();
   TraceOut_average[419] := BenchUut6.average;
   TraceOut_windowSizeReached[419] := BenchUut6.windowSizeReached;
   TraceOut_error[419] := BenchUut6.error;
   TraceOut_status[419] := BenchUut6.status;
   BenchCalls := BenchCalls + 1;
 420:
   BenchUut6.cyclicExecution := FALSE;
   BenchUut6.trigger := TRUE;
   BenchUut6.value := LREAL#89.0;
   BenchUut6.windowSize := INT#100;
   BenchUut6.reset := FALSE;
   TraceIn_cyclicExecution[420] := BenchUut6.cyclicExecution;
   TraceIn_trigger[420] := BenchUut6.trigger;
   TraceIn_value[420] := BenchUut6.value;
   TraceIn_windowSize[420] := BenchUut6.windowSize;
   TraceIn_reset[420] := BenchUut6.reset;
   BenchUut6();
   TraceOut_average[420] := BenchUut6.average;
   TraceOut_windowSizeReached[420] := BenchUut6.windowSizeReached;
   TraceOut_error[420] := BenchUut6.error;
   TraceOut_status[420] := BenchUut6.status;
   BenchCalls := BenchCalls + 1;
 421:
   BenchUut6.cyclicExecution := FALSE;
   BenchUut6.trigger := FALSE;
   BenchUut6.value := LREAL#89.0;
   BenchUut6.windowSize := INT#100;
   BenchUut6.reset := FALSE;
   TraceIn_cyclicExecution[421] := BenchUut6.cyclicExecution;
   TraceIn_trigger[421] := BenchUut6.trigger;
   TraceIn_value[421] := BenchUut6.value;
   TraceIn_windowSize[421] := BenchUut6.windowSize;
   TraceIn_reset[421] := BenchUut6.reset;
   BenchUut6();
   TraceOut_average[421] := BenchUut6.average;
   TraceOut_windowSizeReached[421] := BenchUut6.windowSizeReached;
   TraceOut_error[421] := BenchUut6.error;
   TraceOut_status[421] := BenchUut6.status;
   BenchCalls := BenchCalls + 1;
 422:
   BenchUut6.cyclicExecution := FALSE;
   BenchUut6.trigger := TRUE;
   BenchUut6.value := LREAL#90.0;
   BenchUut6.windowSize := INT#100;
   BenchUut6.reset := FALSE;
   TraceIn_cyclicExecution[422] := BenchUut6.cyclicExecution;
   TraceIn_trigger[422] := BenchUut6.trigger;
   TraceIn_value[422] := BenchUut6.value;
   TraceIn_windowSize[422] := BenchUut6.windowSize;
   TraceIn_reset[422] := BenchUut6.reset;
   BenchUut6();
   TraceOut_average[422] := BenchUut6.average;
   TraceOut_windowSizeReached[422] := BenchUut6.windowSizeReached;
   TraceOut_error[422] := BenchUut6.error;
   TraceOut_status[422] := BenchUut6.status;
   BenchCalls := BenchCalls + 1;
 423:
   BenchUut6.cyclicExecution := FALSE;
   BenchUut6.trigger := FALSE;
   BenchUut6.value := LREAL#90.0;
   BenchUut6.windowSize := INT#100;
   BenchUut6.reset := FALSE;
   TraceIn_cyclicExecution[423] := BenchUut6.cyclicExecution;
   TraceIn_trigger[423] := BenchUut6.trigger;
   TraceIn_value[423] := BenchUut6.value;
   TraceIn_windowSize[423] := BenchUut6.windowSize;
   TraceIn_reset[423] := BenchUut6.reset;
   BenchUut6();
   TraceOut_average[423] := BenchUut6.average;
   TraceOut_windowSizeReached[423] := BenchUut6.windowSizeReached;
   TraceOut_error[423] := BenchUut6.error;
   TraceOut_status[423] := BenchUut6.status;
   BenchCalls := BenchCalls + 1;
 424:
   BenchUut6.cyclicExecution := FALSE;
   BenchUut6.trigger := TRUE;
   BenchUut6.value := LREAL#91.0;
   BenchUut6.windowSize := INT#100;
   BenchUut6.reset := FALSE;
   TraceIn_cyclicExecution[424] := BenchUut6.cyclicExecution;
   TraceIn_trigger[424] := BenchUut6.trigger;
   TraceIn_value[424] := BenchUut6.value;
   TraceIn_windowSize[424] := BenchUut6.windowSize;
   TraceIn_reset[424] := BenchUut6.reset;
   BenchUut6();
   TraceOut_average[424] := BenchUut6.average;
   TraceOut_windowSizeReached[424] := BenchUut6.windowSizeReached;
   TraceOut_error[424] := BenchUut6.error;
   TraceOut_status[424] := BenchUut6.status;
   BenchCalls := BenchCalls + 1;
 425:
   BenchUut6.cyclicExecution := FALSE;
   BenchUut6.trigger := FALSE;
   BenchUut6.value := LREAL#91.0;
   BenchUut6.windowSize := INT#100;
   BenchUut6.reset := FALSE;
   TraceIn_cyclicExecution[425] := BenchUut6.cyclicExecution;
   TraceIn_trigger[425] := BenchUut6.trigger;
   TraceIn_value[425] := BenchUut6.value;
   TraceIn_windowSize[425] := BenchUut6.windowSize;
   TraceIn_reset[425] := BenchUut6.reset;
   BenchUut6();
   TraceOut_average[425] := BenchUut6.average;
   TraceOut_windowSizeReached[425] := BenchUut6.windowSizeReached;
   TraceOut_error[425] := BenchUut6.error;
   TraceOut_status[425] := BenchUut6.status;
   BenchCalls := BenchCalls + 1;
 426:
   BenchUut6.cyclicExecution := FALSE;
   BenchUut6.trigger := TRUE;
   BenchUut6.value := LREAL#92.0;
   BenchUut6.windowSize := INT#100;
   BenchUut6.reset := FALSE;
   TraceIn_cyclicExecution[426] := BenchUut6.cyclicExecution;
   TraceIn_trigger[426] := BenchUut6.trigger;
   TraceIn_value[426] := BenchUut6.value;
   TraceIn_windowSize[426] := BenchUut6.windowSize;
   TraceIn_reset[426] := BenchUut6.reset;
   BenchUut6();
   TraceOut_average[426] := BenchUut6.average;
   TraceOut_windowSizeReached[426] := BenchUut6.windowSizeReached;
   TraceOut_error[426] := BenchUut6.error;
   TraceOut_status[426] := BenchUut6.status;
   BenchCalls := BenchCalls + 1;
 427:
   BenchUut6.cyclicExecution := FALSE;
   BenchUut6.trigger := FALSE;
   BenchUut6.value := LREAL#92.0;
   BenchUut6.windowSize := INT#100;
   BenchUut6.reset := FALSE;
   TraceIn_cyclicExecution[427] := BenchUut6.cyclicExecution;
   TraceIn_trigger[427] := BenchUut6.trigger;
   TraceIn_value[427] := BenchUut6.value;
   TraceIn_windowSize[427] := BenchUut6.windowSize;
   TraceIn_reset[427] := BenchUut6.reset;
   BenchUut6();
   TraceOut_average[427] := BenchUut6.average;
   TraceOut_windowSizeReached[427] := BenchUut6.windowSizeReached;
   TraceOut_error[427] := BenchUut6.error;
   TraceOut_status[427] := BenchUut6.status;
   BenchCalls := BenchCalls + 1;
 428:
   BenchUut6.cyclicExecution := FALSE;
   BenchUut6.trigger := TRUE;
   BenchUut6.value := LREAL#93.0;
   BenchUut6.windowSize := INT#100;
   BenchUut6.reset := FALSE;
   TraceIn_cyclicExecution[428] := BenchUut6.cyclicExecution;
   TraceIn_trigger[428] := BenchUut6.trigger;
   TraceIn_value[428] := BenchUut6.value;
   TraceIn_windowSize[428] := BenchUut6.windowSize;
   TraceIn_reset[428] := BenchUut6.reset;
   BenchUut6();
   TraceOut_average[428] := BenchUut6.average;
   TraceOut_windowSizeReached[428] := BenchUut6.windowSizeReached;
   TraceOut_error[428] := BenchUut6.error;
   TraceOut_status[428] := BenchUut6.status;
   BenchCalls := BenchCalls + 1;
 429:
   BenchUut6.cyclicExecution := FALSE;
   BenchUut6.trigger := FALSE;
   BenchUut6.value := LREAL#93.0;
   BenchUut6.windowSize := INT#100;
   BenchUut6.reset := FALSE;
   TraceIn_cyclicExecution[429] := BenchUut6.cyclicExecution;
   TraceIn_trigger[429] := BenchUut6.trigger;
   TraceIn_value[429] := BenchUut6.value;
   TraceIn_windowSize[429] := BenchUut6.windowSize;
   TraceIn_reset[429] := BenchUut6.reset;
   BenchUut6();
   TraceOut_average[429] := BenchUut6.average;
   TraceOut_windowSizeReached[429] := BenchUut6.windowSizeReached;
   TraceOut_error[429] := BenchUut6.error;
   TraceOut_status[429] := BenchUut6.status;
   BenchCalls := BenchCalls + 1;
 430:
   BenchUut6.cyclicExecution := FALSE;
   BenchUut6.trigger := TRUE;
   BenchUut6.value := LREAL#94.0;
   BenchUut6.windowSize := INT#100;
   BenchUut6.reset := FALSE;
   TraceIn_cyclicExecution[430] := BenchUut6.cyclicExecution;
   TraceIn_trigger[430] := BenchUut6.trigger;
   TraceIn_value[430] := BenchUut6.value;
   TraceIn_windowSize[430] := BenchUut6.windowSize;
   TraceIn_reset[430] := BenchUut6.reset;
   BenchUut6();
   TraceOut_average[430] := BenchUut6.average;
   TraceOut_windowSizeReached[430] := BenchUut6.windowSizeReached;
   TraceOut_error[430] := BenchUut6.error;
   TraceOut_status[430] := BenchUut6.status;
   BenchCalls := BenchCalls + 1;
 431:
   BenchUut6.cyclicExecution := FALSE;
   BenchUut6.trigger := FALSE;
   BenchUut6.value := LREAL#94.0;
   BenchUut6.windowSize := INT#100;
   BenchUut6.reset := FALSE;
   TraceIn_cyclicExecution[431] := BenchUut6.cyclicExecution;
   TraceIn_trigger[431] := BenchUut6.trigger;
   TraceIn_value[431] := BenchUut6.value;
   TraceIn_windowSize[431] := BenchUut6.windowSize;
   TraceIn_reset[431] := BenchUut6.reset;
   BenchUut6();
   TraceOut_average[431] := BenchUut6.average;
   TraceOut_windowSizeReached[431] := BenchUut6.windowSizeReached;
   TraceOut_error[431] := BenchUut6.error;
   TraceOut_status[431] := BenchUut6.status;
   BenchCalls := BenchCalls + 1;
 432:
   BenchUut6.cyclicExecution := FALSE;
   BenchUut6.trigger := TRUE;
   BenchUut6.value := LREAL#95.0;
   BenchUut6.windowSize := INT#100;
   BenchUut6.reset := FALSE;
   TraceIn_cyclicExecution[432] := BenchUut6.cyclicExecution;
   TraceIn_trigger[432] := BenchUut6.trigger;
   TraceIn_value[432] := BenchUut6.value;
   TraceIn_windowSize[432] := BenchUut6.windowSize;
   TraceIn_reset[432] := BenchUut6.reset;
   BenchUut6();
   TraceOut_average[432] := BenchUut6.average;
   TraceOut_windowSizeReached[432] := BenchUut6.windowSizeReached;
   TraceOut_error[432] := BenchUut6.error;
   TraceOut_status[432] := BenchUut6.status;
   BenchCalls := BenchCalls + 1;
 433:
   BenchUut6.cyclicExecution := FALSE;
   BenchUut6.trigger := FALSE;
   BenchUut6.value := LREAL#95.0;
   BenchUut6.windowSize := INT#100;
   BenchUut6.reset := FALSE;
   TraceIn_cyclicExecution[433] := BenchUut6.cyclicExecution;
   TraceIn_trigger[433] := BenchUut6.trigger;
   TraceIn_value[433] := BenchUut6.value;
   TraceIn_windowSize[433] := BenchUut6.windowSize;
   TraceIn_reset[433] := BenchUut6.reset;
   BenchUut6();
   TraceOut_average[433] := BenchUut6.average;
   TraceOut_windowSizeReached[433] := BenchUut6.windowSizeReached;
   TraceOut_error[433] := BenchUut6.error;
   TraceOut_status[433] := BenchUut6.status;
   BenchCalls := BenchCalls + 1;
 434:
   BenchUut6.cyclicExecution := FALSE;
   BenchUut6.trigger := TRUE;
   BenchUut6.value := LREAL#96.0;
   BenchUut6.windowSize := INT#100;
   BenchUut6.reset := FALSE;
   TraceIn_cyclicExecution[434] := BenchUut6.cyclicExecution;
   TraceIn_trigger[434] := BenchUut6.trigger;
   TraceIn_value[434] := BenchUut6.value;
   TraceIn_windowSize[434] := BenchUut6.windowSize;
   TraceIn_reset[434] := BenchUut6.reset;
   BenchUut6();
   TraceOut_average[434] := BenchUut6.average;
   TraceOut_windowSizeReached[434] := BenchUut6.windowSizeReached;
   TraceOut_error[434] := BenchUut6.error;
   TraceOut_status[434] := BenchUut6.status;
   BenchCalls := BenchCalls + 1;
 435:
   BenchUut6.cyclicExecution := FALSE;
   BenchUut6.trigger := FALSE;
   BenchUut6.value := LREAL#96.0;
   BenchUut6.windowSize := INT#100;
   BenchUut6.reset := FALSE;
   TraceIn_cyclicExecution[435] := BenchUut6.cyclicExecution;
   TraceIn_trigger[435] := BenchUut6.trigger;
   TraceIn_value[435] := BenchUut6.value;
   TraceIn_windowSize[435] := BenchUut6.windowSize;
   TraceIn_reset[435] := BenchUut6.reset;
   BenchUut6();
   TraceOut_average[435] := BenchUut6.average;
   TraceOut_windowSizeReached[435] := BenchUut6.windowSizeReached;
   TraceOut_error[435] := BenchUut6.error;
   TraceOut_status[435] := BenchUut6.status;
   BenchCalls := BenchCalls + 1;
 436:
   BenchUut6.cyclicExecution := FALSE;
   BenchUut6.trigger := TRUE;
   BenchUut6.value := LREAL#97.0;
   BenchUut6.windowSize := INT#100;
   BenchUut6.reset := FALSE;
   TraceIn_cyclicExecution[436] := BenchUut6.cyclicExecution;
   TraceIn_trigger[436] := BenchUut6.trigger;
   TraceIn_value[436] := BenchUut6.value;
   TraceIn_windowSize[436] := BenchUut6.windowSize;
   TraceIn_reset[436] := BenchUut6.reset;
   BenchUut6();
   TraceOut_average[436] := BenchUut6.average;
   TraceOut_windowSizeReached[436] := BenchUut6.windowSizeReached;
   TraceOut_error[436] := BenchUut6.error;
   TraceOut_status[436] := BenchUut6.status;
   BenchCalls := BenchCalls + 1;
 437:
   BenchUut6.cyclicExecution := FALSE;
   BenchUut6.trigger := FALSE;
   BenchUut6.value := LREAL#97.0;
   BenchUut6.windowSize := INT#100;
   BenchUut6.reset := FALSE;
   TraceIn_cyclicExecution[437] := BenchUut6.cyclicExecution;
   TraceIn_trigger[437] := BenchUut6.trigger;
   TraceIn_value[437] := BenchUut6.value;
   TraceIn_windowSize[437] := BenchUut6.windowSize;
   TraceIn_reset[437] := BenchUut6.reset;
   BenchUut6();
   TraceOut_average[437] := BenchUut6.average;
   TraceOut_windowSizeReached[437] := BenchUut6.windowSizeReached;
   TraceOut_error[437] := BenchUut6.error;
   TraceOut_status[437] := BenchUut6.status;
   BenchCalls := BenchCalls + 1;
 438:
   BenchUut6.cyclicExecution := FALSE;
   BenchUut6.trigger := TRUE;
   BenchUut6.value := LREAL#98.0;
   BenchUut6.windowSize := INT#100;
   BenchUut6.reset := FALSE;
   TraceIn_cyclicExecution[438] := BenchUut6.cyclicExecution;
   TraceIn_trigger[438] := BenchUut6.trigger;
   TraceIn_value[438] := BenchUut6.value;
   TraceIn_windowSize[438] := BenchUut6.windowSize;
   TraceIn_reset[438] := BenchUut6.reset;
   BenchUut6();
   TraceOut_average[438] := BenchUut6.average;
   TraceOut_windowSizeReached[438] := BenchUut6.windowSizeReached;
   TraceOut_error[438] := BenchUut6.error;
   TraceOut_status[438] := BenchUut6.status;
   BenchCalls := BenchCalls + 1;
 439:
   BenchUut6.cyclicExecution := FALSE;
   BenchUut6.trigger := FALSE;
   BenchUut6.value := LREAL#98.0;
   BenchUut6.windowSize := INT#100;
   BenchUut6.reset := FALSE;
   TraceIn_cyclicExecution[439] := BenchUut6.cyclicExecution;
   TraceIn_trigger[439] := BenchUut6.trigger;
   TraceIn_value[439] := BenchUut6.value;
   TraceIn_windowSize[439] := BenchUut6.windowSize;
   TraceIn_reset[439] := BenchUut6.reset;
   BenchUut6();
   TraceOut_average[439] := BenchUut6.average;
   TraceOut_windowSizeReached[439] := BenchUut6.windowSizeReached;
   TraceOut_error[439] := BenchUut6.error;
   TraceOut_status[439] := BenchUut6.status;
   BenchCalls := BenchCalls + 1;
 440:
   BenchUut6.cyclicExecution := FALSE;
   BenchUut6.trigger := TRUE;
   BenchUut6.value := LREAL#99.0;
   BenchUut6.windowSize := INT#100;
   BenchUut6.reset := FALSE;
   TraceIn_cyclicExecution[440] := BenchUut6.cyclicExecution;
   TraceIn_trigger[440] := BenchUut6.trigger;
   TraceIn_value[440] := BenchUut6.value;
   TraceIn_windowSize[440] := BenchUut6.windowSize;
   TraceIn_reset[440] := BenchUut6.reset;
   BenchUut6();
   TraceOut_average[440] := BenchUut6.average;
   TraceOut_windowSizeReached[440] := BenchUut6.windowSizeReached;
   TraceOut_error[440] := BenchUut6.error;
   TraceOut_status[440] := BenchUut6.status;
   BenchCalls := BenchCalls + 1;
 441:
   BenchUut6.cyclicExecution := FALSE;
   BenchUut6.trigger := FALSE;
   BenchUut6.value := LREAL#99.0;
   BenchUut6.windowSize := INT#100;
   BenchUut6.reset := FALSE;
   TraceIn_cyclicExecution[441] := BenchUut6.cyclicExecution;
   TraceIn_trigger[441] := BenchUut6.trigger;
   TraceIn_value[441] := BenchUut6.value;
   TraceIn_windowSize[441] := BenchUut6.windowSize;
   TraceIn_reset[441] := BenchUut6.reset;
   BenchUut6();
   TraceOut_average[441] := BenchUut6.average;
   TraceOut_windowSizeReached[441] := BenchUut6.windowSizeReached;
   TraceOut_error[441] := BenchUut6.error;
   TraceOut_status[441] := BenchUut6.status;
   BenchCalls := BenchCalls + 1;
 442:
   BenchUut6.cyclicExecution := FALSE;
   BenchUut6.trigger := TRUE;
   BenchUut6.value := LREAL#100.0;
   BenchUut6.windowSize := INT#100;
   BenchUut6.reset := FALSE;
   TraceIn_cyclicExecution[442] := BenchUut6.cyclicExecution;
   TraceIn_trigger[442] := BenchUut6.trigger;
   TraceIn_value[442] := BenchUut6.value;
   TraceIn_windowSize[442] := BenchUut6.windowSize;
   TraceIn_reset[442] := BenchUut6.reset;
   BenchUut6();
   TraceOut_average[442] := BenchUut6.average;
   TraceOut_windowSizeReached[442] := BenchUut6.windowSizeReached;
   TraceOut_error[442] := BenchUut6.error;
   TraceOut_status[442] := BenchUut6.status;
   BenchCalls := BenchCalls + 1;
 443:
   BenchUut6.cyclicExecution := FALSE;
   BenchUut6.trigger := FALSE;
   BenchUut6.value := LREAL#100.0;
   BenchUut6.windowSize := INT#100;
   BenchUut6.reset := FALSE;
   TraceIn_cyclicExecution[443] := BenchUut6.cyclicExecution;
   TraceIn_trigger[443] := BenchUut6.trigger;
   TraceIn_value[443] := BenchUut6.value;
   TraceIn_windowSize[443] := BenchUut6.windowSize;
   TraceIn_reset[443] := BenchUut6.reset;
   BenchUut6();
   TraceOut_average[443] := BenchUut6.average;
   TraceOut_windowSizeReached[443] := BenchUut6.windowSizeReached;
   TraceOut_error[443] := BenchUut6.error;
   TraceOut_status[443] := BenchUut6.status;
   BenchCalls := BenchCalls + 1;
 444:
   BenchUut6.cyclicExecution := FALSE;
   BenchUut6.trigger := TRUE;
   BenchUut6.value := LREAL#101.0;
   BenchUut6.windowSize := INT#100;
   BenchUut6.reset := FALSE;
   TraceIn_cyclicExecution[444] := BenchUut6.cyclicExecution;
   TraceIn_trigger[444] := BenchUut6.trigger;
   TraceIn_value[444] := BenchUut6.value;
   TraceIn_windowSize[444] := BenchUut6.windowSize;
   TraceIn_reset[444] := BenchUut6.reset;
   BenchUut6();
   TraceOut_average[444] := BenchUut6.average;
   TraceOut_windowSizeReached[444] := BenchUut6.windowSizeReached;
   TraceOut_error[444] := BenchUut6.error;
   TraceOut_status[444] := BenchUut6.status;
   BenchCalls := BenchCalls + 1;
 445:
   BenchUut6.cyclicExecution := FALSE;
   BenchUut6.trigger := FALSE;
   BenchUut6.value := LREAL#101.0;
   BenchUut6.windowSize := INT#100;
   BenchUut6.reset := FALSE;
   TraceIn_cyclicExecution[445] := BenchUut6.cyclicExecution;
   TraceIn_trigger[445] := BenchUut6.trigger;
   TraceIn_value[445] := BenchUut6.value;
   TraceIn_windowSize[445] := BenchUut6.windowSize;
   TraceIn_reset[445] := BenchUut6.reset;
   BenchUut6();
   TraceOut_average[445] := BenchUut6.average;
   TraceOut_windowSizeReached[445] := BenchUut6.windowSizeReached;
   TraceOut_error[445] := BenchUut6.error;
   TraceOut_status[445] := BenchUut6.status;
   BenchCalls := BenchCalls + 1;
 446:
   BenchUut6.cyclicExecution := FALSE;
   BenchUut6.trigger := TRUE;
   BenchUut6.value := LREAL#102.0;
   BenchUut6.windowSize := INT#100;
   BenchUut6.reset := FALSE;
   TraceIn_cyclicExecution[446] := BenchUut6.cyclicExecution;
   TraceIn_trigger[446] := BenchUut6.trigger;
   TraceIn_value[446] := BenchUut6.value;
   TraceIn_windowSize[446] := BenchUut6.windowSize;
   TraceIn_reset[446] := BenchUut6.reset;
   BenchUut6();
   TraceOut_average[446] := BenchUut6.average;
   TraceOut_windowSizeReached[446] := BenchUut6.windowSizeReached;
   TraceOut_error[446] := BenchUut6.error;
   TraceOut_status[446] := BenchUut6.status;
   BenchCalls := BenchCalls + 1;
 447:
   BenchUut6.cyclicExecution := FALSE;
   BenchUut6.trigger := FALSE;
   BenchUut6.value := LREAL#102.0;
   BenchUut6.windowSize := INT#100;
   BenchUut6.reset := FALSE;
   TraceIn_cyclicExecution[447] := BenchUut6.cyclicExecution;
   TraceIn_trigger[447] := BenchUut6.trigger;
   TraceIn_value[447] := BenchUut6.value;
   TraceIn_windowSize[447] := BenchUut6.windowSize;
   TraceIn_reset[447] := BenchUut6.reset;
   BenchUut6();
   TraceOut_average[447] := BenchUut6.average;
   TraceOut_windowSizeReached[447] := BenchUut6.windowSizeReached;
   TraceOut_error[447] := BenchUut6.error;
   TraceOut_status[447] := BenchUut6.status;
   BenchCalls := BenchCalls + 1;
 448:
   BenchUut6.cyclicExecution := FALSE;
   BenchUut6.trigger := TRUE;
   BenchUut6.value := LREAL#103.0;
   BenchUut6.windowSize := INT#100;
   BenchUut6.reset := FALSE;
   TraceIn_cyclicExecution[448] := BenchUut6.cyclicExecution;
   TraceIn_trigger[448] := BenchUut6.trigger;
   TraceIn_value[448] := BenchUut6.value;
   TraceIn_windowSize[448] := BenchUut6.windowSize;
   TraceIn_reset[448] := BenchUut6.reset;
   BenchUut6();
   TraceOut_average[448] := BenchUut6.average;
   TraceOut_windowSizeReached[448] := BenchUut6.windowSizeReached;
   TraceOut_error[448] := BenchUut6.error;
   TraceOut_status[448] := BenchUut6.status;
   BenchCalls := BenchCalls + 1;
 449:
   BenchUut6.cyclicExecution := FALSE;
   BenchUut6.trigger := FALSE;
   BenchUut6.value := LREAL#103.0;
   BenchUut6.windowSize := INT#100;
   BenchUut6.reset := FALSE;
   TraceIn_cyclicExecution[449] := BenchUut6.cyclicExecution;
   TraceIn_trigger[449] := BenchUut6.trigger;
   TraceIn_value[449] := BenchUut6.value;
   TraceIn_windowSize[449] := BenchUut6.windowSize;
   TraceIn_reset[449] := BenchUut6.reset;
   BenchUut6();
   TraceOut_average[449] := BenchUut6.average;
   TraceOut_windowSizeReached[449] := BenchUut6.windowSizeReached;
   TraceOut_error[449] := BenchUut6.error;
   TraceOut_status[449] := BenchUut6.status;
   BenchCalls := BenchCalls + 1;
 450:
   BenchUut6.cyclicExecution := FALSE;
   BenchUut6.trigger := TRUE;
   BenchUut6.value := LREAL#104.0;
   BenchUut6.windowSize := INT#100;
   BenchUut6.reset := FALSE;
   TraceIn_cyclicExecution[450] := BenchUut6.cyclicExecution;
   TraceIn_trigger[450] := BenchUut6.trigger;
   TraceIn_value[450] := BenchUut6.value;
   TraceIn_windowSize[450] := BenchUut6.windowSize;
   TraceIn_reset[450] := BenchUut6.reset;
   BenchUut6();
   TraceOut_average[450] := BenchUut6.average;
   TraceOut_windowSizeReached[450] := BenchUut6.windowSizeReached;
   TraceOut_error[450] := BenchUut6.error;
   TraceOut_status[450] := BenchUut6.status;
   BenchCalls := BenchCalls + 1;
 451:
   BenchUut6.cyclicExecution := FALSE;
   BenchUut6.trigger := FALSE;
   BenchUut6.value := LREAL#104.0;
   BenchUut6.windowSize := INT#2;
   BenchUut6.reset := FALSE;
   TraceIn_cyclicExecution[451] := BenchUut6.cyclicExecution;
   TraceIn_trigger[451] := BenchUut6.trigger;
   TraceIn_value[451] := BenchUut6.value;
   TraceIn_windowSize[451] := BenchUut6.windowSize;
   TraceIn_reset[451] := BenchUut6.reset;
   BenchUut6();
   TraceOut_average[451] := BenchUut6.average;
   TraceOut_windowSizeReached[451] := BenchUut6.windowSizeReached;
   TraceOut_error[451] := BenchUut6.error;
   TraceOut_status[451] := BenchUut6.status;
   BenchCalls := BenchCalls + 1;
 452:
   BenchUut6.cyclicExecution := FALSE;
   BenchUut6.trigger := TRUE;
   BenchUut6.value := LREAL#5.0;
   BenchUut6.windowSize := INT#2;
   BenchUut6.reset := FALSE;
   TraceIn_cyclicExecution[452] := BenchUut6.cyclicExecution;
   TraceIn_trigger[452] := BenchUut6.trigger;
   TraceIn_value[452] := BenchUut6.value;
   TraceIn_windowSize[452] := BenchUut6.windowSize;
   TraceIn_reset[452] := BenchUut6.reset;
   BenchUut6();
   TraceOut_average[452] := BenchUut6.average;
   TraceOut_windowSizeReached[452] := BenchUut6.windowSizeReached;
   TraceOut_error[452] := BenchUut6.error;
   TraceOut_status[452] := BenchUut6.status;
   BenchCalls := BenchCalls + 1;
 453:
   BenchUut6.cyclicExecution := FALSE;
   BenchUut6.trigger := FALSE;
   BenchUut6.value := LREAL#5.0;
   BenchUut6.windowSize := INT#100;
   BenchUut6.reset := FALSE;
   TraceIn_cyclicExecution[453] := BenchUut6.cyclicExecution;
   TraceIn_trigger[453] := BenchUut6.trigger;
   TraceIn_value[453] := BenchUut6.value;
   TraceIn_windowSize[453] := BenchUut6.windowSize;
   TraceIn_reset[453] := BenchUut6.reset;
   BenchUut6();
   TraceOut_average[453] := BenchUut6.average;
   TraceOut_windowSizeReached[453] := BenchUut6.windowSizeReached;
   TraceOut_error[453] := BenchUut6.error;
   TraceOut_status[453] := BenchUut6.status;
   BenchCalls := BenchCalls + 1;
 454:
   BenchUut6.cyclicExecution := FALSE;
   BenchUut6.trigger := TRUE;
   BenchUut6.value := LREAL#7.0;
   BenchUut6.windowSize := INT#100;
   BenchUut6.reset := FALSE;
   TraceIn_cyclicExecution[454] := BenchUut6.cyclicExecution;
   TraceIn_trigger[454] := BenchUut6.trigger;
   TraceIn_value[454] := BenchUut6.value;
   TraceIn_windowSize[454] := BenchUut6.windowSize;
   TraceIn_reset[454] := BenchUut6.reset;
   BenchUut6();
   TraceOut_average[454] := BenchUut6.average;
   TraceOut_windowSizeReached[454] := BenchUut6.windowSizeReached;
   TraceOut_error[454] := BenchUut6.error;
   TraceOut_status[454] := BenchUut6.status;
   BenchCalls := BenchCalls + 1;
 END_CASE;
 BenchStep := BenchStep + 1;
 IF BenchStep >= 455 THEN BenchDone := TRUE; END_IF;
END_IF;
END_PROGRAM
